(* IEC 61131-3 sources: STAR-PLC-Agent/results/raw/batch_fresh_20261114/PUB016/functional/attempt_0001, 1 file *)

(* ---- test_program.st ---- *)
PROGRAM PLC_PRG
VAR
 BenchStep : UDINT := 0;
 BenchCalls : UDINT := 0;
 BenchDone : BOOL := FALSE;
 BenchUut0 : FB_Task;
 BenchUut1 : FB_Task;
 BenchUut2 : FB_Task;
 BenchUut3 : FB_Task;
 BenchUut4 : FB_Task;
 BenchUut5 : FB_Task;
 BenchUut6 : FB_Task;
 BenchUut7 : FB_Task;
 TraceIn_processLength : ARRAY[0..159] OF USINT;
 TraceIn_sensor1 : ARRAY[0..159] OF BOOL;
 TraceIn_sensor2 : ARRAY[0..159] OF BOOL;
 TraceIn_sensor3 : ARRAY[0..159] OF BOOL;
 TraceIn_sensor4 : ARRAY[0..159] OF BOOL;
 TraceIn_sensor5 : ARRAY[0..159] OF BOOL;
 TraceIn_station1Start : ARRAY[0..159] OF BOOL;
 TraceIn_station2Complete : ARRAY[0..159] OF BOOL;
 TraceIn_station3Complete : ARRAY[0..159] OF BOOL;
 TraceIn_station4Complete : ARRAY[0..159] OF BOOL;
 TraceIn_processSequence_1 : ARRAY[0..159] OF USINT;
 TraceIn_processSequence_2 : ARRAY[0..159] OF USINT;
 TraceIn_processSequence_3 : ARRAY[0..159] OF USINT;
 TraceIn_processSequence_4 : ARRAY[0..159] OF USINT;
 TraceIn_processSequence_5 : ARRAY[0..159] OF USINT;
 TraceIn_processSequence_6 : ARRAY[0..159] OF USINT;
 TraceIn_processSequence_7 : ARRAY[0..159] OF USINT;
 TraceIn_processSequence_8 : ARRAY[0..159] OF USINT;
 TraceOut_conveyorLeft : ARRAY[0..159] OF BOOL;
 TraceOut_conveyorRight : ARRAY[0..159] OF BOOL;
END_VAR

IF NOT BenchDone THEN
 CASE BenchStep OF
 0:
   BenchUut0.processLength := USINT#3;
   BenchUut0.sensor1 := FALSE;
   BenchUut0.sensor2 := FALSE;
   BenchUut0.sensor3 := FALSE;
   BenchUut0.sensor4 := FALSE;
   BenchUut0.sensor5 := FALSE;
   BenchUut0.station1Start := FALSE;
   BenchUut0.station2Complete := FALSE;
   BenchUut0.station3Complete := FALSE;
   BenchUut0.station4Complete := FALSE;
   BenchUut0.processSequence[1] := USINT#4;
   BenchUut0.processSequence[2] := USINT#2;
   BenchUut0.processSequence[3] := USINT#5;
   BenchUut0.processSequence[4] := USINT#0;
   BenchUut0.processSequence[5] := USINT#0;
   BenchUut0.processSequence[6] := USINT#0;
   BenchUut0.processSequence[7] := USINT#0;
   BenchUut0.processSequence[8] := USINT#0;
   TraceIn_processLength[0] := BenchUut0.processLength;
   TraceIn_sensor1[0] := BenchUut0.sensor1;
   TraceIn_sensor2[0] := BenchUut0.sensor2;
   TraceIn_sensor3[0] := BenchUut0.sensor3;
   TraceIn_sensor4[0] := BenchUut0.sensor4;
   TraceIn_sensor5[0] := BenchUut0.sensor5;
   TraceIn_station1Start[0] := BenchUut0.station1Start;
   TraceIn_station2Complete[0] := BenchUut0.station2Complete;
   TraceIn_station3Complete[0] := BenchUut0.station3Complete;
   TraceIn_station4Complete[0] := BenchUut0.station4Complete;
   TraceIn_processSequence_1[0] := BenchUut0.processSequence[1];
   TraceIn_processSequence_2[0] := BenchUut0.processSequence[2];
   TraceIn_processSequence_3[0] := BenchUut0.processSequence[3];
   TraceIn_processSequence_4[0] := BenchUut0.processSequence[4];
   TraceIn_processSequence_5[0] := BenchUut0.processSequence[5];
   TraceIn_processSequence_6[0] := BenchUut0.processSequence[6];
   TraceIn_processSequence_7[0] := BenchUut0.processSequence[7];
   TraceIn_processSequence_8[0] := BenchUut0.processSequence[8];
   BenchUut0();
   TraceOut_conveyorLeft[0] := BenchUut0.conveyorLeft;
   TraceOut_conveyorRight[0] := BenchUut0.conveyorRight;
   BenchCalls := BenchCalls + 1;
 1:
   BenchUut0.processLength := USINT#3;
   BenchUut0.sensor1 := TRUE;
   BenchUut0.sensor2 := FALSE;
   BenchUut0.sensor3 := FALSE;
   BenchUut0.sensor4 := FALSE;
   BenchUut0.sensor5 := FALSE;
   BenchUut0.station1Start := TRUE;
   BenchUut0.station2Complete := FALSE;
   BenchUut0.station3Complete := FALSE;
   BenchUut0.station4Complete := FALSE;
   BenchUut0.processSequence[1] := USINT#4;
   BenchUut0.processSequence[2] := USINT#2;
   BenchUut0.processSequence[3] := USINT#5;
   BenchUut0.processSequence[4] := USINT#0;
   BenchUut0.processSequence[5] := USINT#0;
   BenchUut0.processSequence[6] := USINT#0;
   BenchUut0.processSequence[7] := USINT#0;
   BenchUut0.processSequence[8] := USINT#0;
   TraceIn_processLength[1] := BenchUut0.processLength;
   TraceIn_sensor1[1] := BenchUut0.sensor1;
   TraceIn_sensor2[1] := BenchUut0.sensor2;
   TraceIn_sensor3[1] := BenchUut0.sensor3;
   TraceIn_sensor4[1] := BenchUut0.sensor4;
   TraceIn_sensor5[1] := BenchUut0.sensor5;
   TraceIn_station1Start[1] := BenchUut0.station1Start;
   TraceIn_station2Complete[1] := BenchUut0.station2Complete;
   TraceIn_station3Complete[1] := BenchUut0.station3Complete;
   TraceIn_station4Complete[1] := BenchUut0.station4Complete;
   TraceIn_processSequence_1[1] := BenchUut0.processSequence[1];
   TraceIn_processSequence_2[1] := BenchUut0.processSequence[2];
   TraceIn_processSequence_3[1] := BenchUut0.processSequence[3];
   TraceIn_processSequence_4[1] := BenchUut0.processSequence[4];
   TraceIn_processSequence_5[1] := BenchUut0.processSequence[5];
   TraceIn_processSequence_6[1] := BenchUut0.processSequence[6];
   TraceIn_processSequence_7[1] := BenchUut0.processSequence[7];
   TraceIn_processSequence_8[1] := BenchUut0.processSequence[8];
   BenchUut0();
   TraceOut_conveyorLeft[1] := BenchUut0.conveyorLeft;
   TraceOut_conveyorRight[1] := BenchUut0.conveyorRight;
   BenchCalls := BenchCalls + 1;
 2:
   BenchUut0.processLength := USINT#3;
   BenchUut0.sensor1 := FALSE;
   BenchUut0.sensor2 := FALSE;
   BenchUut0.sensor3 := FALSE;
   BenchUut0.sensor4 := TRUE;
   BenchUut0.sensor5 := FALSE;
   BenchUut0.station1Start := FALSE;
   BenchUut0.station2Complete := FALSE;
   BenchUut0.station3Complete := FALSE;
   BenchUut0.station4Complete := FALSE;
   BenchUut0.processSequence[1] := USINT#4;
   BenchUut0.processSequence[2] := USINT#2;
   BenchUut0.processSequence[3] := USINT#5;
   BenchUut0.processSequence[4] := USINT#0;
   BenchUut0.processSequence[5] := USINT#0;
   BenchUut0.processSequence[6] := USINT#0;
   BenchUut0.processSequence[7] := USINT#0;
   BenchUut0.processSequence[8] := USINT#0;
   TraceIn_processLength[2] := BenchUut0.processLength;
   TraceIn_sensor1[2] := BenchUut0.sensor1;
   TraceIn_sensor2[2] := BenchUut0.sensor2;
   TraceIn_sensor3[2] := BenchUut0.sensor3;
   TraceIn_sensor4[2] := BenchUut0.sensor4;
   TraceIn_sensor5[2] := BenchUut0.sensor5;
   TraceIn_station1Start[2] := BenchUut0.station1Start;
   TraceIn_station2Complete[2] := BenchUut0.station2Complete;
   TraceIn_station3Complete[2] := BenchUut0.station3Complete;
   TraceIn_station4Complete[2] := BenchUut0.station4Complete;
   TraceIn_processSequence_1[2] := BenchUut0.processSequence[1];
   TraceIn_processSequence_2[2] := BenchUut0.processSequence[2];
   TraceIn_processSequence_3[2] := BenchUut0.processSequence[3];
   TraceIn_processSequence_4[2] := BenchUut0.processSequence[4];
   TraceIn_processSequence_5[2] := BenchUut0.processSequence[5];
   TraceIn_processSequence_6[2] := BenchUut0.processSequence[6];
   TraceIn_processSequence_7[2] := BenchUut0.processSequence[7];
   TraceIn_processSequence_8[2] := BenchUut0.processSequence[8];
   BenchUut0();
   TraceOut_conveyorLeft[2] := BenchUut0.conveyorLeft;
   TraceOut_conveyorRight[2] := BenchUut0.conveyorRight;
   BenchCalls := BenchCalls + 1;
 3:
   BenchUut0.processLength := USINT#3;
   BenchUut0.sensor1 := FALSE;
   BenchUut0.sensor2 := FALSE;
   BenchUut0.sensor3 := FALSE;
   BenchUut0.sensor4 := TRUE;
   BenchUut0.sensor5 := FALSE;
   BenchUut0.station1Start := FALSE;
   BenchUut0.station2Complete := FALSE;
   BenchUut0.station3Complete := TRUE;
   BenchUut0.station4Complete := FALSE;
   BenchUut0.processSequence[1] := USINT#4;
   BenchUut0.processSequence[2] := USINT#2;
   BenchUut0.processSequence[3] := USINT#5;
   BenchUut0.processSequence[4] := USINT#0;
   BenchUut0.processSequence[5] := USINT#0;
   BenchUut0.processSequence[6] := USINT#0;
   BenchUut0.processSequence[7] := USINT#0;
   BenchUut0.processSequence[8] := USINT#0;
   TraceIn_processLength[3] := BenchUut0.processLength;
   TraceIn_sensor1[3] := BenchUut0.sensor1;
   TraceIn_sensor2[3] := BenchUut0.sensor2;
   TraceIn_sensor3[3] := BenchUut0.sensor3;
   TraceIn_sensor4[3] := BenchUut0.sensor4;
   TraceIn_sensor5[3] := BenchUut0.sensor5;
   TraceIn_station1Start[3] := BenchUut0.station1Start;
   TraceIn_station2Complete[3] := BenchUut0.station2Complete;
   TraceIn_station3Complete[3] := BenchUut0.station3Complete;
   TraceIn_station4Complete[3] := BenchUut0.station4Complete;
   TraceIn_processSequence_1[3] := BenchUut0.processSequence[1];
   TraceIn_processSequence_2[3] := BenchUut0.processSequence[2];
   TraceIn_processSequence_3[3] := BenchUut0.processSequence[3];
   TraceIn_processSequence_4[3] := BenchUut0.processSequence[4];
   TraceIn_processSequence_5[3] := BenchUut0.processSequence[5];
   TraceIn_processSequence_6[3] := BenchUut0.processSequence[6];
   TraceIn_processSequence_7[3] := BenchUut0.processSequence[7];
   TraceIn_processSequence_8[3] := BenchUut0.processSequence[8];
   BenchUut0();
   TraceOut_conveyorLeft[3] := BenchUut0.conveyorLeft;
   TraceOut_conveyorRight[3] := BenchUut0.conveyorRight;
   BenchCalls := BenchCalls + 1;
 4:
   BenchUut0.processLength := USINT#3;
   BenchUut0.sensor1 := FALSE;
   BenchUut0.sensor2 := FALSE;
   BenchUut0.sensor3 := FALSE;
   BenchUut0.sensor4 := TRUE;
   BenchUut0.sensor5 := FALSE;
   BenchUut0.station1Start := FALSE;
   BenchUut0.station2Complete := FALSE;
   BenchUut0.station3Complete := FALSE;
   BenchUut0.station4Complete := TRUE;
   BenchUut0.processSequence[1] := USINT#4;
   BenchUut0.processSequence[2] := USINT#2;
   BenchUut0.processSequence[3] := USINT#5;
   BenchUut0.processSequence[4] := USINT#0;
   BenchUut0.processSequence[5] := USINT#0;
   BenchUut0.processSequence[6] := USINT#0;
   BenchUut0.processSequence[7] := USINT#0;
   BenchUut0.processSequence[8] := USINT#0;
   TraceIn_processLength[4] := BenchUut0.processLength;
   TraceIn_sensor1[4] := BenchUut0.sensor1;
   TraceIn_sensor2[4] := BenchUut0.sensor2;
   TraceIn_sensor3[4] := BenchUut0.sensor3;
   TraceIn_sensor4[4] := BenchUut0.sensor4;
   TraceIn_sensor5[4] := BenchUut0.sensor5;
   TraceIn_station1Start[4] := BenchUut0.station1Start;
   TraceIn_station2Complete[4] := BenchUut0.station2Complete;
   TraceIn_station3Complete[4] := BenchUut0.station3Complete;
   TraceIn_station4Complete[4] := BenchUut0.station4Complete;
   TraceIn_processSequence_1[4] := BenchUut0.processSequence[1];
   TraceIn_processSequence_2[4] := BenchUut0.processSequence[2];
   TraceIn_processSequence_3[4] := BenchUut0.processSequence[3];
   TraceIn_processSequence_4[4] := BenchUut0.processSequence[4];
   TraceIn_processSequence_5[4] := BenchUut0.processSequence[5];
   TraceIn_processSequence_6[4] := BenchUut0.processSequence[6];
   TraceIn_processSequence_7[4] := BenchUut0.processSequence[7];
   TraceIn_processSequence_8[4] := BenchUut0.processSequence[8];
   BenchUut0();
   TraceOut_conveyorLeft[4] := BenchUut0.conveyorLeft;
   TraceOut_conveyorRight[4] := BenchUut0.conveyorRight;
   BenchCalls := BenchCalls + 1;
 5:
   BenchUut0.processLength := USINT#3;
   BenchUut0.sensor1 := FALSE;
   BenchUut0.sensor2 := TRUE;
   BenchUut0.sensor3 := FALSE;
   BenchUut0.sensor4 := FALSE;
   BenchUut0.sensor5 := FALSE;
   BenchUut0.station1Start := FALSE;
   BenchUut0.station2Complete := FALSE;
   BenchUut0.station3Complete := FALSE;
   BenchUut0.station4Complete := FALSE;
   BenchUut0.processSequence[1] := USINT#4;
   BenchUut0.processSequence[2] := USINT#2;
   BenchUut0.processSequence[3] := USINT#5;
   BenchUut0.processSequence[4] := USINT#0;
   BenchUut0.processSequence[5] := USINT#0;
   BenchUut0.processSequence[6] := USINT#0;
   BenchUut0.processSequence[7] := USINT#0;
   BenchUut0.processSequence[8] := USINT#0;
   TraceIn_processLength[5] := BenchUut0.processLength;
   TraceIn_sensor1[5] := BenchUut0.sensor1;
   TraceIn_sensor2[5] := BenchUut0.sensor2;
   TraceIn_sensor3[5] := BenchUut0.sensor3;
   TraceIn_sensor4[5] := BenchUut0.sensor4;
   TraceIn_sensor5[5] := BenchUut0.sensor5;
   TraceIn_station1Start[5] := BenchUut0.station1Start;
   TraceIn_station2Complete[5] := BenchUut0.station2Complete;
   TraceIn_station3Complete[5] := BenchUut0.station3Complete;
   TraceIn_station4Complete[5] := BenchUut0.station4Complete;
   TraceIn_processSequence_1[5] := BenchUut0.processSequence[1];
   TraceIn_processSequence_2[5] := BenchUut0.processSequence[2];
   TraceIn_processSequence_3[5] := BenchUut0.processSequence[3];
   TraceIn_processSequence_4[5] := BenchUut0.processSequence[4];
   TraceIn_processSequence_5[5] := BenchUut0.processSequence[5];
   TraceIn_processSequence_6[5] := BenchUut0.processSequence[6];
   TraceIn_processSequence_7[5] := BenchUut0.processSequence[7];
   TraceIn_processSequence_8[5] := BenchUut0.processSequence[8];
   BenchUut0();
   TraceOut_conveyorLeft[5] := BenchUut0.conveyorLeft;
   TraceOut_conveyorRight[5] := BenchUut0.conveyorRight;
   BenchCalls := BenchCalls + 1;
 6:
   BenchUut0.processLength := USINT#3;
   BenchUut0.sensor1 := FALSE;
   BenchUut0.sensor2 := TRUE;
   BenchUut0.sensor3 := FALSE;
   BenchUut0.sensor4 := FALSE;
   BenchUut0.sensor5 := FALSE;
   BenchUut0.station1Start := FALSE;
   BenchUut0.station2Complete := TRUE;
   BenchUut0.station3Complete := FALSE;
   BenchUut0.station4Complete := FALSE;
   BenchUut0.processSequence[1] := USINT#4;
   BenchUut0.processSequence[2] := USINT#2;
   BenchUut0.processSequence[3] := USINT#5;
   BenchUut0.processSequence[4] := USINT#0;
   BenchUut0.processSequence[5] := USINT#0;
   BenchUut0.processSequence[6] := USINT#0;
   BenchUut0.processSequence[7] := USINT#0;
   BenchUut0.processSequence[8] := USINT#0;
   TraceIn_processLength[6] := BenchUut0.processLength;
   TraceIn_sensor1[6] := BenchUut0.sensor1;
   TraceIn_sensor2[6] := BenchUut0.sensor2;
   TraceIn_sensor3[6] := BenchUut0.sensor3;
   TraceIn_sensor4[6] := BenchUut0.sensor4;
   TraceIn_sensor5[6] := BenchUut0.sensor5;
   TraceIn_station1Start[6] := BenchUut0.station1Start;
   TraceIn_station2Complete[6] := BenchUut0.station2Complete;
   TraceIn_station3Complete[6] := BenchUut0.station3Complete;
   TraceIn_station4Complete[6] := BenchUut0.station4Complete;
   TraceIn_processSequence_1[6] := BenchUut0.processSequence[1];
   TraceIn_processSequence_2[6] := BenchUut0.processSequence[2];
   TraceIn_processSequence_3[6] := BenchUut0.processSequence[3];
   TraceIn_processSequence_4[6] := BenchUut0.processSequence[4];
   TraceIn_processSequence_5[6] := BenchUut0.processSequence[5];
   TraceIn_processSequence_6[6] := BenchUut0.processSequence[6];
   TraceIn_processSequence_7[6] := BenchUut0.processSequence[7];
   TraceIn_processSequence_8[6] := BenchUut0.processSequence[8];
   BenchUut0();
   TraceOut_conveyorLeft[6] := BenchUut0.conveyorLeft;
   TraceOut_conveyorRight[6] := BenchUut0.conveyorRight;
   BenchCalls := BenchCalls + 1;
 7:
   BenchUut0.processLength := USINT#3;
   BenchUut0.sensor1 := FALSE;
   BenchUut0.sensor2 := FALSE;
   BenchUut0.sensor3 := FALSE;
   BenchUut0.sensor4 := FALSE;
   BenchUut0.sensor5 := TRUE;
   BenchUut0.station1Start := FALSE;
   BenchUut0.station2Complete := FALSE;
   BenchUut0.station3Complete := FALSE;
   BenchUut0.station4Complete := FALSE;
   BenchUut0.processSequence[1] := USINT#4;
   BenchUut0.processSequence[2] := USINT#2;
   BenchUut0.processSequence[3] := USINT#5;
   BenchUut0.processSequence[4] := USINT#0;
   BenchUut0.processSequence[5] := USINT#0;
   BenchUut0.processSequence[6] := USINT#0;
   BenchUut0.processSequence[7] := USINT#0;
   BenchUut0.processSequence[8] := USINT#0;
   TraceIn_processLength[7] := BenchUut0.processLength;
   TraceIn_sensor1[7] := BenchUut0.sensor1;
   TraceIn_sensor2[7] := BenchUut0.sensor2;
   TraceIn_sensor3[7] := BenchUut0.sensor3;
   TraceIn_sensor4[7] := BenchUut0.sensor4;
   TraceIn_sensor5[7] := BenchUut0.sensor5;
   TraceIn_station1Start[7] := BenchUut0.station1Start;
   TraceIn_station2Complete[7] := BenchUut0.station2Complete;
   TraceIn_station3Complete[7] := BenchUut0.station3Complete;
   TraceIn_station4Complete[7] := BenchUut0.station4Complete;
   TraceIn_processSequence_1[7] := BenchUut0.processSequence[1];
   TraceIn_processSequence_2[7] := BenchUut0.processSequence[2];
   TraceIn_processSequence_3[7] := BenchUut0.processSequence[3];
   TraceIn_processSequence_4[7] := BenchUut0.processSequence[4];
   TraceIn_processSequence_5[7] := BenchUut0.processSequence[5];
   TraceIn_processSequence_6[7] := BenchUut0.processSequence[6];
   TraceIn_processSequence_7[7] := BenchUut0.processSequence[7];
   TraceIn_processSequence_8[7] := BenchUut0.processSequence[8];
   BenchUut0();
   TraceOut_conveyorLeft[7] := BenchUut0.conveyorLeft;
   TraceOut_conveyorRight[7] := BenchUut0.conveyorRight;
   BenchCalls := BenchCalls + 1;
 8:
   BenchUut1.processLength := USINT#1;
   BenchUut1.sensor1 := FALSE;
   BenchUut1.sensor2 := FALSE;
   BenchUut1.sensor3 := FALSE;
   BenchUut1.sensor4 := FALSE;
   BenchUut1.sensor5 := FALSE;
   BenchUut1.station1Start := FALSE;
   BenchUut1.station2Complete := FALSE;
   BenchUut1.station3Complete := FALSE;
   BenchUut1.station4Complete := FALSE;
   BenchUut1.processSequence[1] := USINT#5;
   BenchUut1.processSequence[2] := USINT#0;
   BenchUut1.processSequence[3] := USINT#0;
   BenchUut1.processSequence[4] := USINT#0;
   BenchUut1.processSequence[5] := USINT#0;
   BenchUut1.processSequence[6] := USINT#0;
   BenchUut1.processSequence[7] := USINT#0;
   BenchUut1.processSequence[8] := USINT#0;
   TraceIn_processLength[8] := BenchUut1.processLength;
   TraceIn_sensor1[8] := BenchUut1.sensor1;
   TraceIn_sensor2[8] := BenchUut1.sensor2;
   TraceIn_sensor3[8] := BenchUut1.sensor3;
   TraceIn_sensor4[8] := BenchUut1.sensor4;
   TraceIn_sensor5[8] := BenchUut1.sensor5;
   TraceIn_station1Start[8] := BenchUut1.station1Start;
   TraceIn_station2Complete[8] := BenchUut1.station2Complete;
   TraceIn_station3Complete[8] := BenchUut1.station3Complete;
   TraceIn_station4Complete[8] := BenchUut1.station4Complete;
   TraceIn_processSequence_1[8] := BenchUut1.processSequence[1];
   TraceIn_processSequence_2[8] := BenchUut1.processSequence[2];
   TraceIn_processSequence_3[8] := BenchUut1.processSequence[3];
   TraceIn_processSequence_4[8] := BenchUut1.processSequence[4];
   TraceIn_processSequence_5[8] := BenchUut1.processSequence[5];
   TraceIn_processSequence_6[8] := BenchUut1.processSequence[6];
   TraceIn_processSequence_7[8] := BenchUut1.processSequence[7];
   TraceIn_processSequence_8[8] := BenchUut1.processSequence[8];
   BenchUut1();
   TraceOut_conveyorLeft[8] := BenchUut1.conveyorLeft;
   TraceOut_conveyorRight[8] := BenchUut1.conveyorRight;
   BenchCalls := BenchCalls + 1;
 9:
   BenchUut1.processLength := USINT#1;
   BenchUut1.sensor1 := TRUE;
   BenchUut1.sensor2 := FALSE;
   BenchUut1.sensor3 := FALSE;
   BenchUut1.sensor4 := FALSE;
   BenchUut1.sensor5 := FALSE;
   BenchUut1.station1Start := TRUE;
   BenchUut1.station2Complete := FALSE;
   BenchUut1.station3Complete := FALSE;
   BenchUut1.station4Complete := FALSE;
   BenchUut1.processSequence[1] := USINT#5;
   BenchUut1.processSequence[2] := USINT#0;
   BenchUut1.processSequence[3] := USINT#0;
   BenchUut1.processSequence[4] := USINT#0;
   BenchUut1.processSequence[5] := USINT#0;
   BenchUut1.processSequence[6] := USINT#0;
   BenchUut1.processSequence[7] := USINT#0;
   BenchUut1.processSequence[8] := USINT#0;
   TraceIn_processLength[9] := BenchUut1.processLength;
   TraceIn_sensor1[9] := BenchUut1.sensor1;
   TraceIn_sensor2[9] := BenchUut1.sensor2;
   TraceIn_sensor3[9] := BenchUut1.sensor3;
   TraceIn_sensor4[9] := BenchUut1.sensor4;
   TraceIn_sensor5[9] := BenchUut1.sensor5;
   TraceIn_station1Start[9] := BenchUut1.station1Start;
   TraceIn_station2Complete[9] := BenchUut1.station2Complete;
   TraceIn_station3Complete[9] := BenchUut1.station3Complete;
   TraceIn_station4Complete[9] := BenchUut1.station4Complete;
   TraceIn_processSequence_1[9] := BenchUut1.processSequence[1];
   TraceIn_processSequence_2[9] := BenchUut1.processSequence[2];
   TraceIn_processSequence_3[9] := BenchUut1.processSequence[3];
   TraceIn_processSequence_4[9] := BenchUut1.processSequence[4];
   TraceIn_processSequence_5[9] := BenchUut1.processSequence[5];
   TraceIn_processSequence_6[9] := BenchUut1.processSequence[6];
   TraceIn_processSequence_7[9] := BenchUut1.processSequence[7];
   TraceIn_processSequence_8[9] := BenchUut1.processSequence[8];
   BenchUut1();
   TraceOut_conveyorLeft[9] := BenchUut1.conveyorLeft;
   TraceOut_conveyorRight[9] := BenchUut1.conveyorRight;
   BenchCalls := BenchCalls + 1;
 10:
   BenchUut1.processLength := USINT#1;
   BenchUut1.sensor1 := FALSE;
   BenchUut1.sensor2 := FALSE;
   BenchUut1.sensor3 := FALSE;
   BenchUut1.sensor4 := FALSE;
   BenchUut1.sensor5 := TRUE;
   BenchUut1.station1Start := FALSE;
   BenchUut1.station2Complete := FALSE;
   BenchUut1.station3Complete := FALSE;
   BenchUut1.station4Complete := FALSE;
   BenchUut1.processSequence[1] := USINT#5;
   BenchUut1.processSequence[2] := USINT#0;
   BenchUut1.processSequence[3] := USINT#0;
   BenchUut1.processSequence[4] := USINT#0;
   BenchUut1.processSequence[5] := USINT#0;
   BenchUut1.processSequence[6] := USINT#0;
   BenchUut1.processSequence[7] := USINT#0;
   BenchUut1.processSequence[8] := USINT#0;
   TraceIn_processLength[10] := BenchUut1.processLength;
   TraceIn_sensor1[10] := BenchUut1.sensor1;
   TraceIn_sensor2[10] := BenchUut1.sensor2;
   TraceIn_sensor3[10] := BenchUut1.sensor3;
   TraceIn_sensor4[10] := BenchUut1.sensor4;
   TraceIn_sensor5[10] := BenchUut1.sensor5;
   TraceIn_station1Start[10] := BenchUut1.station1Start;
   TraceIn_station2Complete[10] := BenchUut1.station2Complete;
   TraceIn_station3Complete[10] := BenchUut1.station3Complete;
   TraceIn_station4Complete[10] := BenchUut1.station4Complete;
   TraceIn_processSequence_1[10] := BenchUut1.processSequence[1];
   TraceIn_processSequence_2[10] := BenchUut1.processSequence[2];
   TraceIn_processSequence_3[10] := BenchUut1.processSequence[3];
   TraceIn_processSequence_4[10] := BenchUut1.processSequence[4];
   TraceIn_processSequence_5[10] := BenchUut1.processSequence[5];
   TraceIn_processSequence_6[10] := BenchUut1.processSequence[6];
   TraceIn_processSequence_7[10] := BenchUut1.processSequence[7];
   TraceIn_processSequence_8[10] := BenchUut1.processSequence[8];
   BenchUut1();
   TraceOut_conveyorLeft[10] := BenchUut1.conveyorLeft;
   TraceOut_conveyorRight[10] := BenchUut1.conveyorRight;
   BenchCalls := BenchCalls + 1;
 11:
   BenchUut2.processLength := USINT#3;
   BenchUut2.sensor1 := FALSE;
   BenchUut2.sensor2 := FALSE;
   BenchUut2.sensor3 := FALSE;
   BenchUut2.sensor4 := FALSE;
   BenchUut2.sensor5 := FALSE;
   BenchUut2.station1Start := FALSE;
   BenchUut2.station2Complete := FALSE;
   BenchUut2.station3Complete := FALSE;
   BenchUut2.station4Complete := FALSE;
   BenchUut2.processSequence[1] := USINT#2;
   BenchUut2.processSequence[2] := USINT#2;
   BenchUut2.processSequence[3] := USINT#5;
   BenchUut2.processSequence[4] := USINT#0;
   BenchUut2.processSequence[5] := USINT#0;
   BenchUut2.processSequence[6] := USINT#0;
   BenchUut2.processSequence[7] := USINT#0;
   BenchUut2.processSequence[8] := USINT#0;
   TraceIn_processLength[11] := BenchUut2.processLength;
   TraceIn_sensor1[11] := BenchUut2.sensor1;
   TraceIn_sensor2[11] := BenchUut2.sensor2;
   TraceIn_sensor3[11] := BenchUut2.sensor3;
   TraceIn_sensor4[11] := BenchUut2.sensor4;
   TraceIn_sensor5[11] := BenchUut2.sensor5;
   TraceIn_station1Start[11] := BenchUut2.station1Start;
   TraceIn_station2Complete[11] := BenchUut2.station2Complete;
   TraceIn_station3Complete[11] := BenchUut2.station3Complete;
   TraceIn_station4Complete[11] := BenchUut2.station4Complete;
   TraceIn_processSequence_1[11] := BenchUut2.processSequence[1];
   TraceIn_processSequence_2[11] := BenchUut2.processSequence[2];
   TraceIn_processSequence_3[11] := BenchUut2.processSequence[3];
   TraceIn_processSequence_4[11] := BenchUut2.processSequence[4];
   TraceIn_processSequence_5[11] := BenchUut2.processSequence[5];
   TraceIn_processSequence_6[11] := BenchUut2.processSequence[6];
   TraceIn_processSequence_7[11] := BenchUut2.processSequence[7];
   TraceIn_processSequence_8[11] := BenchUut2.processSequence[8];
   BenchUut2();
   TraceOut_conveyorLeft[11] := BenchUut2.conveyorLeft;
   TraceOut_conveyorRight[11] := BenchUut2.conveyorRight;
   BenchCalls := BenchCalls + 1;
 12:
   BenchUut2.processLength := USINT#3;
   BenchUut2.sensor1 := TRUE;
   BenchUut2.sensor2 := FALSE;
   BenchUut2.sensor3 := FALSE;
   BenchUut2.sensor4 := FALSE;
   BenchUut2.sensor5 := FALSE;
   BenchUut2.station1Start := TRUE;
   BenchUut2.station2Complete := FALSE;
   BenchUut2.station3Complete := FALSE;
   BenchUut2.station4Complete := FALSE;
   BenchUut2.processSequence[1] := USINT#2;
   BenchUut2.processSequence[2] := USINT#2;
   BenchUut2.processSequence[3] := USINT#5;
   BenchUut2.processSequence[4] := USINT#0;
   BenchUut2.processSequence[5] := USINT#0;
   BenchUut2.processSequence[6] := USINT#0;
   BenchUut2.processSequence[7] := USINT#0;
   BenchUut2.processSequence[8] := USINT#0;
   TraceIn_processLength[12] := BenchUut2.processLength;
   TraceIn_sensor1[12] := BenchUut2.sensor1;
   TraceIn_sensor2[12] := BenchUut2.sensor2;
   TraceIn_sensor3[12] := BenchUut2.sensor3;
   TraceIn_sensor4[12] := BenchUut2.sensor4;
   TraceIn_sensor5[12] := BenchUut2.sensor5;
   TraceIn_station1Start[12] := BenchUut2.station1Start;
   TraceIn_station2Complete[12] := BenchUut2.station2Complete;
   TraceIn_station3Complete[12] := BenchUut2.station3Complete;
   TraceIn_station4Complete[12] := BenchUut2.station4Complete;
   TraceIn_processSequence_1[12] := BenchUut2.processSequence[1];
   TraceIn_processSequence_2[12] := BenchUut2.processSequence[2];
   TraceIn_processSequence_3[12] := BenchUut2.processSequence[3];
   TraceIn_processSequence_4[12] := BenchUut2.processSequence[4];
   TraceIn_processSequence_5[12] := BenchUut2.processSequence[5];
   TraceIn_processSequence_6[12] := BenchUut2.processSequence[6];
   TraceIn_processSequence_7[12] := BenchUut2.processSequence[7];
   TraceIn_processSequence_8[12] := BenchUut2.processSequence[8];
   BenchUut2();
   TraceOut_conveyorLeft[12] := BenchUut2.conveyorLeft;
   TraceOut_conveyorRight[12] := BenchUut2.conveyorRight;
   BenchCalls := BenchCalls + 1;
 13:
   BenchUut2.processLength := USINT#3;
   BenchUut2.sensor1 := FALSE;
   BenchUut2.sensor2 := TRUE;
   BenchUut2.sensor3 := FALSE;
   BenchUut2.sensor4 := FALSE;
   BenchUut2.sensor5 := FALSE;
   BenchUut2.station1Start := FALSE;
   BenchUut2.station2Complete := FALSE;
   BenchUut2.station3Complete := FALSE;
   BenchUut2.station4Complete := FALSE;
   BenchUut2.processSequence[1] := USINT#2;
   BenchUut2.processSequence[2] := USINT#2;
   BenchUut2.processSequence[3] := USINT#5;
   BenchUut2.processSequence[4] := USINT#0;
   BenchUut2.processSequence[5] := USINT#0;
   BenchUut2.processSequence[6] := USINT#0;
   BenchUut2.processSequence[7] := USINT#0;
   BenchUut2.processSequence[8] := USINT#0;
   TraceIn_processLength[13] := BenchUut2.processLength;
   TraceIn_sensor1[13] := BenchUut2.sensor1;
   TraceIn_sensor2[13] := BenchUut2.sensor2;
   TraceIn_sensor3[13] := BenchUut2.sensor3;
   TraceIn_sensor4[13] := BenchUut2.sensor4;
   TraceIn_sensor5[13] := BenchUut2.sensor5;
   TraceIn_station1Start[13] := BenchUut2.station1Start;
   TraceIn_station2Complete[13] := BenchUut2.station2Complete;
   TraceIn_station3Complete[13] := BenchUut2.station3Complete;
   TraceIn_station4Complete[13] := BenchUut2.station4Complete;
   TraceIn_processSequence_1[13] := BenchUut2.processSequence[1];
   TraceIn_processSequence_2[13] := BenchUut2.processSequence[2];
   TraceIn_processSequence_3[13] := BenchUut2.processSequence[3];
   TraceIn_processSequence_4[13] := BenchUut2.processSequence[4];
   TraceIn_processSequence_5[13] := BenchUut2.processSequence[5];
   TraceIn_processSequence_6[13] := BenchUut2.processSequence[6];
   TraceIn_processSequence_7[13] := BenchUut2.processSequence[7];
   TraceIn_processSequence_8[13] := BenchUut2.processSequence[8];
   BenchUut2();
   TraceOut_conveyorLeft[13] := BenchUut2.conveyorLeft;
   TraceOut_conveyorRight[13] := BenchUut2.conveyorRight;
   BenchCalls := BenchCalls + 1;
 14:
   BenchUut2.processLength := USINT#3;
   BenchUut2.sensor1 := FALSE;
   BenchUut2.sensor2 := TRUE;
   BenchUut2.sensor3 := FALSE;
   BenchUut2.sensor4 := FALSE;
   BenchUut2.sensor5 := FALSE;
   BenchUut2.station1Start := FALSE;
   BenchUut2.station2Complete := TRUE;
   BenchUut2.station3Complete := FALSE;
   BenchUut2.station4Complete := FALSE;
   BenchUut2.processSequence[1] := USINT#2;
   BenchUut2.processSequence[2] := USINT#2;
   BenchUut2.processSequence[3] := USINT#5;
   BenchUut2.processSequence[4] := USINT#0;
   BenchUut2.processSequence[5] := USINT#0;
   BenchUut2.processSequence[6] := USINT#0;
   BenchUut2.processSequence[7] := USINT#0;
   BenchUut2.processSequence[8] := USINT#0;
   TraceIn_processLength[14] := BenchUut2.processLength;
   TraceIn_sensor1[14] := BenchUut2.sensor1;
   TraceIn_sensor2[14] := BenchUut2.sensor2;
   TraceIn_sensor3[14] := BenchUut2.sensor3;
   TraceIn_sensor4[14] := BenchUut2.sensor4;
   TraceIn_sensor5[14] := BenchUut2.sensor5;
   TraceIn_station1Start[14] := BenchUut2.station1Start;
   TraceIn_station2Complete[14] := BenchUut2.station2Complete;
   TraceIn_station3Complete[14] := BenchUut2.station3Complete;
   TraceIn_station4Complete[14] := BenchUut2.station4Complete;
   TraceIn_processSequence_1[14] := BenchUut2.processSequence[1];
   TraceIn_processSequence_2[14] := BenchUut2.processSequence[2];
   TraceIn_processSequence_3[14] := BenchUut2.processSequence[3];
   TraceIn_processSequence_4[14] := BenchUut2.processSequence[4];
   TraceIn_processSequence_5[14] := BenchUut2.processSequence[5];
   TraceIn_processSequence_6[14] := BenchUut2.processSequence[6];
   TraceIn_processSequence_7[14] := BenchUut2.processSequence[7];
   TraceIn_processSequence_8[14] := BenchUut2.processSequence[8];
   BenchUut2();
   TraceOut_conveyorLeft[14] := BenchUut2.conveyorLeft;
   TraceOut_conveyorRight[14] := BenchUut2.conveyorRight;
   BenchCalls := BenchCalls + 1;
 15:
   BenchUut2.processLength := USINT#3;
   BenchUut2.sensor1 := FALSE;
   BenchUut2.sensor2 := TRUE;
   BenchUut2.sensor3 := FALSE;
   BenchUut2.sensor4 := FALSE;
   BenchUut2.sensor5 := FALSE;
   BenchUut2.station1Start := FALSE;
   BenchUut2.station2Complete := TRUE;
   BenchUut2.station3Complete := FALSE;
   BenchUut2.station4Complete := FALSE;
   BenchUut2.processSequence[1] := USINT#2;
   BenchUut2.processSequence[2] := USINT#2;
   BenchUut2.processSequence[3] := USINT#5;
   BenchUut2.processSequence[4] := USINT#0;
   BenchUut2.processSequence[5] := USINT#0;
   BenchUut2.processSequence[6] := USINT#0;
   BenchUut2.processSequence[7] := USINT#0;
   BenchUut2.processSequence[8] := USINT#0;
   TraceIn_processLength[15] := BenchUut2.processLength;
   TraceIn_sensor1[15] := BenchUut2.sensor1;
   TraceIn_sensor2[15] := BenchUut2.sensor2;
   TraceIn_sensor3[15] := BenchUut2.sensor3;
   TraceIn_sensor4[15] := BenchUut2.sensor4;
   TraceIn_sensor5[15] := BenchUut2.sensor5;
   TraceIn_station1Start[15] := BenchUut2.station1Start;
   TraceIn_station2Complete[15] := BenchUut2.station2Complete;
   TraceIn_station3Complete[15] := BenchUut2.station3Complete;
   TraceIn_station4Complete[15] := BenchUut2.station4Complete;
   TraceIn_processSequence_1[15] := BenchUut2.processSequence[1];
   TraceIn_processSequence_2[15] := BenchUut2.processSequence[2];
   TraceIn_processSequence_3[15] := BenchUut2.processSequence[3];
   TraceIn_processSequence_4[15] := BenchUut2.processSequence[4];
   TraceIn_processSequence_5[15] := BenchUut2.processSequence[5];
   TraceIn_processSequence_6[15] := BenchUut2.processSequence[6];
   TraceIn_processSequence_7[15] := BenchUut2.processSequence[7];
   TraceIn_processSequence_8[15] := BenchUut2.processSequence[8];
   BenchUut2();
   TraceOut_conveyorLeft[15] := BenchUut2.conveyorLeft;
   TraceOut_conveyorRight[15] := BenchUut2.conveyorRight;
   BenchCalls := BenchCalls + 1;
 16:
   BenchUut2.processLength := USINT#3;
   BenchUut2.sensor1 := FALSE;
   BenchUut2.sensor2 := TRUE;
   BenchUut2.sensor3 := FALSE;
   BenchUut2.sensor4 := FALSE;
   BenchUut2.sensor5 := FALSE;
   BenchUut2.station1Start := FALSE;
   BenchUut2.station2Complete := FALSE;
   BenchUut2.station3Complete := FALSE;
   BenchUut2.station4Complete := FALSE;
   BenchUut2.processSequence[1] := USINT#2;
   BenchUut2.processSequence[2] := USINT#2;
   BenchUut2.processSequence[3] := USINT#5;
   BenchUut2.processSequence[4] := USINT#0;
   BenchUut2.processSequence[5] := USINT#0;
   BenchUut2.processSequence[6] := USINT#0;
   BenchUut2.processSequence[7] := USINT#0;
   BenchUut2.processSequence[8] := USINT#0;
   TraceIn_processLength[16] := BenchUut2.processLength;
   TraceIn_sensor1[16] := BenchUut2.sensor1;
   TraceIn_sensor2[16] := BenchUut2.sensor2;
   TraceIn_sensor3[16] := BenchUut2.sensor3;
   TraceIn_sensor4[16] := BenchUut2.sensor4;
   TraceIn_sensor5[16] := BenchUut2.sensor5;
   TraceIn_station1Start[16] := BenchUut2.station1Start;
   TraceIn_station2Complete[16] := BenchUut2.station2Complete;
   TraceIn_station3Complete[16] := BenchUut2.station3Complete;
   TraceIn_station4Complete[16] := BenchUut2.station4Complete;
   TraceIn_processSequence_1[16] := BenchUut2.processSequence[1];
   TraceIn_processSequence_2[16] := BenchUut2.processSequence[2];
   TraceIn_processSequence_3[16] := BenchUut2.processSequence[3];
   TraceIn_processSequence_4[16] := BenchUut2.processSequence[4];
   TraceIn_processSequence_5[16] := BenchUut2.processSequence[5];
   TraceIn_processSequence_6[16] := BenchUut2.processSequence[6];
   TraceIn_processSequence_7[16] := BenchUut2.processSequence[7];
   TraceIn_processSequence_8[16] := BenchUut2.processSequence[8];
   BenchUut2();
   TraceOut_conveyorLeft[16] := BenchUut2.conveyorLeft;
   TraceOut_conveyorRight[16] := BenchUut2.conveyorRight;
   BenchCalls := BenchCalls + 1;
 17:
   BenchUut2.processLength := USINT#3;
   BenchUut2.sensor1 := FALSE;
   BenchUut2.sensor2 := TRUE;
   BenchUut2.sensor3 := FALSE;
   BenchUut2.sensor4 := FALSE;
   BenchUut2.sensor5 := FALSE;
   BenchUut2.station1Start := FALSE;
   BenchUut2.station2Complete := TRUE;
   BenchUut2.station3Complete := FALSE;
   BenchUut2.station4Complete := FALSE;
   BenchUut2.processSequence[1] := USINT#2;
   BenchUut2.processSequence[2] := USINT#2;
   BenchUut2.processSequence[3] := USINT#5;
   BenchUut2.processSequence[4] := USINT#0;
   BenchUut2.processSequence[5] := USINT#0;
   BenchUut2.processSequence[6] := USINT#0;
   BenchUut2.processSequence[7] := USINT#0;
   BenchUut2.processSequence[8] := USINT#0;
   TraceIn_processLength[17] := BenchUut2.processLength;
   TraceIn_sensor1[17] := BenchUut2.sensor1;
   TraceIn_sensor2[17] := BenchUut2.sensor2;
   TraceIn_sensor3[17] := BenchUut2.sensor3;
   TraceIn_sensor4[17] := BenchUut2.sensor4;
   TraceIn_sensor5[17] := BenchUut2.sensor5;
   TraceIn_station1Start[17] := BenchUut2.station1Start;
   TraceIn_station2Complete[17] := BenchUut2.station2Complete;
   TraceIn_station3Complete[17] := BenchUut2.station3Complete;
   TraceIn_station4Complete[17] := BenchUut2.station4Complete;
   TraceIn_processSequence_1[17] := BenchUut2.processSequence[1];
   TraceIn_processSequence_2[17] := BenchUut2.processSequence[2];
   TraceIn_processSequence_3[17] := BenchUut2.processSequence[3];
   TraceIn_processSequence_4[17] := BenchUut2.processSequence[4];
   TraceIn_processSequence_5[17] := BenchUut2.processSequence[5];
   TraceIn_processSequence_6[17] := BenchUut2.processSequence[6];
   TraceIn_processSequence_7[17] := BenchUut2.processSequence[7];
   TraceIn_processSequence_8[17] := BenchUut2.processSequence[8];
   BenchUut2();
   TraceOut_conveyorLeft[17] := BenchUut2.conveyorLeft;
   TraceOut_conveyorRight[17] := BenchUut2.conveyorRight;
   BenchCalls := BenchCalls + 1;
 18:
   BenchUut3.processLength := USINT#3;
   BenchUut3.sensor1 := TRUE;
   BenchUut3.sensor2 := FALSE;
   BenchUut3.sensor3 := FALSE;
   BenchUut3.sensor4 := FALSE;
   BenchUut3.sensor5 := FALSE;
   BenchUut3.station1Start := TRUE;
   BenchUut3.station2Complete := FALSE;
   BenchUut3.station3Complete := FALSE;
   BenchUut3.station4Complete := FALSE;
   BenchUut3.processSequence[1] := USINT#2;
   BenchUut3.processSequence[2] := USINT#2;
   BenchUut3.processSequence[3] := USINT#5;
   BenchUut3.processSequence[4] := USINT#0;
   BenchUut3.processSequence[5] := USINT#0;
   BenchUut3.processSequence[6] := USINT#0;
   BenchUut3.processSequence[7] := USINT#0;
   BenchUut3.processSequence[8] := USINT#0;
   TraceIn_processLength[18] := BenchUut3.processLength;
   TraceIn_sensor1[18] := BenchUut3.sensor1;
   TraceIn_sensor2[18] := BenchUut3.sensor2;
   TraceIn_sensor3[18] := BenchUut3.sensor3;
   TraceIn_sensor4[18] := BenchUut3.sensor4;
   TraceIn_sensor5[18] := BenchUut3.sensor5;
   TraceIn_station1Start[18] := BenchUut3.station1Start;
   TraceIn_station2Complete[18] := BenchUut3.station2Complete;
   TraceIn_station3Complete[18] := BenchUut3.station3Complete;
   TraceIn_station4Complete[18] := BenchUut3.station4Complete;
   TraceIn_processSequence_1[18] := BenchUut3.processSequence[1];
   TraceIn_processSequence_2[18] := BenchUut3.processSequence[2];
   TraceIn_processSequence_3[18] := BenchUut3.processSequence[3];
   TraceIn_processSequence_4[18] := BenchUut3.processSequence[4];
   TraceIn_processSequence_5[18] := BenchUut3.processSequence[5];
   TraceIn_processSequence_6[18] := BenchUut3.processSequence[6];
   TraceIn_processSequence_7[18] := BenchUut3.processSequence[7];
   TraceIn_processSequence_8[18] := BenchUut3.processSequence[8];
   BenchUut3();
   TraceOut_conveyorLeft[18] := BenchUut3.conveyorLeft;
   TraceOut_conveyorRight[18] := BenchUut3.conveyorRight;
   BenchCalls := BenchCalls + 1;
 19:
   BenchUut3.processLength := USINT#3;
   BenchUut3.sensor1 := FALSE;
   BenchUut3.sensor2 := TRUE;
   BenchUut3.sensor3 := FALSE;
   BenchUut3.sensor4 := FALSE;
   BenchUut3.sensor5 := FALSE;
   BenchUut3.station1Start := FALSE;
   BenchUut3.station2Complete := TRUE;
   BenchUut3.station3Complete := FALSE;
   BenchUut3.station4Complete := FALSE;
   BenchUut3.processSequence[1] := USINT#2;
   BenchUut3.processSequence[2] := USINT#2;
   BenchUut3.processSequence[3] := USINT#5;
   BenchUut3.processSequence[4] := USINT#0;
   BenchUut3.processSequence[5] := USINT#0;
   BenchUut3.processSequence[6] := USINT#0;
   BenchUut3.processSequence[7] := USINT#0;
   BenchUut3.processSequence[8] := USINT#0;
   TraceIn_processLength[19] := BenchUut3.processLength;
   TraceIn_sensor1[19] := BenchUut3.sensor1;
   TraceIn_sensor2[19] := BenchUut3.sensor2;
   TraceIn_sensor3[19] := BenchUut3.sensor3;
   TraceIn_sensor4[19] := BenchUut3.sensor4;
   TraceIn_sensor5[19] := BenchUut3.sensor5;
   TraceIn_station1Start[19] := BenchUut3.station1Start;
   TraceIn_station2Complete[19] := BenchUut3.station2Complete;
   TraceIn_station3Complete[19] := BenchUut3.station3Complete;
   TraceIn_station4Complete[19] := BenchUut3.station4Complete;
   TraceIn_processSequence_1[19] := BenchUut3.processSequence[1];
   TraceIn_processSequence_2[19] := BenchUut3.processSequence[2];
   TraceIn_processSequence_3[19] := BenchUut3.processSequence[3];
   TraceIn_processSequence_4[19] := BenchUut3.processSequence[4];
   TraceIn_processSequence_5[19] := BenchUut3.processSequence[5];
   TraceIn_processSequence_6[19] := BenchUut3.processSequence[6];
   TraceIn_processSequence_7[19] := BenchUut3.processSequence[7];
   TraceIn_processSequence_8[19] := BenchUut3.processSequence[8];
   BenchUut3();
   TraceOut_conveyorLeft[19] := BenchUut3.conveyorLeft;
   TraceOut_conveyorRight[19] := BenchUut3.conveyorRight;
   BenchCalls := BenchCalls + 1;
 20:
   BenchUut3.processLength := USINT#3;
   BenchUut3.sensor1 := FALSE;
   BenchUut3.sensor2 := TRUE;
   BenchUut3.sensor3 := FALSE;
   BenchUut3.sensor4 := FALSE;
   BenchUut3.sensor5 := FALSE;
   BenchUut3.station1Start := FALSE;
   BenchUut3.station2Complete := TRUE;
   BenchUut3.station3Complete := FALSE;
   BenchUut3.station4Complete := FALSE;
   BenchUut3.processSequence[1] := USINT#2;
   BenchUut3.processSequence[2] := USINT#2;
   BenchUut3.processSequence[3] := USINT#5;
   BenchUut3.processSequence[4] := USINT#0;
   BenchUut3.processSequence[5] := USINT#0;
   BenchUut3.processSequence[6] := USINT#0;
   BenchUut3.processSequence[7] := USINT#0;
   BenchUut3.processSequence[8] := USINT#0;
   TraceIn_processLength[20] := BenchUut3.processLength;
   TraceIn_sensor1[20] := BenchUut3.sensor1;
   TraceIn_sensor2[20] := BenchUut3.sensor2;
   TraceIn_sensor3[20] := BenchUut3.sensor3;
   TraceIn_sensor4[20] := BenchUut3.sensor4;
   TraceIn_sensor5[20] := BenchUut3.sensor5;
   TraceIn_station1Start[20] := BenchUut3.station1Start;
   TraceIn_station2Complete[20] := BenchUut3.station2Complete;
   TraceIn_station3Complete[20] := BenchUut3.station3Complete;
   TraceIn_station4Complete[20] := BenchUut3.station4Complete;
   TraceIn_processSequence_1[20] := BenchUut3.processSequence[1];
   TraceIn_processSequence_2[20] := BenchUut3.processSequence[2];
   TraceIn_processSequence_3[20] := BenchUut3.processSequence[3];
   TraceIn_processSequence_4[20] := BenchUut3.processSequence[4];
   TraceIn_processSequence_5[20] := BenchUut3.processSequence[5];
   TraceIn_processSequence_6[20] := BenchUut3.processSequence[6];
   TraceIn_processSequence_7[20] := BenchUut3.processSequence[7];
   TraceIn_processSequence_8[20] := BenchUut3.processSequence[8];
   BenchUut3();
   TraceOut_conveyorLeft[20] := BenchUut3.conveyorLeft;
   TraceOut_conveyorRight[20] := BenchUut3.conveyorRight;
   BenchCalls := BenchCalls + 1;
 21:
   BenchUut3.processLength := USINT#3;
   BenchUut3.sensor1 := FALSE;
   BenchUut3.sensor2 := TRUE;
   BenchUut3.sensor3 := FALSE;
   BenchUut3.sensor4 := FALSE;
   BenchUut3.sensor5 := FALSE;
   BenchUut3.station1Start := FALSE;
   BenchUut3.station2Complete := FALSE;
   BenchUut3.station3Complete := FALSE;
   BenchUut3.station4Complete := FALSE;
   BenchUut3.processSequence[1] := USINT#2;
   BenchUut3.processSequence[2] := USINT#2;
   BenchUut3.processSequence[3] := USINT#5;
   BenchUut3.processSequence[4] := USINT#0;
   BenchUut3.processSequence[5] := USINT#0;
   BenchUut3.processSequence[6] := USINT#0;
   BenchUut3.processSequence[7] := USINT#0;
   BenchUut3.processSequence[8] := USINT#0;
   TraceIn_processLength[21] := BenchUut3.processLength;
   TraceIn_sensor1[21] := BenchUut3.sensor1;
   TraceIn_sensor2[21] := BenchUut3.sensor2;
   TraceIn_sensor3[21] := BenchUut3.sensor3;
   TraceIn_sensor4[21] := BenchUut3.sensor4;
   TraceIn_sensor5[21] := BenchUut3.sensor5;
   TraceIn_station1Start[21] := BenchUut3.station1Start;
   TraceIn_station2Complete[21] := BenchUut3.station2Complete;
   TraceIn_station3Complete[21] := BenchUut3.station3Complete;
   TraceIn_station4Complete[21] := BenchUut3.station4Complete;
   TraceIn_processSequence_1[21] := BenchUut3.processSequence[1];
   TraceIn_processSequence_2[21] := BenchUut3.processSequence[2];
   TraceIn_processSequence_3[21] := BenchUut3.processSequence[3];
   TraceIn_processSequence_4[21] := BenchUut3.processSequence[4];
   TraceIn_processSequence_5[21] := BenchUut3.processSequence[5];
   TraceIn_processSequence_6[21] := BenchUut3.processSequence[6];
   TraceIn_processSequence_7[21] := BenchUut3.processSequence[7];
   TraceIn_processSequence_8[21] := BenchUut3.processSequence[8];
   BenchUut3();
   TraceOut_conveyorLeft[21] := BenchUut3.conveyorLeft;
   TraceOut_conveyorRight[21] := BenchUut3.conveyorRight;
   BenchCalls := BenchCalls + 1;
 22:
   BenchUut3.processLength := USINT#3;
   BenchUut3.sensor1 := FALSE;
   BenchUut3.sensor2 := TRUE;
   BenchUut3.sensor3 := FALSE;
   BenchUut3.sensor4 := FALSE;
   BenchUut3.sensor5 := FALSE;
   BenchUut3.station1Start := FALSE;
   BenchUut3.station2Complete := TRUE;
   BenchUut3.station3Complete := FALSE;
   BenchUut3.station4Complete := FALSE;
   BenchUut3.processSequence[1] := USINT#2;
   BenchUut3.processSequence[2] := USINT#2;
   BenchUut3.processSequence[3] := USINT#5;
   BenchUut3.processSequence[4] := USINT#0;
   BenchUut3.processSequence[5] := USINT#0;
   BenchUut3.processSequence[6] := USINT#0;
   BenchUut3.processSequence[7] := USINT#0;
   BenchUut3.processSequence[8] := USINT#0;
   TraceIn_processLength[22] := BenchUut3.processLength;
   TraceIn_sensor1[22] := BenchUut3.sensor1;
   TraceIn_sensor2[22] := BenchUut3.sensor2;
   TraceIn_sensor3[22] := BenchUut3.sensor3;
   TraceIn_sensor4[22] := BenchUut3.sensor4;
   TraceIn_sensor5[22] := BenchUut3.sensor5;
   TraceIn_station1Start[22] := BenchUut3.station1Start;
   TraceIn_station2Complete[22] := BenchUut3.station2Complete;
   TraceIn_station3Complete[22] := BenchUut3.station3Complete;
   TraceIn_station4Complete[22] := BenchUut3.station4Complete;
   TraceIn_processSequence_1[22] := BenchUut3.processSequence[1];
   TraceIn_processSequence_2[22] := BenchUut3.processSequence[2];
   TraceIn_processSequence_3[22] := BenchUut3.processSequence[3];
   TraceIn_processSequence_4[22] := BenchUut3.processSequence[4];
   TraceIn_processSequence_5[22] := BenchUut3.processSequence[5];
   TraceIn_processSequence_6[22] := BenchUut3.processSequence[6];
   TraceIn_processSequence_7[22] := BenchUut3.processSequence[7];
   TraceIn_processSequence_8[22] := BenchUut3.processSequence[8];
   BenchUut3();
   TraceOut_conveyorLeft[22] := BenchUut3.conveyorLeft;
   TraceOut_conveyorRight[22] := BenchUut3.conveyorRight;
   BenchCalls := BenchCalls + 1;
 23:
   BenchUut3.processLength := USINT#3;
   BenchUut3.sensor1 := FALSE;
   BenchUut3.sensor2 := TRUE;
   BenchUut3.sensor3 := FALSE;
   BenchUut3.sensor4 := FALSE;
   BenchUut3.sensor5 := FALSE;
   BenchUut3.station1Start := FALSE;
   BenchUut3.station2Complete := TRUE;
   BenchUut3.station3Complete := FALSE;
   BenchUut3.station4Complete := FALSE;
   BenchUut3.processSequence[1] := USINT#2;
   BenchUut3.processSequence[2] := USINT#2;
   BenchUut3.processSequence[3] := USINT#5;
   BenchUut3.processSequence[4] := USINT#0;
   BenchUut3.processSequence[5] := USINT#0;
   BenchUut3.processSequence[6] := USINT#0;
   BenchUut3.processSequence[7] := USINT#0;
   BenchUut3.processSequence[8] := USINT#0;
   TraceIn_processLength[23] := BenchUut3.processLength;
   TraceIn_sensor1[23] := BenchUut3.sensor1;
   TraceIn_sensor2[23] := BenchUut3.sensor2;
   TraceIn_sensor3[23] := BenchUut3.sensor3;
   TraceIn_sensor4[23] := BenchUut3.sensor4;
   TraceIn_sensor5[23] := BenchUut3.sensor5;
   TraceIn_station1Start[23] := BenchUut3.station1Start;
   TraceIn_station2Complete[23] := BenchUut3.station2Complete;
   TraceIn_station3Complete[23] := BenchUut3.station3Complete;
   TraceIn_station4Complete[23] := BenchUut3.station4Complete;
   TraceIn_processSequence_1[23] := BenchUut3.processSequence[1];
   TraceIn_processSequence_2[23] := BenchUut3.processSequence[2];
   TraceIn_processSequence_3[23] := BenchUut3.processSequence[3];
   TraceIn_processSequence_4[23] := BenchUut3.processSequence[4];
   TraceIn_processSequence_5[23] := BenchUut3.processSequence[5];
   TraceIn_processSequence_6[23] := BenchUut3.processSequence[6];
   TraceIn_processSequence_7[23] := BenchUut3.processSequence[7];
   TraceIn_processSequence_8[23] := BenchUut3.processSequence[8];
   BenchUut3();
   TraceOut_conveyorLeft[23] := BenchUut3.conveyorLeft;
   TraceOut_conveyorRight[23] := BenchUut3.conveyorRight;
   BenchCalls := BenchCalls + 1;
 24:
   BenchUut3.processLength := USINT#3;
   BenchUut3.sensor1 := FALSE;
   BenchUut3.sensor2 := TRUE;
   BenchUut3.sensor3 := FALSE;
   BenchUut3.sensor4 := FALSE;
   BenchUut3.sensor5 := FALSE;
   BenchUut3.station1Start := FALSE;
   BenchUut3.station2Complete := FALSE;
   BenchUut3.station3Complete := FALSE;
   BenchUut3.station4Complete := FALSE;
   BenchUut3.processSequence[1] := USINT#2;
   BenchUut3.processSequence[2] := USINT#2;
   BenchUut3.processSequence[3] := USINT#5;
   BenchUut3.processSequence[4] := USINT#0;
   BenchUut3.processSequence[5] := USINT#0;
   BenchUut3.processSequence[6] := USINT#0;
   BenchUut3.processSequence[7] := USINT#0;
   BenchUut3.processSequence[8] := USINT#0;
   TraceIn_processLength[24] := BenchUut3.processLength;
   TraceIn_sensor1[24] := BenchUut3.sensor1;
   TraceIn_sensor2[24] := BenchUut3.sensor2;
   TraceIn_sensor3[24] := BenchUut3.sensor3;
   TraceIn_sensor4[24] := BenchUut3.sensor4;
   TraceIn_sensor5[24] := BenchUut3.sensor5;
   TraceIn_station1Start[24] := BenchUut3.station1Start;
   TraceIn_station2Complete[24] := BenchUut3.station2Complete;
   TraceIn_station3Complete[24] := BenchUut3.station3Complete;
   TraceIn_station4Complete[24] := BenchUut3.station4Complete;
   TraceIn_processSequence_1[24] := BenchUut3.processSequence[1];
   TraceIn_processSequence_2[24] := BenchUut3.processSequence[2];
   TraceIn_processSequence_3[24] := BenchUut3.processSequence[3];
   TraceIn_processSequence_4[24] := BenchUut3.processSequence[4];
   TraceIn_processSequence_5[24] := BenchUut3.processSequence[5];
   TraceIn_processSequence_6[24] := BenchUut3.processSequence[6];
   TraceIn_processSequence_7[24] := BenchUut3.processSequence[7];
   TraceIn_processSequence_8[24] := BenchUut3.processSequence[8];
   BenchUut3();
   TraceOut_conveyorLeft[24] := BenchUut3.conveyorLeft;
   TraceOut_conveyorRight[24] := BenchUut3.conveyorRight;
   BenchCalls := BenchCalls + 1;
 25:
   BenchUut3.processLength := USINT#3;
   BenchUut3.sensor1 := FALSE;
   BenchUut3.sensor2 := TRUE;
   BenchUut3.sensor3 := FALSE;
   BenchUut3.sensor4 := FALSE;
   BenchUut3.sensor5 := FALSE;
   BenchUut3.station1Start := FALSE;
   BenchUut3.station2Complete := TRUE;
   BenchUut3.station3Complete := FALSE;
   BenchUut3.station4Complete := FALSE;
   BenchUut3.processSequence[1] := USINT#2;
   BenchUut3.processSequence[2] := USINT#2;
   BenchUut3.processSequence[3] := USINT#5;
   BenchUut3.processSequence[4] := USINT#0;
   BenchUut3.processSequence[5] := USINT#0;
   BenchUut3.processSequence[6] := USINT#0;
   BenchUut3.processSequence[7] := USINT#0;
   BenchUut3.processSequence[8] := USINT#0;
   TraceIn_processLength[25] := BenchUut3.processLength;
   TraceIn_sensor1[25] := BenchUut3.sensor1;
   TraceIn_sensor2[25] := BenchUut3.sensor2;
   TraceIn_sensor3[25] := BenchUut3.sensor3;
   TraceIn_sensor4[25] := BenchUut3.sensor4;
   TraceIn_sensor5[25] := BenchUut3.sensor5;
   TraceIn_station1Start[25] := BenchUut3.station1Start;
   TraceIn_station2Complete[25] := BenchUut3.station2Complete;
   TraceIn_station3Complete[25] := BenchUut3.station3Complete;
   TraceIn_station4Complete[25] := BenchUut3.station4Complete;
   TraceIn_processSequence_1[25] := BenchUut3.processSequence[1];
   TraceIn_processSequence_2[25] := BenchUut3.processSequence[2];
   TraceIn_processSequence_3[25] := BenchUut3.processSequence[3];
   TraceIn_processSequence_4[25] := BenchUut3.processSequence[4];
   TraceIn_processSequence_5[25] := BenchUut3.processSequence[5];
   TraceIn_processSequence_6[25] := BenchUut3.processSequence[6];
   TraceIn_processSequence_7[25] := BenchUut3.processSequence[7];
   TraceIn_processSequence_8[25] := BenchUut3.processSequence[8];
   BenchUut3();
   TraceOut_conveyorLeft[25] := BenchUut3.conveyorLeft;
   TraceOut_conveyorRight[25] := BenchUut3.conveyorRight;
   BenchCalls := BenchCalls + 1;
 26:
   BenchUut3.processLength := USINT#3;
   BenchUut3.sensor1 := FALSE;
   BenchUut3.sensor2 := FALSE;
   BenchUut3.sensor3 := FALSE;
   BenchUut3.sensor4 := FALSE;
   BenchUut3.sensor5 := TRUE;
   BenchUut3.station1Start := FALSE;
   BenchUut3.station2Complete := FALSE;
   BenchUut3.station3Complete := FALSE;
   BenchUut3.station4Complete := FALSE;
   BenchUut3.processSequence[1] := USINT#2;
   BenchUut3.processSequence[2] := USINT#2;
   BenchUut3.processSequence[3] := USINT#5;
   BenchUut3.processSequence[4] := USINT#0;
   BenchUut3.processSequence[5] := USINT#0;
   BenchUut3.processSequence[6] := USINT#0;
   BenchUut3.processSequence[7] := USINT#0;
   BenchUut3.processSequence[8] := USINT#0;
   TraceIn_processLength[26] := BenchUut3.processLength;
   TraceIn_sensor1[26] := BenchUut3.sensor1;
   TraceIn_sensor2[26] := BenchUut3.sensor2;
   TraceIn_sensor3[26] := BenchUut3.sensor3;
   TraceIn_sensor4[26] := BenchUut3.sensor4;
   TraceIn_sensor5[26] := BenchUut3.sensor5;
   TraceIn_station1Start[26] := BenchUut3.station1Start;
   TraceIn_station2Complete[26] := BenchUut3.station2Complete;
   TraceIn_station3Complete[26] := BenchUut3.station3Complete;
   TraceIn_station4Complete[26] := BenchUut3.station4Complete;
   TraceIn_processSequence_1[26] := BenchUut3.processSequence[1];
   TraceIn_processSequence_2[26] := BenchUut3.processSequence[2];
   TraceIn_processSequence_3[26] := BenchUut3.processSequence[3];
   TraceIn_processSequence_4[26] := BenchUut3.processSequence[4];
   TraceIn_processSequence_5[26] := BenchUut3.processSequence[5];
   TraceIn_processSequence_6[26] := BenchUut3.processSequence[6];
   TraceIn_processSequence_7[26] := BenchUut3.processSequence[7];
   TraceIn_processSequence_8[26] := BenchUut3.processSequence[8];
   BenchUut3();
   TraceOut_conveyorLeft[26] := BenchUut3.conveyorLeft;
   TraceOut_conveyorRight[26] := BenchUut3.conveyorRight;
   BenchCalls := BenchCalls + 1;
 27:
   BenchUut4.processLength := USINT#8;
   BenchUut4.sensor1 := FALSE;
   BenchUut4.sensor2 := FALSE;
   BenchUut4.sensor3 := FALSE;
   BenchUut4.sensor4 := FALSE;
   BenchUut4.sensor5 := FALSE;
   BenchUut4.station1Start := TRUE;
   BenchUut4.station2Complete := FALSE;
   BenchUut4.station3Complete := FALSE;
   BenchUut4.station4Complete := FALSE;
   BenchUut4.processSequence[1] := USINT#4;
   BenchUut4.processSequence[2] := USINT#3;
   BenchUut4.processSequence[3] := USINT#2;
   BenchUut4.processSequence[4] := USINT#4;
   BenchUut4.processSequence[5] := USINT#2;
   BenchUut4.processSequence[6] := USINT#3;
   BenchUut4.processSequence[7] := USINT#4;
   BenchUut4.processSequence[8] := USINT#5;
   TraceIn_processLength[27] := BenchUut4.processLength;
   TraceIn_sensor1[27] := BenchUut4.sensor1;
   TraceIn_sensor2[27] := BenchUut4.sensor2;
   TraceIn_sensor3[27] := BenchUut4.sensor3;
   TraceIn_sensor4[27] := BenchUut4.sensor4;
   TraceIn_sensor5[27] := BenchUut4.sensor5;
   TraceIn_station1Start[27] := BenchUut4.station1Start;
   TraceIn_station2Complete[27] := BenchUut4.station2Complete;
   TraceIn_station3Complete[27] := BenchUut4.station3Complete;
   TraceIn_station4Complete[27] := BenchUut4.station4Complete;
   TraceIn_processSequence_1[27] := BenchUut4.processSequence[1];
   TraceIn_processSequence_2[27] := BenchUut4.processSequence[2];
   TraceIn_processSequence_3[27] := BenchUut4.processSequence[3];
   TraceIn_processSequence_4[27] := BenchUut4.processSequence[4];
   TraceIn_processSequence_5[27] := BenchUut4.processSequence[5];
   TraceIn_processSequence_6[27] := BenchUut4.processSequence[6];
   TraceIn_processSequence_7[27] := BenchUut4.processSequence[7];
   TraceIn_processSequence_8[27] := BenchUut4.processSequence[8];
   BenchUut4();
   TraceOut_conveyorLeft[27] := BenchUut4.conveyorLeft;
   TraceOut_conveyorRight[27] := BenchUut4.conveyorRight;
   BenchCalls := BenchCalls + 1;
 28:
   BenchUut4.processLength := USINT#8;
   BenchUut4.sensor1 := TRUE;
   BenchUut4.sensor2 := FALSE;
   BenchUut4.sensor3 := FALSE;
   BenchUut4.sensor4 := FALSE;
   BenchUut4.sensor5 := FALSE;
   BenchUut4.station1Start := TRUE;
   BenchUut4.station2Complete := FALSE;
   BenchUut4.station3Complete := FALSE;
   BenchUut4.station4Complete := FALSE;
   BenchUut4.processSequence[1] := USINT#4;
   BenchUut4.processSequence[2] := USINT#3;
   BenchUut4.processSequence[3] := USINT#2;
   BenchUut4.processSequence[4] := USINT#4;
   BenchUut4.processSequence[5] := USINT#2;
   BenchUut4.processSequence[6] := USINT#3;
   BenchUut4.processSequence[7] := USINT#4;
   BenchUut4.processSequence[8] := USINT#5;
   TraceIn_processLength[28] := BenchUut4.processLength;
   TraceIn_sensor1[28] := BenchUut4.sensor1;
   TraceIn_sensor2[28] := BenchUut4.sensor2;
   TraceIn_sensor3[28] := BenchUut4.sensor3;
   TraceIn_sensor4[28] := BenchUut4.sensor4;
   TraceIn_sensor5[28] := BenchUut4.sensor5;
   TraceIn_station1Start[28] := BenchUut4.station1Start;
   TraceIn_station2Complete[28] := BenchUut4.station2Complete;
   TraceIn_station3Complete[28] := BenchUut4.station3Complete;
   TraceIn_station4Complete[28] := BenchUut4.station4Complete;
   TraceIn_processSequence_1[28] := BenchUut4.processSequence[1];
   TraceIn_processSequence_2[28] := BenchUut4.processSequence[2];
   TraceIn_processSequence_3[28] := BenchUut4.processSequence[3];
   TraceIn_processSequence_4[28] := BenchUut4.processSequence[4];
   TraceIn_processSequence_5[28] := BenchUut4.processSequence[5];
   TraceIn_processSequence_6[28] := BenchUut4.processSequence[6];
   TraceIn_processSequence_7[28] := BenchUut4.processSequence[7];
   TraceIn_processSequence_8[28] := BenchUut4.processSequence[8];
   BenchUut4();
   TraceOut_conveyorLeft[28] := BenchUut4.conveyorLeft;
   TraceOut_conveyorRight[28] := BenchUut4.conveyorRight;
   BenchCalls := BenchCalls + 1;
 29:
   BenchUut4.processLength := USINT#8;
   BenchUut4.sensor1 := FALSE;
   BenchUut4.sensor2 := TRUE;
   BenchUut4.sensor3 := FALSE;
   BenchUut4.sensor4 := FALSE;
   BenchUut4.sensor5 := FALSE;
   BenchUut4.station1Start := FALSE;
   BenchUut4.station2Complete := FALSE;
   BenchUut4.station3Complete := FALSE;
   BenchUut4.station4Complete := FALSE;
   BenchUut4.processSequence[1] := USINT#4;
   BenchUut4.processSequence[2] := USINT#3;
   BenchUut4.processSequence[3] := USINT#2;
   BenchUut4.processSequence[4] := USINT#4;
   BenchUut4.processSequence[5] := USINT#2;
   BenchUut4.processSequence[6] := USINT#3;
   BenchUut4.processSequence[7] := USINT#4;
   BenchUut4.processSequence[8] := USINT#5;
   TraceIn_processLength[29] := BenchUut4.processLength;
   TraceIn_sensor1[29] := BenchUut4.sensor1;
   TraceIn_sensor2[29] := BenchUut4.sensor2;
   TraceIn_sensor3[29] := BenchUut4.sensor3;
   TraceIn_sensor4[29] := BenchUut4.sensor4;
   TraceIn_sensor5[29] := BenchUut4.sensor5;
   TraceIn_station1Start[29] := BenchUut4.station1Start;
   TraceIn_station2Complete[29] := BenchUut4.station2Complete;
   TraceIn_station3Complete[29] := BenchUut4.station3Complete;
   TraceIn_station4Complete[29] := BenchUut4.station4Complete;
   TraceIn_processSequence_1[29] := BenchUut4.processSequence[1];
   TraceIn_processSequence_2[29] := BenchUut4.processSequence[2];
   TraceIn_processSequence_3[29] := BenchUut4.processSequence[3];
   TraceIn_processSequence_4[29] := BenchUut4.processSequence[4];
   TraceIn_processSequence_5[29] := BenchUut4.processSequence[5];
   TraceIn_processSequence_6[29] := BenchUut4.processSequence[6];
   TraceIn_processSequence_7[29] := BenchUut4.processSequence[7];
   TraceIn_processSequence_8[29] := BenchUut4.processSequence[8];
   BenchUut4();
   TraceOut_conveyorLeft[29] := BenchUut4.conveyorLeft;
   TraceOut_conveyorRight[29] := BenchUut4.conveyorRight;
   BenchCalls := BenchCalls + 1;
 30:
   BenchUut4.processLength := USINT#8;
   BenchUut4.sensor1 := FALSE;
   BenchUut4.sensor2 := FALSE;
   BenchUut4.sensor3 := FALSE;
   BenchUut4.sensor4 := FALSE;
   BenchUut4.sensor5 := FALSE;
   BenchUut4.station1Start := FALSE;
   BenchUut4.station2Complete := FALSE;
   BenchUut4.station3Complete := FALSE;
   BenchUut4.station4Complete := FALSE;
   BenchUut4.processSequence[1] := USINT#4;
   BenchUut4.processSequence[2] := USINT#3;
   BenchUut4.processSequence[3] := USINT#2;
   BenchUut4.processSequence[4] := USINT#4;
   BenchUut4.processSequence[5] := USINT#2;
   BenchUut4.processSequence[6] := USINT#3;
   BenchUut4.processSequence[7] := USINT#4;
   BenchUut4.processSequence[8] := USINT#5;
   TraceIn_processLength[30] := BenchUut4.processLength;
   TraceIn_sensor1[30] := BenchUut4.sensor1;
   TraceIn_sensor2[30] := BenchUut4.sensor2;
   TraceIn_sensor3[30] := BenchUut4.sensor3;
   TraceIn_sensor4[30] := BenchUut4.sensor4;
   TraceIn_sensor5[30] := BenchUut4.sensor5;
   TraceIn_station1Start[30] := BenchUut4.station1Start;
   TraceIn_station2Complete[30] := BenchUut4.station2Complete;
   TraceIn_station3Complete[30] := BenchUut4.station3Complete;
   TraceIn_station4Complete[30] := BenchUut4.station4Complete;
   TraceIn_processSequence_1[30] := BenchUut4.processSequence[1];
   TraceIn_processSequence_2[30] := BenchUut4.processSequence[2];
   TraceIn_processSequence_3[30] := BenchUut4.processSequence[3];
   TraceIn_processSequence_4[30] := BenchUut4.processSequence[4];
   TraceIn_processSequence_5[30] := BenchUut4.processSequence[5];
   TraceIn_processSequence_6[30] := BenchUut4.processSequence[6];
   TraceIn_processSequence_7[30] := BenchUut4.processSequence[7];
   TraceIn_processSequence_8[30] := BenchUut4.processSequence[8];
   BenchUut4();
   TraceOut_conveyorLeft[30] := BenchUut4.conveyorLeft;
   TraceOut_conveyorRight[30] := BenchUut4.conveyorRight;
   BenchCalls := BenchCalls + 1;
 31:
   BenchUut4.processLength := USINT#8;
   BenchUut4.sensor1 := FALSE;
   BenchUut4.sensor2 := FALSE;
   BenchUut4.sensor3 := FALSE;
   BenchUut4.sensor4 := TRUE;
   BenchUut4.sensor5 := FALSE;
   BenchUut4.station1Start := FALSE;
   BenchUut4.station2Complete := FALSE;
   BenchUut4.station3Complete := FALSE;
   BenchUut4.station4Complete := FALSE;
   BenchUut4.processSequence[1] := USINT#4;
   BenchUut4.processSequence[2] := USINT#3;
   BenchUut4.processSequence[3] := USINT#2;
   BenchUut4.processSequence[4] := USINT#4;
   BenchUut4.processSequence[5] := USINT#2;
   BenchUut4.processSequence[6] := USINT#3;
   BenchUut4.processSequence[7] := USINT#4;
   BenchUut4.processSequence[8] := USINT#5;
   TraceIn_processLength[31] := BenchUut4.processLength;
   TraceIn_sensor1[31] := BenchUut4.sensor1;
   TraceIn_sensor2[31] := BenchUut4.sensor2;
   TraceIn_sensor3[31] := BenchUut4.sensor3;
   TraceIn_sensor4[31] := BenchUut4.sensor4;
   TraceIn_sensor5[31] := BenchUut4.sensor5;
   TraceIn_station1Start[31] := BenchUut4.station1Start;
   TraceIn_station2Complete[31] := BenchUut4.station2Complete;
   TraceIn_station3Complete[31] := BenchUut4.station3Complete;
   TraceIn_station4Complete[31] := BenchUut4.station4Complete;
   TraceIn_processSequence_1[31] := BenchUut4.processSequence[1];
   TraceIn_processSequence_2[31] := BenchUut4.processSequence[2];
   TraceIn_processSequence_3[31] := BenchUut4.processSequence[3];
   TraceIn_processSequence_4[31] := BenchUut4.processSequence[4];
   TraceIn_processSequence_5[31] := BenchUut4.processSequence[5];
   TraceIn_processSequence_6[31] := BenchUut4.processSequence[6];
   TraceIn_processSequence_7[31] := BenchUut4.processSequence[7];
   TraceIn_processSequence_8[31] := BenchUut4.processSequence[8];
   BenchUut4();
   TraceOut_conveyorLeft[31] := BenchUut4.conveyorLeft;
   TraceOut_conveyorRight[31] := BenchUut4.conveyorRight;
   BenchCalls := BenchCalls + 1;
 32:
   BenchUut4.processLength := USINT#8;
   BenchUut4.sensor1 := FALSE;
   BenchUut4.sensor2 := FALSE;
   BenchUut4.sensor3 := FALSE;
   BenchUut4.sensor4 := TRUE;
   BenchUut4.sensor5 := FALSE;
   BenchUut4.station1Start := FALSE;
   BenchUut4.station2Complete := FALSE;
   BenchUut4.station3Complete := FALSE;
   BenchUut4.station4Complete := TRUE;
   BenchUut4.processSequence[1] := USINT#4;
   BenchUut4.processSequence[2] := USINT#3;
   BenchUut4.processSequence[3] := USINT#2;
   BenchUut4.processSequence[4] := USINT#4;
   BenchUut4.processSequence[5] := USINT#2;
   BenchUut4.processSequence[6] := USINT#3;
   BenchUut4.processSequence[7] := USINT#4;
   BenchUut4.processSequence[8] := USINT#5;
   TraceIn_processLength[32] := BenchUut4.processLength;
   TraceIn_sensor1[32] := BenchUut4.sensor1;
   TraceIn_sensor2[32] := BenchUut4.sensor2;
   TraceIn_sensor3[32] := BenchUut4.sensor3;
   TraceIn_sensor4[32] := BenchUut4.sensor4;
   TraceIn_sensor5[32] := BenchUut4.sensor5;
   TraceIn_station1Start[32] := BenchUut4.station1Start;
   TraceIn_station2Complete[32] := BenchUut4.station2Complete;
   TraceIn_station3Complete[32] := BenchUut4.station3Complete;
   TraceIn_station4Complete[32] := BenchUut4.station4Complete;
   TraceIn_processSequence_1[32] := BenchUut4.processSequence[1];
   TraceIn_processSequence_2[32] := BenchUut4.processSequence[2];
   TraceIn_processSequence_3[32] := BenchUut4.processSequence[3];
   TraceIn_processSequence_4[32] := BenchUut4.processSequence[4];
   TraceIn_processSequence_5[32] := BenchUut4.processSequence[5];
   TraceIn_processSequence_6[32] := BenchUut4.processSequence[6];
   TraceIn_processSequence_7[32] := BenchUut4.processSequence[7];
   TraceIn_processSequence_8[32] := BenchUut4.processSequence[8];
   BenchUut4();
   TraceOut_conveyorLeft[32] := BenchUut4.conveyorLeft;
   TraceOut_conveyorRight[32] := BenchUut4.conveyorRight;
   BenchCalls := BenchCalls + 1;
 33:
   BenchUut4.processLength := USINT#8;
   BenchUut4.sensor1 := FALSE;
   BenchUut4.sensor2 := FALSE;
   BenchUut4.sensor3 := FALSE;
   BenchUut4.sensor4 := FALSE;
   BenchUut4.sensor5 := FALSE;
   BenchUut4.station1Start := FALSE;
   BenchUut4.station2Complete := FALSE;
   BenchUut4.station3Complete := FALSE;
   BenchUut4.station4Complete := FALSE;
   BenchUut4.processSequence[1] := USINT#4;
   BenchUut4.processSequence[2] := USINT#3;
   BenchUut4.processSequence[3] := USINT#2;
   BenchUut4.processSequence[4] := USINT#4;
   BenchUut4.processSequence[5] := USINT#2;
   BenchUut4.processSequence[6] := USINT#3;
   BenchUut4.processSequence[7] := USINT#4;
   BenchUut4.processSequence[8] := USINT#5;
   TraceIn_processLength[33] := BenchUut4.processLength;
   TraceIn_sensor1[33] := BenchUut4.sensor1;
   TraceIn_sensor2[33] := BenchUut4.sensor2;
   TraceIn_sensor3[33] := BenchUut4.sensor3;
   TraceIn_sensor4[33] := BenchUut4.sensor4;
   TraceIn_sensor5[33] := BenchUut4.sensor5;
   TraceIn_station1Start[33] := BenchUut4.station1Start;
   TraceIn_station2Complete[33] := BenchUut4.station2Complete;
   TraceIn_station3Complete[33] := BenchUut4.station3Complete;
   TraceIn_station4Complete[33] := BenchUut4.station4Complete;
   TraceIn_processSequence_1[33] := BenchUut4.processSequence[1];
   TraceIn_processSequence_2[33] := BenchUut4.processSequence[2];
   TraceIn_processSequence_3[33] := BenchUut4.processSequence[3];
   TraceIn_processSequence_4[33] := BenchUut4.processSequence[4];
   TraceIn_processSequence_5[33] := BenchUut4.processSequence[5];
   TraceIn_processSequence_6[33] := BenchUut4.processSequence[6];
   TraceIn_processSequence_7[33] := BenchUut4.processSequence[7];
   TraceIn_processSequence_8[33] := BenchUut4.processSequence[8];
   BenchUut4();
   TraceOut_conveyorLeft[33] := BenchUut4.conveyorLeft;
   TraceOut_conveyorRight[33] := BenchUut4.conveyorRight;
   BenchCalls := BenchCalls + 1;
 34:
   BenchUut4.processLength := USINT#8;
   BenchUut4.sensor1 := FALSE;
   BenchUut4.sensor2 := FALSE;
   BenchUut4.sensor3 := TRUE;
   BenchUut4.sensor4 := FALSE;
   BenchUut4.sensor5 := FALSE;
   BenchUut4.station1Start := FALSE;
   BenchUut4.station2Complete := FALSE;
   BenchUut4.station3Complete := FALSE;
   BenchUut4.station4Complete := FALSE;
   BenchUut4.processSequence[1] := USINT#4;
   BenchUut4.processSequence[2] := USINT#3;
   BenchUut4.processSequence[3] := USINT#2;
   BenchUut4.processSequence[4] := USINT#4;
   BenchUut4.processSequence[5] := USINT#2;
   BenchUut4.processSequence[6] := USINT#3;
   BenchUut4.processSequence[7] := USINT#4;
   BenchUut4.processSequence[8] := USINT#5;
   TraceIn_processLength[34] := BenchUut4.processLength;
   TraceIn_sensor1[34] := BenchUut4.sensor1;
   TraceIn_sensor2[34] := BenchUut4.sensor2;
   TraceIn_sensor3[34] := BenchUut4.sensor3;
   TraceIn_sensor4[34] := BenchUut4.sensor4;
   TraceIn_sensor5[34] := BenchUut4.sensor5;
   TraceIn_station1Start[34] := BenchUut4.station1Start;
   TraceIn_station2Complete[34] := BenchUut4.station2Complete;
   TraceIn_station3Complete[34] := BenchUut4.station3Complete;
   TraceIn_station4Complete[34] := BenchUut4.station4Complete;
   TraceIn_processSequence_1[34] := BenchUut4.processSequence[1];
   TraceIn_processSequence_2[34] := BenchUut4.processSequence[2];
   TraceIn_processSequence_3[34] := BenchUut4.processSequence[3];
   TraceIn_processSequence_4[34] := BenchUut4.processSequence[4];
   TraceIn_processSequence_5[34] := BenchUut4.processSequence[5];
   TraceIn_processSequence_6[34] := BenchUut4.processSequence[6];
   TraceIn_processSequence_7[34] := BenchUut4.processSequence[7];
   TraceIn_processSequence_8[34] := BenchUut4.processSequence[8];
   BenchUut4();
   TraceOut_conveyorLeft[34] := BenchUut4.conveyorLeft;
   TraceOut_conveyorRight[34] := BenchUut4.conveyorRight;
   BenchCalls := BenchCalls + 1;
 35:
   BenchUut4.processLength := USINT#8;
   BenchUut4.sensor1 := FALSE;
   BenchUut4.sensor2 := FALSE;
   BenchUut4.sensor3 := TRUE;
   BenchUut4.sensor4 := FALSE;
   BenchUut4.sensor5 := FALSE;
   BenchUut4.station1Start := FALSE;
   BenchUut4.station2Complete := FALSE;
   BenchUut4.station3Complete := TRUE;
   BenchUut4.station4Complete := FALSE;
   BenchUut4.processSequence[1] := USINT#4;
   BenchUut4.processSequence[2] := USINT#3;
   BenchUut4.processSequence[3] := USINT#2;
   BenchUut4.processSequence[4] := USINT#4;
   BenchUut4.processSequence[5] := USINT#2;
   BenchUut4.processSequence[6] := USINT#3;
   BenchUut4.processSequence[7] := USINT#4;
   BenchUut4.processSequence[8] := USINT#5;
   TraceIn_processLength[35] := BenchUut4.processLength;
   TraceIn_sensor1[35] := BenchUut4.sensor1;
   TraceIn_sensor2[35] := BenchUut4.sensor2;
   TraceIn_sensor3[35] := BenchUut4.sensor3;
   TraceIn_sensor4[35] := BenchUut4.sensor4;
   TraceIn_sensor5[35] := BenchUut4.sensor5;
   TraceIn_station1Start[35] := BenchUut4.station1Start;
   TraceIn_station2Complete[35] := BenchUut4.station2Complete;
   TraceIn_station3Complete[35] := BenchUut4.station3Complete;
   TraceIn_station4Complete[35] := BenchUut4.station4Complete;
   TraceIn_processSequence_1[35] := BenchUut4.processSequence[1];
   TraceIn_processSequence_2[35] := BenchUut4.processSequence[2];
   TraceIn_processSequence_3[35] := BenchUut4.processSequence[3];
   TraceIn_processSequence_4[35] := BenchUut4.processSequence[4];
   TraceIn_processSequence_5[35] := BenchUut4.processSequence[5];
   TraceIn_processSequence_6[35] := BenchUut4.processSequence[6];
   TraceIn_processSequence_7[35] := BenchUut4.processSequence[7];
   TraceIn_processSequence_8[35] := BenchUut4.processSequence[8];
   BenchUut4();
   TraceOut_conveyorLeft[35] := BenchUut4.conveyorLeft;
   TraceOut_conveyorRight[35] := BenchUut4.conveyorRight;
   BenchCalls := BenchCalls + 1;
 36:
   BenchUut4.processLength := USINT#8;
   BenchUut4.sensor1 := FALSE;
   BenchUut4.sensor2 := TRUE;
   BenchUut4.sensor3 := FALSE;
   BenchUut4.sensor4 := FALSE;
   BenchUut4.sensor5 := FALSE;
   BenchUut4.station1Start := FALSE;
   BenchUut4.station2Complete := FALSE;
   BenchUut4.station3Complete := FALSE;
   BenchUut4.station4Complete := FALSE;
   BenchUut4.processSequence[1] := USINT#4;
   BenchUut4.processSequence[2] := USINT#3;
   BenchUut4.processSequence[3] := USINT#2;
   BenchUut4.processSequence[4] := USINT#4;
   BenchUut4.processSequence[5] := USINT#2;
   BenchUut4.processSequence[6] := USINT#3;
   BenchUut4.processSequence[7] := USINT#4;
   BenchUut4.processSequence[8] := USINT#5;
   TraceIn_processLength[36] := BenchUut4.processLength;
   TraceIn_sensor1[36] := BenchUut4.sensor1;
   TraceIn_sensor2[36] := BenchUut4.sensor2;
   TraceIn_sensor3[36] := BenchUut4.sensor3;
   TraceIn_sensor4[36] := BenchUut4.sensor4;
   TraceIn_sensor5[36] := BenchUut4.sensor5;
   TraceIn_station1Start[36] := BenchUut4.station1Start;
   TraceIn_station2Complete[36] := BenchUut4.station2Complete;
   TraceIn_station3Complete[36] := BenchUut4.station3Complete;
   TraceIn_station4Complete[36] := BenchUut4.station4Complete;
   TraceIn_processSequence_1[36] := BenchUut4.processSequence[1];
   TraceIn_processSequence_2[36] := BenchUut4.processSequence[2];
   TraceIn_processSequence_3[36] := BenchUut4.processSequence[3];
   TraceIn_processSequence_4[36] := BenchUut4.processSequence[4];
   TraceIn_processSequence_5[36] := BenchUut4.processSequence[5];
   TraceIn_processSequence_6[36] := BenchUut4.processSequence[6];
   TraceIn_processSequence_7[36] := BenchUut4.processSequence[7];
   TraceIn_processSequence_8[36] := BenchUut4.processSequence[8];
   BenchUut4();
   TraceOut_conveyorLeft[36] := BenchUut4.conveyorLeft;
   TraceOut_conveyorRight[36] := BenchUut4.conveyorRight;
   BenchCalls := BenchCalls + 1;
 37:
   BenchUut4.processLength := USINT#8;
   BenchUut4.sensor1 := FALSE;
   BenchUut4.sensor2 := TRUE;
   BenchUut4.sensor3 := FALSE;
   BenchUut4.sensor4 := FALSE;
   BenchUut4.sensor5 := FALSE;
   BenchUut4.station1Start := FALSE;
   BenchUut4.station2Complete := TRUE;
   BenchUut4.station3Complete := FALSE;
   BenchUut4.station4Complete := FALSE;
   BenchUut4.processSequence[1] := USINT#4;
   BenchUut4.processSequence[2] := USINT#3;
   BenchUut4.processSequence[3] := USINT#2;
   BenchUut4.processSequence[4] := USINT#4;
   BenchUut4.processSequence[5] := USINT#2;
   BenchUut4.processSequence[6] := USINT#3;
   BenchUut4.processSequence[7] := USINT#4;
   BenchUut4.processSequence[8] := USINT#5;
   TraceIn_processLength[37] := BenchUut4.processLength;
   TraceIn_sensor1[37] := BenchUut4.sensor1;
   TraceIn_sensor2[37] := BenchUut4.sensor2;
   TraceIn_sensor3[37] := BenchUut4.sensor3;
   TraceIn_sensor4[37] := BenchUut4.sensor4;
   TraceIn_sensor5[37] := BenchUut4.sensor5;
   TraceIn_station1Start[37] := BenchUut4.station1Start;
   TraceIn_station2Complete[37] := BenchUut4.station2Complete;
   TraceIn_station3Complete[37] := BenchUut4.station3Complete;
   TraceIn_station4Complete[37] := BenchUut4.station4Complete;
   TraceIn_processSequence_1[37] := BenchUut4.processSequence[1];
   TraceIn_processSequence_2[37] := BenchUut4.processSequence[2];
   TraceIn_processSequence_3[37] := BenchUut4.processSequence[3];
   TraceIn_processSequence_4[37] := BenchUut4.processSequence[4];
   TraceIn_processSequence_5[37] := BenchUut4.processSequence[5];
   TraceIn_processSequence_6[37] := BenchUut4.processSequence[6];
   TraceIn_processSequence_7[37] := BenchUut4.processSequence[7];
   TraceIn_processSequence_8[37] := BenchUut4.processSequence[8];
   BenchUut4();
   TraceOut_conveyorLeft[37] := BenchUut4.conveyorLeft;
   TraceOut_conveyorRight[37] := BenchUut4.conveyorRight;
   BenchCalls := BenchCalls + 1;
 38:
   BenchUut4.processLength := USINT#8;
   BenchUut4.sensor1 := FALSE;
   BenchUut4.sensor2 := FALSE;
   BenchUut4.sensor3 := FALSE;
   BenchUut4.sensor4 := TRUE;
   BenchUut4.sensor5 := FALSE;
   BenchUut4.station1Start := FALSE;
   BenchUut4.station2Complete := FALSE;
   BenchUut4.station3Complete := FALSE;
   BenchUut4.station4Complete := FALSE;
   BenchUut4.processSequence[1] := USINT#4;
   BenchUut4.processSequence[2] := USINT#3;
   BenchUut4.processSequence[3] := USINT#2;
   BenchUut4.processSequence[4] := USINT#4;
   BenchUut4.processSequence[5] := USINT#2;
   BenchUut4.processSequence[6] := USINT#3;
   BenchUut4.processSequence[7] := USINT#4;
   BenchUut4.processSequence[8] := USINT#5;
   TraceIn_processLength[38] := BenchUut4.processLength;
   TraceIn_sensor1[38] := BenchUut4.sensor1;
   TraceIn_sensor2[38] := BenchUut4.sensor2;
   TraceIn_sensor3[38] := BenchUut4.sensor3;
   TraceIn_sensor4[38] := BenchUut4.sensor4;
   TraceIn_sensor5[38] := BenchUut4.sensor5;
   TraceIn_station1Start[38] := BenchUut4.station1Start;
   TraceIn_station2Complete[38] := BenchUut4.station2Complete;
   TraceIn_station3Complete[38] := BenchUut4.station3Complete;
   TraceIn_station4Complete[38] := BenchUut4.station4Complete;
   TraceIn_processSequence_1[38] := BenchUut4.processSequence[1];
   TraceIn_processSequence_2[38] := BenchUut4.processSequence[2];
   TraceIn_processSequence_3[38] := BenchUut4.processSequence[3];
   TraceIn_processSequence_4[38] := BenchUut4.processSequence[4];
   TraceIn_processSequence_5[38] := BenchUut4.processSequence[5];
   TraceIn_processSequence_6[38] := BenchUut4.processSequence[6];
   TraceIn_processSequence_7[38] := BenchUut4.processSequence[7];
   TraceIn_processSequence_8[38] := BenchUut4.processSequence[8];
   BenchUut4();
   TraceOut_conveyorLeft[38] := BenchUut4.conveyorLeft;
   TraceOut_conveyorRight[38] := BenchUut4.conveyorRight;
   BenchCalls := BenchCalls + 1;
 39:
   BenchUut4.processLength := USINT#8;
   BenchUut4.sensor1 := FALSE;
   BenchUut4.sensor2 := FALSE;
   BenchUut4.sensor3 := FALSE;
   BenchUut4.sensor4 := TRUE;
   BenchUut4.sensor5 := FALSE;
   BenchUut4.station1Start := FALSE;
   BenchUut4.station2Complete := FALSE;
   BenchUut4.station3Complete := FALSE;
   BenchUut4.station4Complete := TRUE;
   BenchUut4.processSequence[1] := USINT#4;
   BenchUut4.processSequence[2] := USINT#3;
   BenchUut4.processSequence[3] := USINT#2;
   BenchUut4.processSequence[4] := USINT#4;
   BenchUut4.processSequence[5] := USINT#2;
   BenchUut4.processSequence[6] := USINT#3;
   BenchUut4.processSequence[7] := USINT#4;
   BenchUut4.processSequence[8] := USINT#5;
   TraceIn_processLength[39] := BenchUut4.processLength;
   TraceIn_sensor1[39] := BenchUut4.sensor1;
   TraceIn_sensor2[39] := BenchUut4.sensor2;
   TraceIn_sensor3[39] := BenchUut4.sensor3;
   TraceIn_sensor4[39] := BenchUut4.sensor4;
   TraceIn_sensor5[39] := BenchUut4.sensor5;
   TraceIn_station1Start[39] := BenchUut4.station1Start;
   TraceIn_station2Complete[39] := BenchUut4.station2Complete;
   TraceIn_station3Complete[39] := BenchUut4.station3Complete;
   TraceIn_station4Complete[39] := BenchUut4.station4Complete;
   TraceIn_processSequence_1[39] := BenchUut4.processSequence[1];
   TraceIn_processSequence_2[39] := BenchUut4.processSequence[2];
   TraceIn_processSequence_3[39] := BenchUut4.processSequence[3];
   TraceIn_processSequence_4[39] := BenchUut4.processSequence[4];
   TraceIn_processSequence_5[39] := BenchUut4.processSequence[5];
   TraceIn_processSequence_6[39] := BenchUut4.processSequence[6];
   TraceIn_processSequence_7[39] := BenchUut4.processSequence[7];
   TraceIn_processSequence_8[39] := BenchUut4.processSequence[8];
   BenchUut4();
   TraceOut_conveyorLeft[39] := BenchUut4.conveyorLeft;
   TraceOut_conveyorRight[39] := BenchUut4.conveyorRight;
   BenchCalls := BenchCalls + 1;
 40:
   BenchUut4.processLength := USINT#8;
   BenchUut4.sensor1 := FALSE;
   BenchUut4.sensor2 := TRUE;
   BenchUut4.sensor3 := FALSE;
   BenchUut4.sensor4 := FALSE;
   BenchUut4.sensor5 := FALSE;
   BenchUut4.station1Start := FALSE;
   BenchUut4.station2Complete := FALSE;
   BenchUut4.station3Complete := FALSE;
   BenchUut4.station4Complete := FALSE;
   BenchUut4.processSequence[1] := USINT#4;
   BenchUut4.processSequence[2] := USINT#3;
   BenchUut4.processSequence[3] := USINT#2;
   BenchUut4.processSequence[4] := USINT#4;
   BenchUut4.processSequence[5] := USINT#2;
   BenchUut4.processSequence[6] := USINT#3;
   BenchUut4.processSequence[7] := USINT#4;
   BenchUut4.processSequence[8] := USINT#5;
   TraceIn_processLength[40] := BenchUut4.processLength;
   TraceIn_sensor1[40] := BenchUut4.sensor1;
   TraceIn_sensor2[40] := BenchUut4.sensor2;
   TraceIn_sensor3[40] := BenchUut4.sensor3;
   TraceIn_sensor4[40] := BenchUut4.sensor4;
   TraceIn_sensor5[40] := BenchUut4.sensor5;
   TraceIn_station1Start[40] := BenchUut4.station1Start;
   TraceIn_station2Complete[40] := BenchUut4.station2Complete;
   TraceIn_station3Complete[40] := BenchUut4.station3Complete;
   TraceIn_station4Complete[40] := BenchUut4.station4Complete;
   TraceIn_processSequence_1[40] := BenchUut4.processSequence[1];
   TraceIn_processSequence_2[40] := BenchUut4.processSequence[2];
   TraceIn_processSequence_3[40] := BenchUut4.processSequence[3];
   TraceIn_processSequence_4[40] := BenchUut4.processSequence[4];
   TraceIn_processSequence_5[40] := BenchUut4.processSequence[5];
   TraceIn_processSequence_6[40] := BenchUut4.processSequence[6];
   TraceIn_processSequence_7[40] := BenchUut4.processSequence[7];
   TraceIn_processSequence_8[40] := BenchUut4.processSequence[8];
   BenchUut4();
   TraceOut_conveyorLeft[40] := BenchUut4.conveyorLeft;
   TraceOut_conveyorRight[40] := BenchUut4.conveyorRight;
   BenchCalls := BenchCalls + 1;
 41:
   BenchUut4.processLength := USINT#8;
   BenchUut4.sensor1 := FALSE;
   BenchUut4.sensor2 := TRUE;
   BenchUut4.sensor3 := FALSE;
   BenchUut4.sensor4 := FALSE;
   BenchUut4.sensor5 := FALSE;
   BenchUut4.station1Start := FALSE;
   BenchUut4.station2Complete := TRUE;
   BenchUut4.station3Complete := FALSE;
   BenchUut4.station4Complete := FALSE;
   BenchUut4.processSequence[1] := USINT#4;
   BenchUut4.processSequence[2] := USINT#3;
   BenchUut4.processSequence[3] := USINT#2;
   BenchUut4.processSequence[4] := USINT#4;
   BenchUut4.processSequence[5] := USINT#2;
   BenchUut4.processSequence[6] := USINT#3;
   BenchUut4.processSequence[7] := USINT#4;
   BenchUut4.processSequence[8] := USINT#5;
   TraceIn_processLength[41] := BenchUut4.processLength;
   TraceIn_sensor1[41] := BenchUut4.sensor1;
   TraceIn_sensor2[41] := BenchUut4.sensor2;
   TraceIn_sensor3[41] := BenchUut4.sensor3;
   TraceIn_sensor4[41] := BenchUut4.sensor4;
   TraceIn_sensor5[41] := BenchUut4.sensor5;
   TraceIn_station1Start[41] := BenchUut4.station1Start;
   TraceIn_station2Complete[41] := BenchUut4.station2Complete;
   TraceIn_station3Complete[41] := BenchUut4.station3Complete;
   TraceIn_station4Complete[41] := BenchUut4.station4Complete;
   TraceIn_processSequence_1[41] := BenchUut4.processSequence[1];
   TraceIn_processSequence_2[41] := BenchUut4.processSequence[2];
   TraceIn_processSequence_3[41] := BenchUut4.processSequence[3];
   TraceIn_processSequence_4[41] := BenchUut4.processSequence[4];
   TraceIn_processSequence_5[41] := BenchUut4.processSequence[5];
   TraceIn_processSequence_6[41] := BenchUut4.processSequence[6];
   TraceIn_processSequence_7[41] := BenchUut4.processSequence[7];
   TraceIn_processSequence_8[41] := BenchUut4.processSequence[8];
   BenchUut4();
   TraceOut_conveyorLeft[41] := BenchUut4.conveyorLeft;
   TraceOut_conveyorRight[41] := BenchUut4.conveyorRight;
   BenchCalls := BenchCalls + 1;
 42:
   BenchUut4.processLength := USINT#8;
   BenchUut4.sensor1 := FALSE;
   BenchUut4.sensor2 := FALSE;
   BenchUut4.sensor3 := TRUE;
   BenchUut4.sensor4 := FALSE;
   BenchUut4.sensor5 := FALSE;
   BenchUut4.station1Start := FALSE;
   BenchUut4.station2Complete := FALSE;
   BenchUut4.station3Complete := FALSE;
   BenchUut4.station4Complete := FALSE;
   BenchUut4.processSequence[1] := USINT#4;
   BenchUut4.processSequence[2] := USINT#3;
   BenchUut4.processSequence[3] := USINT#2;
   BenchUut4.processSequence[4] := USINT#4;
   BenchUut4.processSequence[5] := USINT#2;
   BenchUut4.processSequence[6] := USINT#3;
   BenchUut4.processSequence[7] := USINT#4;
   BenchUut4.processSequence[8] := USINT#5;
   TraceIn_processLength[42] := BenchUut4.processLength;
   TraceIn_sensor1[42] := BenchUut4.sensor1;
   TraceIn_sensor2[42] := BenchUut4.sensor2;
   TraceIn_sensor3[42] := BenchUut4.sensor3;
   TraceIn_sensor4[42] := BenchUut4.sensor4;
   TraceIn_sensor5[42] := BenchUut4.sensor5;
   TraceIn_station1Start[42] := BenchUut4.station1Start;
   TraceIn_station2Complete[42] := BenchUut4.station2Complete;
   TraceIn_station3Complete[42] := BenchUut4.station3Complete;
   TraceIn_station4Complete[42] := BenchUut4.station4Complete;
   TraceIn_processSequence_1[42] := BenchUut4.processSequence[1];
   TraceIn_processSequence_2[42] := BenchUut4.processSequence[2];
   TraceIn_processSequence_3[42] := BenchUut4.processSequence[3];
   TraceIn_processSequence_4[42] := BenchUut4.processSequence[4];
   TraceIn_processSequence_5[42] := BenchUut4.processSequence[5];
   TraceIn_processSequence_6[42] := BenchUut4.processSequence[6];
   TraceIn_processSequence_7[42] := BenchUut4.processSequence[7];
   TraceIn_processSequence_8[42] := BenchUut4.processSequence[8];
   BenchUut4();
   TraceOut_conveyorLeft[42] := BenchUut4.conveyorLeft;
   TraceOut_conveyorRight[42] := BenchUut4.conveyorRight;
   BenchCalls := BenchCalls + 1;
 43:
   BenchUut4.processLength := USINT#8;
   BenchUut4.sensor1 := FALSE;
   BenchUut4.sensor2 := FALSE;
   BenchUut4.sensor3 := TRUE;
   BenchUut4.sensor4 := FALSE;
   BenchUut4.sensor5 := FALSE;
   BenchUut4.station1Start := FALSE;
   BenchUut4.station2Complete := FALSE;
   BenchUut4.station3Complete := TRUE;
   BenchUut4.station4Complete := FALSE;
   BenchUut4.processSequence[1] := USINT#4;
   BenchUut4.processSequence[2] := USINT#3;
   BenchUut4.processSequence[3] := USINT#2;
   BenchUut4.processSequence[4] := USINT#4;
   BenchUut4.processSequence[5] := USINT#2;
   BenchUut4.processSequence[6] := USINT#3;
   BenchUut4.processSequence[7] := USINT#4;
   BenchUut4.processSequence[8] := USINT#5;
   TraceIn_processLength[43] := BenchUut4.processLength;
   TraceIn_sensor1[43] := BenchUut4.sensor1;
   TraceIn_sensor2[43] := BenchUut4.sensor2;
   TraceIn_sensor3[43] := BenchUut4.sensor3;
   TraceIn_sensor4[43] := BenchUut4.sensor4;
   TraceIn_sensor5[43] := BenchUut4.sensor5;
   TraceIn_station1Start[43] := BenchUut4.station1Start;
   TraceIn_station2Complete[43] := BenchUut4.station2Complete;
   TraceIn_station3Complete[43] := BenchUut4.station3Complete;
   TraceIn_station4Complete[43] := BenchUut4.station4Complete;
   TraceIn_processSequence_1[43] := BenchUut4.processSequence[1];
   TraceIn_processSequence_2[43] := BenchUut4.processSequence[2];
   TraceIn_processSequence_3[43] := BenchUut4.processSequence[3];
   TraceIn_processSequence_4[43] := BenchUut4.processSequence[4];
   TraceIn_processSequence_5[43] := BenchUut4.processSequence[5];
   TraceIn_processSequence_6[43] := BenchUut4.processSequence[6];
   TraceIn_processSequence_7[43] := BenchUut4.processSequence[7];
   TraceIn_processSequence_8[43] := BenchUut4.processSequence[8];
   BenchUut4();
   TraceOut_conveyorLeft[43] := BenchUut4.conveyorLeft;
   TraceOut_conveyorRight[43] := BenchUut4.conveyorRight;
   BenchCalls := BenchCalls + 1;
 44:
   BenchUut4.processLength := USINT#8;
   BenchUut4.sensor1 := FALSE;
   BenchUut4.sensor2 := FALSE;
   BenchUut4.sensor3 := FALSE;
   BenchUut4.sensor4 := TRUE;
   BenchUut4.sensor5 := FALSE;
   BenchUut4.station1Start := FALSE;
   BenchUut4.station2Complete := FALSE;
   BenchUut4.station3Complete := FALSE;
   BenchUut4.station4Complete := FALSE;
   BenchUut4.processSequence[1] := USINT#4;
   BenchUut4.processSequence[2] := USINT#3;
   BenchUut4.processSequence[3] := USINT#2;
   BenchUut4.processSequence[4] := USINT#4;
   BenchUut4.processSequence[5] := USINT#2;
   BenchUut4.processSequence[6] := USINT#3;
   BenchUut4.processSequence[7] := USINT#4;
   BenchUut4.processSequence[8] := USINT#5;
   TraceIn_processLength[44] := BenchUut4.processLength;
   TraceIn_sensor1[44] := BenchUut4.sensor1;
   TraceIn_sensor2[44] := BenchUut4.sensor2;
   TraceIn_sensor3[44] := BenchUut4.sensor3;
   TraceIn_sensor4[44] := BenchUut4.sensor4;
   TraceIn_sensor5[44] := BenchUut4.sensor5;
   TraceIn_station1Start[44] := BenchUut4.station1Start;
   TraceIn_station2Complete[44] := BenchUut4.station2Complete;
   TraceIn_station3Complete[44] := BenchUut4.station3Complete;
   TraceIn_station4Complete[44] := BenchUut4.station4Complete;
   TraceIn_processSequence_1[44] := BenchUut4.processSequence[1];
   TraceIn_processSequence_2[44] := BenchUut4.processSequence[2];
   TraceIn_processSequence_3[44] := BenchUut4.processSequence[3];
   TraceIn_processSequence_4[44] := BenchUut4.processSequence[4];
   TraceIn_processSequence_5[44] := BenchUut4.processSequence[5];
   TraceIn_processSequence_6[44] := BenchUut4.processSequence[6];
   TraceIn_processSequence_7[44] := BenchUut4.processSequence[7];
   TraceIn_processSequence_8[44] := BenchUut4.processSequence[8];
   BenchUut4();
   TraceOut_conveyorLeft[44] := BenchUut4.conveyorLeft;
   TraceOut_conveyorRight[44] := BenchUut4.conveyorRight;
   BenchCalls := BenchCalls + 1;
 45:
   BenchUut4.processLength := USINT#8;
   BenchUut4.sensor1 := FALSE;
   BenchUut4.sensor2 := FALSE;
   BenchUut4.sensor3 := FALSE;
   BenchUut4.sensor4 := TRUE;
   BenchUut4.sensor5 := FALSE;
   BenchUut4.station1Start := FALSE;
   BenchUut4.station2Complete := FALSE;
   BenchUut4.station3Complete := FALSE;
   BenchUut4.station4Complete := TRUE;
   BenchUut4.processSequence[1] := USINT#4;
   BenchUut4.processSequence[2] := USINT#3;
   BenchUut4.processSequence[3] := USINT#2;
   BenchUut4.processSequence[4] := USINT#4;
   BenchUut4.processSequence[5] := USINT#2;
   BenchUut4.processSequence[6] := USINT#3;
   BenchUut4.processSequence[7] := USINT#4;
   BenchUut4.processSequence[8] := USINT#5;
   TraceIn_processLength[45] := BenchUut4.processLength;
   TraceIn_sensor1[45] := BenchUut4.sensor1;
   TraceIn_sensor2[45] := BenchUut4.sensor2;
   TraceIn_sensor3[45] := BenchUut4.sensor3;
   TraceIn_sensor4[45] := BenchUut4.sensor4;
   TraceIn_sensor5[45] := BenchUut4.sensor5;
   TraceIn_station1Start[45] := BenchUut4.station1Start;
   TraceIn_station2Complete[45] := BenchUut4.station2Complete;
   TraceIn_station3Complete[45] := BenchUut4.station3Complete;
   TraceIn_station4Complete[45] := BenchUut4.station4Complete;
   TraceIn_processSequence_1[45] := BenchUut4.processSequence[1];
   TraceIn_processSequence_2[45] := BenchUut4.processSequence[2];
   TraceIn_processSequence_3[45] := BenchUut4.processSequence[3];
   TraceIn_processSequence_4[45] := BenchUut4.processSequence[4];
   TraceIn_processSequence_5[45] := BenchUut4.processSequence[5];
   TraceIn_processSequence_6[45] := BenchUut4.processSequence[6];
   TraceIn_processSequence_7[45] := BenchUut4.processSequence[7];
   TraceIn_processSequence_8[45] := BenchUut4.processSequence[8];
   BenchUut4();
   TraceOut_conveyorLeft[45] := BenchUut4.conveyorLeft;
   TraceOut_conveyorRight[45] := BenchUut4.conveyorRight;
   BenchCalls := BenchCalls + 1;
 46:
   BenchUut4.processLength := USINT#8;
   BenchUut4.sensor1 := FALSE;
   BenchUut4.sensor2 := FALSE;
   BenchUut4.sensor3 := FALSE;
   BenchUut4.sensor4 := FALSE;
   BenchUut4.sensor5 := TRUE;
   BenchUut4.station1Start := FALSE;
   BenchUut4.station2Complete := FALSE;
   BenchUut4.station3Complete := FALSE;
   BenchUut4.station4Complete := FALSE;
   BenchUut4.processSequence[1] := USINT#4;
   BenchUut4.processSequence[2] := USINT#3;
   BenchUut4.processSequence[3] := USINT#2;
   BenchUut4.processSequence[4] := USINT#4;
   BenchUut4.processSequence[5] := USINT#2;
   BenchUut4.processSequence[6] := USINT#3;
   BenchUut4.processSequence[7] := USINT#4;
   BenchUut4.processSequence[8] := USINT#5;
   TraceIn_processLength[46] := BenchUut4.processLength;
   TraceIn_sensor1[46] := BenchUut4.sensor1;
   TraceIn_sensor2[46] := BenchUut4.sensor2;
   TraceIn_sensor3[46] := BenchUut4.sensor3;
   TraceIn_sensor4[46] := BenchUut4.sensor4;
   TraceIn_sensor5[46] := BenchUut4.sensor5;
   TraceIn_station1Start[46] := BenchUut4.station1Start;
   TraceIn_station2Complete[46] := BenchUut4.station2Complete;
   TraceIn_station3Complete[46] := BenchUut4.station3Complete;
   TraceIn_station4Complete[46] := BenchUut4.station4Complete;
   TraceIn_processSequence_1[46] := BenchUut4.processSequence[1];
   TraceIn_processSequence_2[46] := BenchUut4.processSequence[2];
   TraceIn_processSequence_3[46] := BenchUut4.processSequence[3];
   TraceIn_processSequence_4[46] := BenchUut4.processSequence[4];
   TraceIn_processSequence_5[46] := BenchUut4.processSequence[5];
   TraceIn_processSequence_6[46] := BenchUut4.processSequence[6];
   TraceIn_processSequence_7[46] := BenchUut4.processSequence[7];
   TraceIn_processSequence_8[46] := BenchUut4.processSequence[8];
   BenchUut4();
   TraceOut_conveyorLeft[46] := BenchUut4.conveyorLeft;
   TraceOut_conveyorRight[46] := BenchUut4.conveyorRight;
   BenchCalls := BenchCalls + 1;
 47:
   BenchUut5.processLength := USINT#8;
   BenchUut5.sensor1 := TRUE;
   BenchUut5.sensor2 := FALSE;
   BenchUut5.sensor3 := FALSE;
   BenchUut5.sensor4 := FALSE;
   BenchUut5.sensor5 := FALSE;
   BenchUut5.station1Start := TRUE;
   BenchUut5.station2Complete := FALSE;
   BenchUut5.station3Complete := FALSE;
   BenchUut5.station4Complete := FALSE;
   BenchUut5.processSequence[1] := USINT#2;
   BenchUut5.processSequence[2] := USINT#3;
   BenchUut5.processSequence[3] := USINT#4;
   BenchUut5.processSequence[4] := USINT#3;
   BenchUut5.processSequence[5] := USINT#2;
   BenchUut5.processSequence[6] := USINT#4;
   BenchUut5.processSequence[7] := USINT#3;
   BenchUut5.processSequence[8] := USINT#5;
   TraceIn_processLength[47] := BenchUut5.processLength;
   TraceIn_sensor1[47] := BenchUut5.sensor1;
   TraceIn_sensor2[47] := BenchUut5.sensor2;
   TraceIn_sensor3[47] := BenchUut5.sensor3;
   TraceIn_sensor4[47] := BenchUut5.sensor4;
   TraceIn_sensor5[47] := BenchUut5.sensor5;
   TraceIn_station1Start[47] := BenchUut5.station1Start;
   TraceIn_station2Complete[47] := BenchUut5.station2Complete;
   TraceIn_station3Complete[47] := BenchUut5.station3Complete;
   TraceIn_station4Complete[47] := BenchUut5.station4Complete;
   TraceIn_processSequence_1[47] := BenchUut5.processSequence[1];
   TraceIn_processSequence_2[47] := BenchUut5.processSequence[2];
   TraceIn_processSequence_3[47] := BenchUut5.processSequence[3];
   TraceIn_processSequence_4[47] := BenchUut5.processSequence[4];
   TraceIn_processSequence_5[47] := BenchUut5.processSequence[5];
   TraceIn_processSequence_6[47] := BenchUut5.processSequence[6];
   TraceIn_processSequence_7[47] := BenchUut5.processSequence[7];
   TraceIn_processSequence_8[47] := BenchUut5.processSequence[8];
   BenchUut5();
   TraceOut_conveyorLeft[47] := BenchUut5.conveyorLeft;
   TraceOut_conveyorRight[47] := BenchUut5.conveyorRight;
   BenchCalls := BenchCalls + 1;
 48:
   BenchUut5.processLength := USINT#8;
   BenchUut5.sensor1 := FALSE;
   BenchUut5.sensor2 := FALSE;
   BenchUut5.sensor3 := FALSE;
   BenchUut5.sensor4 := FALSE;
   BenchUut5.sensor5 := FALSE;
   BenchUut5.station1Start := FALSE;
   BenchUut5.station2Complete := FALSE;
   BenchUut5.station3Complete := FALSE;
   BenchUut5.station4Complete := FALSE;
   BenchUut5.processSequence[1] := USINT#2;
   BenchUut5.processSequence[2] := USINT#3;
   BenchUut5.processSequence[3] := USINT#4;
   BenchUut5.processSequence[4] := USINT#3;
   BenchUut5.processSequence[5] := USINT#2;
   BenchUut5.processSequence[6] := USINT#4;
   BenchUut5.processSequence[7] := USINT#3;
   BenchUut5.processSequence[8] := USINT#5;
   TraceIn_processLength[48] := BenchUut5.processLength;
   TraceIn_sensor1[48] := BenchUut5.sensor1;
   TraceIn_sensor2[48] := BenchUut5.sensor2;
   TraceIn_sensor3[48] := BenchUut5.sensor3;
   TraceIn_sensor4[48] := BenchUut5.sensor4;
   TraceIn_sensor5[48] := BenchUut5.sensor5;
   TraceIn_station1Start[48] := BenchUut5.station1Start;
   TraceIn_station2Complete[48] := BenchUut5.station2Complete;
   TraceIn_station3Complete[48] := BenchUut5.station3Complete;
   TraceIn_station4Complete[48] := BenchUut5.station4Complete;
   TraceIn_processSequence_1[48] := BenchUut5.processSequence[1];
   TraceIn_processSequence_2[48] := BenchUut5.processSequence[2];
   TraceIn_processSequence_3[48] := BenchUut5.processSequence[3];
   TraceIn_processSequence_4[48] := BenchUut5.processSequence[4];
   TraceIn_processSequence_5[48] := BenchUut5.processSequence[5];
   TraceIn_processSequence_6[48] := BenchUut5.processSequence[6];
   TraceIn_processSequence_7[48] := BenchUut5.processSequence[7];
   TraceIn_processSequence_8[48] := BenchUut5.processSequence[8];
   BenchUut5();
   TraceOut_conveyorLeft[48] := BenchUut5.conveyorLeft;
   TraceOut_conveyorRight[48] := BenchUut5.conveyorRight;
   BenchCalls := BenchCalls + 1;
 49:
   BenchUut5.processLength := USINT#8;
   BenchUut5.sensor1 := FALSE;
   BenchUut5.sensor2 := FALSE;
   BenchUut5.sensor3 := FALSE;
   BenchUut5.sensor4 := FALSE;
   BenchUut5.sensor5 := FALSE;
   BenchUut5.station1Start := FALSE;
   BenchUut5.station2Complete := FALSE;
   BenchUut5.station3Complete := FALSE;
   BenchUut5.station4Complete := FALSE;
   BenchUut5.processSequence[1] := USINT#2;
   BenchUut5.processSequence[2] := USINT#3;
   BenchUut5.processSequence[3] := USINT#4;
   BenchUut5.processSequence[4] := USINT#3;
   BenchUut5.processSequence[5] := USINT#2;
   BenchUut5.processSequence[6] := USINT#4;
   BenchUut5.processSequence[7] := USINT#3;
   BenchUut5.processSequence[8] := USINT#5;
   TraceIn_processLength[49] := BenchUut5.processLength;
   TraceIn_sensor1[49] := BenchUut5.sensor1;
   TraceIn_sensor2[49] := BenchUut5.sensor2;
   TraceIn_sensor3[49] := BenchUut5.sensor3;
   TraceIn_sensor4[49] := BenchUut5.sensor4;
   TraceIn_sensor5[49] := BenchUut5.sensor5;
   TraceIn_station1Start[49] := BenchUut5.station1Start;
   TraceIn_station2Complete[49] := BenchUut5.station2Complete;
   TraceIn_station3Complete[49] := BenchUut5.station3Complete;
   TraceIn_station4Complete[49] := BenchUut5.station4Complete;
   TraceIn_processSequence_1[49] := BenchUut5.processSequence[1];
   TraceIn_processSequence_2[49] := BenchUut5.processSequence[2];
   TraceIn_processSequence_3[49] := BenchUut5.processSequence[3];
   TraceIn_processSequence_4[49] := BenchUut5.processSequence[4];
   TraceIn_processSequence_5[49] := BenchUut5.processSequence[5];
   TraceIn_processSequence_6[49] := BenchUut5.processSequence[6];
   TraceIn_processSequence_7[49] := BenchUut5.processSequence[7];
   TraceIn_processSequence_8[49] := BenchUut5.processSequence[8];
   BenchUut5();
   TraceOut_conveyorLeft[49] := BenchUut5.conveyorLeft;
   TraceOut_conveyorRight[49] := BenchUut5.conveyorRight;
   BenchCalls := BenchCalls + 1;
 50:
   BenchUut5.processLength := USINT#8;
   BenchUut5.sensor1 := FALSE;
   BenchUut5.sensor2 := TRUE;
   BenchUut5.sensor3 := FALSE;
   BenchUut5.sensor4 := FALSE;
   BenchUut5.sensor5 := FALSE;
   BenchUut5.station1Start := FALSE;
   BenchUut5.station2Complete := FALSE;
   BenchUut5.station3Complete := FALSE;
   BenchUut5.station4Complete := FALSE;
   BenchUut5.processSequence[1] := USINT#2;
   BenchUut5.processSequence[2] := USINT#3;
   BenchUut5.processSequence[3] := USINT#4;
   BenchUut5.processSequence[4] := USINT#3;
   BenchUut5.processSequence[5] := USINT#2;
   BenchUut5.processSequence[6] := USINT#4;
   BenchUut5.processSequence[7] := USINT#3;
   BenchUut5.processSequence[8] := USINT#5;
   TraceIn_processLength[50] := BenchUut5.processLength;
   TraceIn_sensor1[50] := BenchUut5.sensor1;
   TraceIn_sensor2[50] := BenchUut5.sensor2;
   TraceIn_sensor3[50] := BenchUut5.sensor3;
   TraceIn_sensor4[50] := BenchUut5.sensor4;
   TraceIn_sensor5[50] := BenchUut5.sensor5;
   TraceIn_station1Start[50] := BenchUut5.station1Start;
   TraceIn_station2Complete[50] := BenchUut5.station2Complete;
   TraceIn_station3Complete[50] := BenchUut5.station3Complete;
   TraceIn_station4Complete[50] := BenchUut5.station4Complete;
   TraceIn_processSequence_1[50] := BenchUut5.processSequence[1];
   TraceIn_processSequence_2[50] := BenchUut5.processSequence[2];
   TraceIn_processSequence_3[50] := BenchUut5.processSequence[3];
   TraceIn_processSequence_4[50] := BenchUut5.processSequence[4];
   TraceIn_processSequence_5[50] := BenchUut5.processSequence[5];
   TraceIn_processSequence_6[50] := BenchUut5.processSequence[6];
   TraceIn_processSequence_7[50] := BenchUut5.processSequence[7];
   TraceIn_processSequence_8[50] := BenchUut5.processSequence[8];
   BenchUut5();
   TraceOut_conveyorLeft[50] := BenchUut5.conveyorLeft;
   TraceOut_conveyorRight[50] := BenchUut5.conveyorRight;
   BenchCalls := BenchCalls + 1;
 51:
   BenchUut5.processLength := USINT#8;
   BenchUut5.sensor1 := FALSE;
   BenchUut5.sensor2 := TRUE;
   BenchUut5.sensor3 := FALSE;
   BenchUut5.sensor4 := FALSE;
   BenchUut5.sensor5 := FALSE;
   BenchUut5.station1Start := FALSE;
   BenchUut5.station2Complete := FALSE;
   BenchUut5.station3Complete := FALSE;
   BenchUut5.station4Complete := FALSE;
   BenchUut5.processSequence[1] := USINT#2;
   BenchUut5.processSequence[2] := USINT#3;
   BenchUut5.processSequence[3] := USINT#4;
   BenchUut5.processSequence[4] := USINT#3;
   BenchUut5.processSequence[5] := USINT#2;
   BenchUut5.processSequence[6] := USINT#4;
   BenchUut5.processSequence[7] := USINT#3;
   BenchUut5.processSequence[8] := USINT#5;
   TraceIn_processLength[51] := BenchUut5.processLength;
   TraceIn_sensor1[51] := BenchUut5.sensor1;
   TraceIn_sensor2[51] := BenchUut5.sensor2;
   TraceIn_sensor3[51] := BenchUut5.sensor3;
   TraceIn_sensor4[51] := BenchUut5.sensor4;
   TraceIn_sensor5[51] := BenchUut5.sensor5;
   TraceIn_station1Start[51] := BenchUut5.station1Start;
   TraceIn_station2Complete[51] := BenchUut5.station2Complete;
   TraceIn_station3Complete[51] := BenchUut5.station3Complete;
   TraceIn_station4Complete[51] := BenchUut5.station4Complete;
   TraceIn_processSequence_1[51] := BenchUut5.processSequence[1];
   TraceIn_processSequence_2[51] := BenchUut5.processSequence[2];
   TraceIn_processSequence_3[51] := BenchUut5.processSequence[3];
   TraceIn_processSequence_4[51] := BenchUut5.processSequence[4];
   TraceIn_processSequence_5[51] := BenchUut5.processSequence[5];
   TraceIn_processSequence_6[51] := BenchUut5.processSequence[6];
   TraceIn_processSequence_7[51] := BenchUut5.processSequence[7];
   TraceIn_processSequence_8[51] := BenchUut5.processSequence[8];
   BenchUut5();
   TraceOut_conveyorLeft[51] := BenchUut5.conveyorLeft;
   TraceOut_conveyorRight[51] := BenchUut5.conveyorRight;
   BenchCalls := BenchCalls + 1;
 52:
   BenchUut5.processLength := USINT#8;
   BenchUut5.sensor1 := FALSE;
   BenchUut5.sensor2 := TRUE;
   BenchUut5.sensor3 := FALSE;
   BenchUut5.sensor4 := FALSE;
   BenchUut5.sensor5 := FALSE;
   BenchUut5.station1Start := FALSE;
   BenchUut5.station2Complete := FALSE;
   BenchUut5.station3Complete := FALSE;
   BenchUut5.station4Complete := FALSE;
   BenchUut5.processSequence[1] := USINT#2;
   BenchUut5.processSequence[2] := USINT#3;
   BenchUut5.processSequence[3] := USINT#4;
   BenchUut5.processSequence[4] := USINT#3;
   BenchUut5.processSequence[5] := USINT#2;
   BenchUut5.processSequence[6] := USINT#4;
   BenchUut5.processSequence[7] := USINT#3;
   BenchUut5.processSequence[8] := USINT#5;
   TraceIn_processLength[52] := BenchUut5.processLength;
   TraceIn_sensor1[52] := BenchUut5.sensor1;
   TraceIn_sensor2[52] := BenchUut5.sensor2;
   TraceIn_sensor3[52] := BenchUut5.sensor3;
   TraceIn_sensor4[52] := BenchUut5.sensor4;
   TraceIn_sensor5[52] := BenchUut5.sensor5;
   TraceIn_station1Start[52] := BenchUut5.station1Start;
   TraceIn_station2Complete[52] := BenchUut5.station2Complete;
   TraceIn_station3Complete[52] := BenchUut5.station3Complete;
   TraceIn_station4Complete[52] := BenchUut5.station4Complete;
   TraceIn_processSequence_1[52] := BenchUut5.processSequence[1];
   TraceIn_processSequence_2[52] := BenchUut5.processSequence[2];
   TraceIn_processSequence_3[52] := BenchUut5.processSequence[3];
   TraceIn_processSequence_4[52] := BenchUut5.processSequence[4];
   TraceIn_processSequence_5[52] := BenchUut5.processSequence[5];
   TraceIn_processSequence_6[52] := BenchUut5.processSequence[6];
   TraceIn_processSequence_7[52] := BenchUut5.processSequence[7];
   TraceIn_processSequence_8[52] := BenchUut5.processSequence[8];
   BenchUut5();
   TraceOut_conveyorLeft[52] := BenchUut5.conveyorLeft;
   TraceOut_conveyorRight[52] := BenchUut5.conveyorRight;
   BenchCalls := BenchCalls + 1;
 53:
   BenchUut5.processLength := USINT#8;
   BenchUut5.sensor1 := FALSE;
   BenchUut5.sensor2 := TRUE;
   BenchUut5.sensor3 := FALSE;
   BenchUut5.sensor4 := FALSE;
   BenchUut5.sensor5 := FALSE;
   BenchUut5.station1Start := FALSE;
   BenchUut5.station2Complete := TRUE;
   BenchUut5.station3Complete := FALSE;
   BenchUut5.station4Complete := FALSE;
   BenchUut5.processSequence[1] := USINT#2;
   BenchUut5.processSequence[2] := USINT#3;
   BenchUut5.processSequence[3] := USINT#4;
   BenchUut5.processSequence[4] := USINT#3;
   BenchUut5.processSequence[5] := USINT#2;
   BenchUut5.processSequence[6] := USINT#4;
   BenchUut5.processSequence[7] := USINT#3;
   BenchUut5.processSequence[8] := USINT#5;
   TraceIn_processLength[53] := BenchUut5.processLength;
   TraceIn_sensor1[53] := BenchUut5.sensor1;
   TraceIn_sensor2[53] := BenchUut5.sensor2;
   TraceIn_sensor3[53] := BenchUut5.sensor3;
   TraceIn_sensor4[53] := BenchUut5.sensor4;
   TraceIn_sensor5[53] := BenchUut5.sensor5;
   TraceIn_station1Start[53] := BenchUut5.station1Start;
   TraceIn_station2Complete[53] := BenchUut5.station2Complete;
   TraceIn_station3Complete[53] := BenchUut5.station3Complete;
   TraceIn_station4Complete[53] := BenchUut5.station4Complete;
   TraceIn_processSequence_1[53] := BenchUut5.processSequence[1];
   TraceIn_processSequence_2[53] := BenchUut5.processSequence[2];
   TraceIn_processSequence_3[53] := BenchUut5.processSequence[3];
   TraceIn_processSequence_4[53] := BenchUut5.processSequence[4];
   TraceIn_processSequence_5[53] := BenchUut5.processSequence[5];
   TraceIn_processSequence_6[53] := BenchUut5.processSequence[6];
   TraceIn_processSequence_7[53] := BenchUut5.processSequence[7];
   TraceIn_processSequence_8[53] := BenchUut5.processSequence[8];
   BenchUut5();
   TraceOut_conveyorLeft[53] := BenchUut5.conveyorLeft;
   TraceOut_conveyorRight[53] := BenchUut5.conveyorRight;
   BenchCalls := BenchCalls + 1;
 54:
   BenchUut5.processLength := USINT#8;
   BenchUut5.sensor1 := FALSE;
   BenchUut5.sensor2 := FALSE;
   BenchUut5.sensor3 := FALSE;
   BenchUut5.sensor4 := FALSE;
   BenchUut5.sensor5 := FALSE;
   BenchUut5.station1Start := FALSE;
   BenchUut5.station2Complete := FALSE;
   BenchUut5.station3Complete := FALSE;
   BenchUut5.station4Complete := FALSE;
   BenchUut5.processSequence[1] := USINT#2;
   BenchUut5.processSequence[2] := USINT#3;
   BenchUut5.processSequence[3] := USINT#4;
   BenchUut5.processSequence[4] := USINT#3;
   BenchUut5.processSequence[5] := USINT#2;
   BenchUut5.processSequence[6] := USINT#4;
   BenchUut5.processSequence[7] := USINT#3;
   BenchUut5.processSequence[8] := USINT#5;
   TraceIn_processLength[54] := BenchUut5.processLength;
   TraceIn_sensor1[54] := BenchUut5.sensor1;
   TraceIn_sensor2[54] := BenchUut5.sensor2;
   TraceIn_sensor3[54] := BenchUut5.sensor3;
   TraceIn_sensor4[54] := BenchUut5.sensor4;
   TraceIn_sensor5[54] := BenchUut5.sensor5;
   TraceIn_station1Start[54] := BenchUut5.station1Start;
   TraceIn_station2Complete[54] := BenchUut5.station2Complete;
   TraceIn_station3Complete[54] := BenchUut5.station3Complete;
   TraceIn_station4Complete[54] := BenchUut5.station4Complete;
   TraceIn_processSequence_1[54] := BenchUut5.processSequence[1];
   TraceIn_processSequence_2[54] := BenchUut5.processSequence[2];
   TraceIn_processSequence_3[54] := BenchUut5.processSequence[3];
   TraceIn_processSequence_4[54] := BenchUut5.processSequence[4];
   TraceIn_processSequence_5[54] := BenchUut5.processSequence[5];
   TraceIn_processSequence_6[54] := BenchUut5.processSequence[6];
   TraceIn_processSequence_7[54] := BenchUut5.processSequence[7];
   TraceIn_processSequence_8[54] := BenchUut5.processSequence[8];
   BenchUut5();
   TraceOut_conveyorLeft[54] := BenchUut5.conveyorLeft;
   TraceOut_conveyorRight[54] := BenchUut5.conveyorRight;
   BenchCalls := BenchCalls + 1;
 55:
   BenchUut5.processLength := USINT#8;
   BenchUut5.sensor1 := FALSE;
   BenchUut5.sensor2 := FALSE;
   BenchUut5.sensor3 := FALSE;
   BenchUut5.sensor4 := FALSE;
   BenchUut5.sensor5 := FALSE;
   BenchUut5.station1Start := FALSE;
   BenchUut5.station2Complete := FALSE;
   BenchUut5.station3Complete := FALSE;
   BenchUut5.station4Complete := FALSE;
   BenchUut5.processSequence[1] := USINT#2;
   BenchUut5.processSequence[2] := USINT#3;
   BenchUut5.processSequence[3] := USINT#4;
   BenchUut5.processSequence[4] := USINT#3;
   BenchUut5.processSequence[5] := USINT#2;
   BenchUut5.processSequence[6] := USINT#4;
   BenchUut5.processSequence[7] := USINT#3;
   BenchUut5.processSequence[8] := USINT#5;
   TraceIn_processLength[55] := BenchUut5.processLength;
   TraceIn_sensor1[55] := BenchUut5.sensor1;
   TraceIn_sensor2[55] := BenchUut5.sensor2;
   TraceIn_sensor3[55] := BenchUut5.sensor3;
   TraceIn_sensor4[55] := BenchUut5.sensor4;
   TraceIn_sensor5[55] := BenchUut5.sensor5;
   TraceIn_station1Start[55] := BenchUut5.station1Start;
   TraceIn_station2Complete[55] := BenchUut5.station2Complete;
   TraceIn_station3Complete[55] := BenchUut5.station3Complete;
   TraceIn_station4Complete[55] := BenchUut5.station4Complete;
   TraceIn_processSequence_1[55] := BenchUut5.processSequence[1];
   TraceIn_processSequence_2[55] := BenchUut5.processSequence[2];
   TraceIn_processSequence_3[55] := BenchUut5.processSequence[3];
   TraceIn_processSequence_4[55] := BenchUut5.processSequence[4];
   TraceIn_processSequence_5[55] := BenchUut5.processSequence[5];
   TraceIn_processSequence_6[55] := BenchUut5.processSequence[6];
   TraceIn_processSequence_7[55] := BenchUut5.processSequence[7];
   TraceIn_processSequence_8[55] := BenchUut5.processSequence[8];
   BenchUut5();
   TraceOut_conveyorLeft[55] := BenchUut5.conveyorLeft;
   TraceOut_conveyorRight[55] := BenchUut5.conveyorRight;
   BenchCalls := BenchCalls + 1;
 56:
   BenchUut5.processLength := USINT#8;
   BenchUut5.sensor1 := FALSE;
   BenchUut5.sensor2 := FALSE;
   BenchUut5.sensor3 := TRUE;
   BenchUut5.sensor4 := FALSE;
   BenchUut5.sensor5 := FALSE;
   BenchUut5.station1Start := FALSE;
   BenchUut5.station2Complete := FALSE;
   BenchUut5.station3Complete := FALSE;
   BenchUut5.station4Complete := FALSE;
   BenchUut5.processSequence[1] := USINT#2;
   BenchUut5.processSequence[2] := USINT#3;
   BenchUut5.processSequence[3] := USINT#4;
   BenchUut5.processSequence[4] := USINT#3;
   BenchUut5.processSequence[5] := USINT#2;
   BenchUut5.processSequence[6] := USINT#4;
   BenchUut5.processSequence[7] := USINT#3;
   BenchUut5.processSequence[8] := USINT#5;
   TraceIn_processLength[56] := BenchUut5.processLength;
   TraceIn_sensor1[56] := BenchUut5.sensor1;
   TraceIn_sensor2[56] := BenchUut5.sensor2;
   TraceIn_sensor3[56] := BenchUut5.sensor3;
   TraceIn_sensor4[56] := BenchUut5.sensor4;
   TraceIn_sensor5[56] := BenchUut5.sensor5;
   TraceIn_station1Start[56] := BenchUut5.station1Start;
   TraceIn_station2Complete[56] := BenchUut5.station2Complete;
   TraceIn_station3Complete[56] := BenchUut5.station3Complete;
   TraceIn_station4Complete[56] := BenchUut5.station4Complete;
   TraceIn_processSequence_1[56] := BenchUut5.processSequence[1];
   TraceIn_processSequence_2[56] := BenchUut5.processSequence[2];
   TraceIn_processSequence_3[56] := BenchUut5.processSequence[3];
   TraceIn_processSequence_4[56] := BenchUut5.processSequence[4];
   TraceIn_processSequence_5[56] := BenchUut5.processSequence[5];
   TraceIn_processSequence_6[56] := BenchUut5.processSequence[6];
   TraceIn_processSequence_7[56] := BenchUut5.processSequence[7];
   TraceIn_processSequence_8[56] := BenchUut5.processSequence[8];
   BenchUut5();
   TraceOut_conveyorLeft[56] := BenchUut5.conveyorLeft;
   TraceOut_conveyorRight[56] := BenchUut5.conveyorRight;
   BenchCalls := BenchCalls + 1;
 57:
   BenchUut5.processLength := USINT#8;
   BenchUut5.sensor1 := FALSE;
   BenchUut5.sensor2 := FALSE;
   BenchUut5.sensor3 := TRUE;
   BenchUut5.sensor4 := FALSE;
   BenchUut5.sensor5 := FALSE;
   BenchUut5.station1Start := FALSE;
   BenchUut5.station2Complete := FALSE;
   BenchUut5.station3Complete := FALSE;
   BenchUut5.station4Complete := FALSE;
   BenchUut5.processSequence[1] := USINT#2;
   BenchUut5.processSequence[2] := USINT#3;
   BenchUut5.processSequence[3] := USINT#4;
   BenchUut5.processSequence[4] := USINT#3;
   BenchUut5.processSequence[5] := USINT#2;
   BenchUut5.processSequence[6] := USINT#4;
   BenchUut5.processSequence[7] := USINT#3;
   BenchUut5.processSequence[8] := USINT#5;
   TraceIn_processLength[57] := BenchUut5.processLength;
   TraceIn_sensor1[57] := BenchUut5.sensor1;
   TraceIn_sensor2[57] := BenchUut5.sensor2;
   TraceIn_sensor3[57] := BenchUut5.sensor3;
   TraceIn_sensor4[57] := BenchUut5.sensor4;
   TraceIn_sensor5[57] := BenchUut5.sensor5;
   TraceIn_station1Start[57] := BenchUut5.station1Start;
   TraceIn_station2Complete[57] := BenchUut5.station2Complete;
   TraceIn_station3Complete[57] := BenchUut5.station3Complete;
   TraceIn_station4Complete[57] := BenchUut5.station4Complete;
   TraceIn_processSequence_1[57] := BenchUut5.processSequence[1];
   TraceIn_processSequence_2[57] := BenchUut5.processSequence[2];
   TraceIn_processSequence_3[57] := BenchUut5.processSequence[3];
   TraceIn_processSequence_4[57] := BenchUut5.processSequence[4];
   TraceIn_processSequence_5[57] := BenchUut5.processSequence[5];
   TraceIn_processSequence_6[57] := BenchUut5.processSequence[6];
   TraceIn_processSequence_7[57] := BenchUut5.processSequence[7];
   TraceIn_processSequence_8[57] := BenchUut5.processSequence[8];
   BenchUut5();
   TraceOut_conveyorLeft[57] := BenchUut5.conveyorLeft;
   TraceOut_conveyorRight[57] := BenchUut5.conveyorRight;
   BenchCalls := BenchCalls + 1;
 58:
   BenchUut5.processLength := USINT#8;
   BenchUut5.sensor1 := FALSE;
   BenchUut5.sensor2 := FALSE;
   BenchUut5.sensor3 := TRUE;
   BenchUut5.sensor4 := FALSE;
   BenchUut5.sensor5 := FALSE;
   BenchUut5.station1Start := FALSE;
   BenchUut5.station2Complete := FALSE;
   BenchUut5.station3Complete := FALSE;
   BenchUut5.station4Complete := FALSE;
   BenchUut5.processSequence[1] := USINT#2;
   BenchUut5.processSequence[2] := USINT#3;
   BenchUut5.processSequence[3] := USINT#4;
   BenchUut5.processSequence[4] := USINT#3;
   BenchUut5.processSequence[5] := USINT#2;
   BenchUut5.processSequence[6] := USINT#4;
   BenchUut5.processSequence[7] := USINT#3;
   BenchUut5.processSequence[8] := USINT#5;
   TraceIn_processLength[58] := BenchUut5.processLength;
   TraceIn_sensor1[58] := BenchUut5.sensor1;
   TraceIn_sensor2[58] := BenchUut5.sensor2;
   TraceIn_sensor3[58] := BenchUut5.sensor3;
   TraceIn_sensor4[58] := BenchUut5.sensor4;
   TraceIn_sensor5[58] := BenchUut5.sensor5;
   TraceIn_station1Start[58] := BenchUut5.station1Start;
   TraceIn_station2Complete[58] := BenchUut5.station2Complete;
   TraceIn_station3Complete[58] := BenchUut5.station3Complete;
   TraceIn_station4Complete[58] := BenchUut5.station4Complete;
   TraceIn_processSequence_1[58] := BenchUut5.processSequence[1];
   TraceIn_processSequence_2[58] := BenchUut5.processSequence[2];
   TraceIn_processSequence_3[58] := BenchUut5.processSequence[3];
   TraceIn_processSequence_4[58] := BenchUut5.processSequence[4];
   TraceIn_processSequence_5[58] := BenchUut5.processSequence[5];
   TraceIn_processSequence_6[58] := BenchUut5.processSequence[6];
   TraceIn_processSequence_7[58] := BenchUut5.processSequence[7];
   TraceIn_processSequence_8[58] := BenchUut5.processSequence[8];
   BenchUut5();
   TraceOut_conveyorLeft[58] := BenchUut5.conveyorLeft;
   TraceOut_conveyorRight[58] := BenchUut5.conveyorRight;
   BenchCalls := BenchCalls + 1;
 59:
   BenchUut5.processLength := USINT#8;
   BenchUut5.sensor1 := FALSE;
   BenchUut5.sensor2 := FALSE;
   BenchUut5.sensor3 := TRUE;
   BenchUut5.sensor4 := FALSE;
   BenchUut5.sensor5 := FALSE;
   BenchUut5.station1Start := FALSE;
   BenchUut5.station2Complete := FALSE;
   BenchUut5.station3Complete := TRUE;
   BenchUut5.station4Complete := FALSE;
   BenchUut5.processSequence[1] := USINT#2;
   BenchUut5.processSequence[2] := USINT#3;
   BenchUut5.processSequence[3] := USINT#4;
   BenchUut5.processSequence[4] := USINT#3;
   BenchUut5.processSequence[5] := USINT#2;
   BenchUut5.processSequence[6] := USINT#4;
   BenchUut5.processSequence[7] := USINT#3;
   BenchUut5.processSequence[8] := USINT#5;
   TraceIn_processLength[59] := BenchUut5.processLength;
   TraceIn_sensor1[59] := BenchUut5.sensor1;
   TraceIn_sensor2[59] := BenchUut5.sensor2;
   TraceIn_sensor3[59] := BenchUut5.sensor3;
   TraceIn_sensor4[59] := BenchUut5.sensor4;
   TraceIn_sensor5[59] := BenchUut5.sensor5;
   TraceIn_station1Start[59] := BenchUut5.station1Start;
   TraceIn_station2Complete[59] := BenchUut5.station2Complete;
   TraceIn_station3Complete[59] := BenchUut5.station3Complete;
   TraceIn_station4Complete[59] := BenchUut5.station4Complete;
   TraceIn_processSequence_1[59] := BenchUut5.processSequence[1];
   TraceIn_processSequence_2[59] := BenchUut5.processSequence[2];
   TraceIn_processSequence_3[59] := BenchUut5.processSequence[3];
   TraceIn_processSequence_4[59] := BenchUut5.processSequence[4];
   TraceIn_processSequence_5[59] := BenchUut5.processSequence[5];
   TraceIn_processSequence_6[59] := BenchUut5.processSequence[6];
   TraceIn_processSequence_7[59] := BenchUut5.processSequence[7];
   TraceIn_processSequence_8[59] := BenchUut5.processSequence[8];
   BenchUut5();
   TraceOut_conveyorLeft[59] := BenchUut5.conveyorLeft;
   TraceOut_conveyorRight[59] := BenchUut5.conveyorRight;
   BenchCalls := BenchCalls + 1;
 60:
   BenchUut5.processLength := USINT#8;
   BenchUut5.sensor1 := FALSE;
   BenchUut5.sensor2 := FALSE;
   BenchUut5.sensor3 := FALSE;
   BenchUut5.sensor4 := FALSE;
   BenchUut5.sensor5 := FALSE;
   BenchUut5.station1Start := FALSE;
   BenchUut5.station2Complete := FALSE;
   BenchUut5.station3Complete := FALSE;
   BenchUut5.station4Complete := FALSE;
   BenchUut5.processSequence[1] := USINT#2;
   BenchUut5.processSequence[2] := USINT#3;
   BenchUut5.processSequence[3] := USINT#4;
   BenchUut5.processSequence[4] := USINT#3;
   BenchUut5.processSequence[5] := USINT#2;
   BenchUut5.processSequence[6] := USINT#4;
   BenchUut5.processSequence[7] := USINT#3;
   BenchUut5.processSequence[8] := USINT#5;
   TraceIn_processLength[60] := BenchUut5.processLength;
   TraceIn_sensor1[60] := BenchUut5.sensor1;
   TraceIn_sensor2[60] := BenchUut5.sensor2;
   TraceIn_sensor3[60] := BenchUut5.sensor3;
   TraceIn_sensor4[60] := BenchUut5.sensor4;
   TraceIn_sensor5[60] := BenchUut5.sensor5;
   TraceIn_station1Start[60] := BenchUut5.station1Start;
   TraceIn_station2Complete[60] := BenchUut5.station2Complete;
   TraceIn_station3Complete[60] := BenchUut5.station3Complete;
   TraceIn_station4Complete[60] := BenchUut5.station4Complete;
   TraceIn_processSequence_1[60] := BenchUut5.processSequence[1];
   TraceIn_processSequence_2[60] := BenchUut5.processSequence[2];
   TraceIn_processSequence_3[60] := BenchUut5.processSequence[3];
   TraceIn_processSequence_4[60] := BenchUut5.processSequence[4];
   TraceIn_processSequence_5[60] := BenchUut5.processSequence[5];
   TraceIn_processSequence_6[60] := BenchUut5.processSequence[6];
   TraceIn_processSequence_7[60] := BenchUut5.processSequence[7];
   TraceIn_processSequence_8[60] := BenchUut5.processSequence[8];
   BenchUut5();
   TraceOut_conveyorLeft[60] := BenchUut5.conveyorLeft;
   TraceOut_conveyorRight[60] := BenchUut5.conveyorRight;
   BenchCalls := BenchCalls + 1;
 61:
   BenchUut5.processLength := USINT#8;
   BenchUut5.sensor1 := FALSE;
   BenchUut5.sensor2 := FALSE;
   BenchUut5.sensor3 := FALSE;
   BenchUut5.sensor4 := FALSE;
   BenchUut5.sensor5 := FALSE;
   BenchUut5.station1Start := FALSE;
   BenchUut5.station2Complete := FALSE;
   BenchUut5.station3Complete := FALSE;
   BenchUut5.station4Complete := FALSE;
   BenchUut5.processSequence[1] := USINT#2;
   BenchUut5.processSequence[2] := USINT#3;
   BenchUut5.processSequence[3] := USINT#4;
   BenchUut5.processSequence[4] := USINT#3;
   BenchUut5.processSequence[5] := USINT#2;
   BenchUut5.processSequence[6] := USINT#4;
   BenchUut5.processSequence[7] := USINT#3;
   BenchUut5.processSequence[8] := USINT#5;
   TraceIn_processLength[61] := BenchUut5.processLength;
   TraceIn_sensor1[61] := BenchUut5.sensor1;
   TraceIn_sensor2[61] := BenchUut5.sensor2;
   TraceIn_sensor3[61] := BenchUut5.sensor3;
   TraceIn_sensor4[61] := BenchUut5.sensor4;
   TraceIn_sensor5[61] := BenchUut5.sensor5;
   TraceIn_station1Start[61] := BenchUut5.station1Start;
   TraceIn_station2Complete[61] := BenchUut5.station2Complete;
   TraceIn_station3Complete[61] := BenchUut5.station3Complete;
   TraceIn_station4Complete[61] := BenchUut5.station4Complete;
   TraceIn_processSequence_1[61] := BenchUut5.processSequence[1];
   TraceIn_processSequence_2[61] := BenchUut5.processSequence[2];
   TraceIn_processSequence_3[61] := BenchUut5.processSequence[3];
   TraceIn_processSequence_4[61] := BenchUut5.processSequence[4];
   TraceIn_processSequence_5[61] := BenchUut5.processSequence[5];
   TraceIn_processSequence_6[61] := BenchUut5.processSequence[6];
   TraceIn_processSequence_7[61] := BenchUut5.processSequence[7];
   TraceIn_processSequence_8[61] := BenchUut5.processSequence[8];
   BenchUut5();
   TraceOut_conveyorLeft[61] := BenchUut5.conveyorLeft;
   TraceOut_conveyorRight[61] := BenchUut5.conveyorRight;
   BenchCalls := BenchCalls + 1;
 62:
   BenchUut5.processLength := USINT#8;
   BenchUut5.sensor1 := FALSE;
   BenchUut5.sensor2 := FALSE;
   BenchUut5.sensor3 := FALSE;
   BenchUut5.sensor4 := TRUE;
   BenchUut5.sensor5 := FALSE;
   BenchUut5.station1Start := FALSE;
   BenchUut5.station2Complete := FALSE;
   BenchUut5.station3Complete := FALSE;
   BenchUut5.station4Complete := FALSE;
   BenchUut5.processSequence[1] := USINT#2;
   BenchUut5.processSequence[2] := USINT#3;
   BenchUut5.processSequence[3] := USINT#4;
   BenchUut5.processSequence[4] := USINT#3;
   BenchUut5.processSequence[5] := USINT#2;
   BenchUut5.processSequence[6] := USINT#4;
   BenchUut5.processSequence[7] := USINT#3;
   BenchUut5.processSequence[8] := USINT#5;
   TraceIn_processLength[62] := BenchUut5.processLength;
   TraceIn_sensor1[62] := BenchUut5.sensor1;
   TraceIn_sensor2[62] := BenchUut5.sensor2;
   TraceIn_sensor3[62] := BenchUut5.sensor3;
   TraceIn_sensor4[62] := BenchUut5.sensor4;
   TraceIn_sensor5[62] := BenchUut5.sensor5;
   TraceIn_station1Start[62] := BenchUut5.station1Start;
   TraceIn_station2Complete[62] := BenchUut5.station2Complete;
   TraceIn_station3Complete[62] := BenchUut5.station3Complete;
   TraceIn_station4Complete[62] := BenchUut5.station4Complete;
   TraceIn_processSequence_1[62] := BenchUut5.processSequence[1];
   TraceIn_processSequence_2[62] := BenchUut5.processSequence[2];
   TraceIn_processSequence_3[62] := BenchUut5.processSequence[3];
   TraceIn_processSequence_4[62] := BenchUut5.processSequence[4];
   TraceIn_processSequence_5[62] := BenchUut5.processSequence[5];
   TraceIn_processSequence_6[62] := BenchUut5.processSequence[6];
   TraceIn_processSequence_7[62] := BenchUut5.processSequence[7];
   TraceIn_processSequence_8[62] := BenchUut5.processSequence[8];
   BenchUut5();
   TraceOut_conveyorLeft[62] := BenchUut5.conveyorLeft;
   TraceOut_conveyorRight[62] := BenchUut5.conveyorRight;
   BenchCalls := BenchCalls + 1;
 63:
   BenchUut5.processLength := USINT#8;
   BenchUut5.sensor1 := FALSE;
   BenchUut5.sensor2 := FALSE;
   BenchUut5.sensor3 := FALSE;
   BenchUut5.sensor4 := TRUE;
   BenchUut5.sensor5 := FALSE;
   BenchUut5.station1Start := FALSE;
   BenchUut5.station2Complete := FALSE;
   BenchUut5.station3Complete := FALSE;
   BenchUut5.station4Complete := FALSE;
   BenchUut5.processSequence[1] := USINT#2;
   BenchUut5.processSequence[2] := USINT#3;
   BenchUut5.processSequence[3] := USINT#4;
   BenchUut5.processSequence[4] := USINT#3;
   BenchUut5.processSequence[5] := USINT#2;
   BenchUut5.processSequence[6] := USINT#4;
   BenchUut5.processSequence[7] := USINT#3;
   BenchUut5.processSequence[8] := USINT#5;
   TraceIn_processLength[63] := BenchUut5.processLength;
   TraceIn_sensor1[63] := BenchUut5.sensor1;
   TraceIn_sensor2[63] := BenchUut5.sensor2;
   TraceIn_sensor3[63] := BenchUut5.sensor3;
   TraceIn_sensor4[63] := BenchUut5.sensor4;
   TraceIn_sensor5[63] := BenchUut5.sensor5;
   TraceIn_station1Start[63] := BenchUut5.station1Start;
   TraceIn_station2Complete[63] := BenchUut5.station2Complete;
   TraceIn_station3Complete[63] := BenchUut5.station3Complete;
   TraceIn_station4Complete[63] := BenchUut5.station4Complete;
   TraceIn_processSequence_1[63] := BenchUut5.processSequence[1];
   TraceIn_processSequence_2[63] := BenchUut5.processSequence[2];
   TraceIn_processSequence_3[63] := BenchUut5.processSequence[3];
   TraceIn_processSequence_4[63] := BenchUut5.processSequence[4];
   TraceIn_processSequence_5[63] := BenchUut5.processSequence[5];
   TraceIn_processSequence_6[63] := BenchUut5.processSequence[6];
   TraceIn_processSequence_7[63] := BenchUut5.processSequence[7];
   TraceIn_processSequence_8[63] := BenchUut5.processSequence[8];
   BenchUut5();
   TraceOut_conveyorLeft[63] := BenchUut5.conveyorLeft;
   TraceOut_conveyorRight[63] := BenchUut5.conveyorRight;
   BenchCalls := BenchCalls + 1;
 64:
   BenchUut5.processLength := USINT#8;
   BenchUut5.sensor1 := FALSE;
   BenchUut5.sensor2 := FALSE;
   BenchUut5.sensor3 := FALSE;
   BenchUut5.sensor4 := TRUE;
   BenchUut5.sensor5 := FALSE;
   BenchUut5.station1Start := FALSE;
   BenchUut5.station2Complete := FALSE;
   BenchUut5.station3Complete := FALSE;
   BenchUut5.station4Complete := FALSE;
   BenchUut5.processSequence[1] := USINT#2;
   BenchUut5.processSequence[2] := USINT#3;
   BenchUut5.processSequence[3] := USINT#4;
   BenchUut5.processSequence[4] := USINT#3;
   BenchUut5.processSequence[5] := USINT#2;
   BenchUut5.processSequence[6] := USINT#4;
   BenchUut5.processSequence[7] := USINT#3;
   BenchUut5.processSequence[8] := USINT#5;
   TraceIn_processLength[64] := BenchUut5.processLength;
   TraceIn_sensor1[64] := BenchUut5.sensor1;
   TraceIn_sensor2[64] := BenchUut5.sensor2;
   TraceIn_sensor3[64] := BenchUut5.sensor3;
   TraceIn_sensor4[64] := BenchUut5.sensor4;
   TraceIn_sensor5[64] := BenchUut5.sensor5;
   TraceIn_station1Start[64] := BenchUut5.station1Start;
   TraceIn_station2Complete[64] := BenchUut5.station2Complete;
   TraceIn_station3Complete[64] := BenchUut5.station3Complete;
   TraceIn_station4Complete[64] := BenchUut5.station4Complete;
   TraceIn_processSequence_1[64] := BenchUut5.processSequence[1];
   TraceIn_processSequence_2[64] := BenchUut5.processSequence[2];
   TraceIn_processSequence_3[64] := BenchUut5.processSequence[3];
   TraceIn_processSequence_4[64] := BenchUut5.processSequence[4];
   TraceIn_processSequence_5[64] := BenchUut5.processSequence[5];
   TraceIn_processSequence_6[64] := BenchUut5.processSequence[6];
   TraceIn_processSequence_7[64] := BenchUut5.processSequence[7];
   TraceIn_processSequence_8[64] := BenchUut5.processSequence[8];
   BenchUut5();
   TraceOut_conveyorLeft[64] := BenchUut5.conveyorLeft;
   TraceOut_conveyorRight[64] := BenchUut5.conveyorRight;
   BenchCalls := BenchCalls + 1;
 65:
   BenchUut5.processLength := USINT#8;
   BenchUut5.sensor1 := FALSE;
   BenchUut5.sensor2 := FALSE;
   BenchUut5.sensor3 := FALSE;
   BenchUut5.sensor4 := TRUE;
   BenchUut5.sensor5 := FALSE;
   BenchUut5.station1Start := FALSE;
   BenchUut5.station2Complete := FALSE;
   BenchUut5.station3Complete := FALSE;
   BenchUut5.station4Complete := TRUE;
   BenchUut5.processSequence[1] := USINT#2;
   BenchUut5.processSequence[2] := USINT#3;
   BenchUut5.processSequence[3] := USINT#4;
   BenchUut5.processSequence[4] := USINT#3;
   BenchUut5.processSequence[5] := USINT#2;
   BenchUut5.processSequence[6] := USINT#4;
   BenchUut5.processSequence[7] := USINT#3;
   BenchUut5.processSequence[8] := USINT#5;
   TraceIn_processLength[65] := BenchUut5.processLength;
   TraceIn_sensor1[65] := BenchUut5.sensor1;
   TraceIn_sensor2[65] := BenchUut5.sensor2;
   TraceIn_sensor3[65] := BenchUut5.sensor3;
   TraceIn_sensor4[65] := BenchUut5.sensor4;
   TraceIn_sensor5[65] := BenchUut5.sensor5;
   TraceIn_station1Start[65] := BenchUut5.station1Start;
   TraceIn_station2Complete[65] := BenchUut5.station2Complete;
   TraceIn_station3Complete[65] := BenchUut5.station3Complete;
   TraceIn_station4Complete[65] := BenchUut5.station4Complete;
   TraceIn_processSequence_1[65] := BenchUut5.processSequence[1];
   TraceIn_processSequence_2[65] := BenchUut5.processSequence[2];
   TraceIn_processSequence_3[65] := BenchUut5.processSequence[3];
   TraceIn_processSequence_4[65] := BenchUut5.processSequence[4];
   TraceIn_processSequence_5[65] := BenchUut5.processSequence[5];
   TraceIn_processSequence_6[65] := BenchUut5.processSequence[6];
   TraceIn_processSequence_7[65] := BenchUut5.processSequence[7];
   TraceIn_processSequence_8[65] := BenchUut5.processSequence[8];
   BenchUut5();
   TraceOut_conveyorLeft[65] := BenchUut5.conveyorLeft;
   TraceOut_conveyorRight[65] := BenchUut5.conveyorRight;
   BenchCalls := BenchCalls + 1;
 66:
   BenchUut5.processLength := USINT#8;
   BenchUut5.sensor1 := FALSE;
   BenchUut5.sensor2 := FALSE;
   BenchUut5.sensor3 := FALSE;
   BenchUut5.sensor4 := FALSE;
   BenchUut5.sensor5 := FALSE;
   BenchUut5.station1Start := FALSE;
   BenchUut5.station2Complete := FALSE;
   BenchUut5.station3Complete := FALSE;
   BenchUut5.station4Complete := FALSE;
   BenchUut5.processSequence[1] := USINT#2;
   BenchUut5.processSequence[2] := USINT#3;
   BenchUut5.processSequence[3] := USINT#4;
   BenchUut5.processSequence[4] := USINT#3;
   BenchUut5.processSequence[5] := USINT#2;
   BenchUut5.processSequence[6] := USINT#4;
   BenchUut5.processSequence[7] := USINT#3;
   BenchUut5.processSequence[8] := USINT#5;
   TraceIn_processLength[66] := BenchUut5.processLength;
   TraceIn_sensor1[66] := BenchUut5.sensor1;
   TraceIn_sensor2[66] := BenchUut5.sensor2;
   TraceIn_sensor3[66] := BenchUut5.sensor3;
   TraceIn_sensor4[66] := BenchUut5.sensor4;
   TraceIn_sensor5[66] := BenchUut5.sensor5;
   TraceIn_station1Start[66] := BenchUut5.station1Start;
   TraceIn_station2Complete[66] := BenchUut5.station2Complete;
   TraceIn_station3Complete[66] := BenchUut5.station3Complete;
   TraceIn_station4Complete[66] := BenchUut5.station4Complete;
   TraceIn_processSequence_1[66] := BenchUut5.processSequence[1];
   TraceIn_processSequence_2[66] := BenchUut5.processSequence[2];
   TraceIn_processSequence_3[66] := BenchUut5.processSequence[3];
   TraceIn_processSequence_4[66] := BenchUut5.processSequence[4];
   TraceIn_processSequence_5[66] := BenchUut5.processSequence[5];
   TraceIn_processSequence_6[66] := BenchUut5.processSequence[6];
   TraceIn_processSequence_7[66] := BenchUut5.processSequence[7];
   TraceIn_processSequence_8[66] := BenchUut5.processSequence[8];
   BenchUut5();
   TraceOut_conveyorLeft[66] := BenchUut5.conveyorLeft;
   TraceOut_conveyorRight[66] := BenchUut5.conveyorRight;
   BenchCalls := BenchCalls + 1;
 67:
   BenchUut5.processLength := USINT#8;
   BenchUut5.sensor1 := FALSE;
   BenchUut5.sensor2 := FALSE;
   BenchUut5.sensor3 := FALSE;
   BenchUut5.sensor4 := FALSE;
   BenchUut5.sensor5 := FALSE;
   BenchUut5.station1Start := FALSE;
   BenchUut5.station2Complete := FALSE;
   BenchUut5.station3Complete := FALSE;
   BenchUut5.station4Complete := FALSE;
   BenchUut5.processSequence[1] := USINT#2;
   BenchUut5.processSequence[2] := USINT#3;
   BenchUut5.processSequence[3] := USINT#4;
   BenchUut5.processSequence[4] := USINT#3;
   BenchUut5.processSequence[5] := USINT#2;
   BenchUut5.processSequence[6] := USINT#4;
   BenchUut5.processSequence[7] := USINT#3;
   BenchUut5.processSequence[8] := USINT#5;
   TraceIn_processLength[67] := BenchUut5.processLength;
   TraceIn_sensor1[67] := BenchUut5.sensor1;
   TraceIn_sensor2[67] := BenchUut5.sensor2;
   TraceIn_sensor3[67] := BenchUut5.sensor3;
   TraceIn_sensor4[67] := BenchUut5.sensor4;
   TraceIn_sensor5[67] := BenchUut5.sensor5;
   TraceIn_station1Start[67] := BenchUut5.station1Start;
   TraceIn_station2Complete[67] := BenchUut5.station2Complete;
   TraceIn_station3Complete[67] := BenchUut5.station3Complete;
   TraceIn_station4Complete[67] := BenchUut5.station4Complete;
   TraceIn_processSequence_1[67] := BenchUut5.processSequence[1];
   TraceIn_processSequence_2[67] := BenchUut5.processSequence[2];
   TraceIn_processSequence_3[67] := BenchUut5.processSequence[3];
   TraceIn_processSequence_4[67] := BenchUut5.processSequence[4];
   TraceIn_processSequence_5[67] := BenchUut5.processSequence[5];
   TraceIn_processSequence_6[67] := BenchUut5.processSequence[6];
   TraceIn_processSequence_7[67] := BenchUut5.processSequence[7];
   TraceIn_processSequence_8[67] := BenchUut5.processSequence[8];
   BenchUut5();
   TraceOut_conveyorLeft[67] := BenchUut5.conveyorLeft;
   TraceOut_conveyorRight[67] := BenchUut5.conveyorRight;
   BenchCalls := BenchCalls + 1;
 68:
   BenchUut5.processLength := USINT#8;
   BenchUut5.sensor1 := FALSE;
   BenchUut5.sensor2 := FALSE;
   BenchUut5.sensor3 := TRUE;
   BenchUut5.sensor4 := FALSE;
   BenchUut5.sensor5 := FALSE;
   BenchUut5.station1Start := FALSE;
   BenchUut5.station2Complete := FALSE;
   BenchUut5.station3Complete := FALSE;
   BenchUut5.station4Complete := FALSE;
   BenchUut5.processSequence[1] := USINT#2;
   BenchUut5.processSequence[2] := USINT#3;
   BenchUut5.processSequence[3] := USINT#4;
   BenchUut5.processSequence[4] := USINT#3;
   BenchUut5.processSequence[5] := USINT#2;
   BenchUut5.processSequence[6] := USINT#4;
   BenchUut5.processSequence[7] := USINT#3;
   BenchUut5.processSequence[8] := USINT#5;
   TraceIn_processLength[68] := BenchUut5.processLength;
   TraceIn_sensor1[68] := BenchUut5.sensor1;
   TraceIn_sensor2[68] := BenchUut5.sensor2;
   TraceIn_sensor3[68] := BenchUut5.sensor3;
   TraceIn_sensor4[68] := BenchUut5.sensor4;
   TraceIn_sensor5[68] := BenchUut5.sensor5;
   TraceIn_station1Start[68] := BenchUut5.station1Start;
   TraceIn_station2Complete[68] := BenchUut5.station2Complete;
   TraceIn_station3Complete[68] := BenchUut5.station3Complete;
   TraceIn_station4Complete[68] := BenchUut5.station4Complete;
   TraceIn_processSequence_1[68] := BenchUut5.processSequence[1];
   TraceIn_processSequence_2[68] := BenchUut5.processSequence[2];
   TraceIn_processSequence_3[68] := BenchUut5.processSequence[3];
   TraceIn_processSequence_4[68] := BenchUut5.processSequence[4];
   TraceIn_processSequence_5[68] := BenchUut5.processSequence[5];
   TraceIn_processSequence_6[68] := BenchUut5.processSequence[6];
   TraceIn_processSequence_7[68] := BenchUut5.processSequence[7];
   TraceIn_processSequence_8[68] := BenchUut5.processSequence[8];
   BenchUut5();
   TraceOut_conveyorLeft[68] := BenchUut5.conveyorLeft;
   TraceOut_conveyorRight[68] := BenchUut5.conveyorRight;
   BenchCalls := BenchCalls + 1;
 69:
   BenchUut5.processLength := USINT#8;
   BenchUut5.sensor1 := FALSE;
   BenchUut5.sensor2 := FALSE;
   BenchUut5.sensor3 := TRUE;
   BenchUut5.sensor4 := FALSE;
   BenchUut5.sensor5 := FALSE;
   BenchUut5.station1Start := FALSE;
   BenchUut5.station2Complete := FALSE;
   BenchUut5.station3Complete := FALSE;
   BenchUut5.station4Complete := FALSE;
   BenchUut5.processSequence[1] := USINT#2;
   BenchUut5.processSequence[2] := USINT#3;
   BenchUut5.processSequence[3] := USINT#4;
   BenchUut5.processSequence[4] := USINT#3;
   BenchUut5.processSequence[5] := USINT#2;
   BenchUut5.processSequence[6] := USINT#4;
   BenchUut5.processSequence[7] := USINT#3;
   BenchUut5.processSequence[8] := USINT#5;
   TraceIn_processLength[69] := BenchUut5.processLength;
   TraceIn_sensor1[69] := BenchUut5.sensor1;
   TraceIn_sensor2[69] := BenchUut5.sensor2;
   TraceIn_sensor3[69] := BenchUut5.sensor3;
   TraceIn_sensor4[69] := BenchUut5.sensor4;
   TraceIn_sensor5[69] := BenchUut5.sensor5;
   TraceIn_station1Start[69] := BenchUut5.station1Start;
   TraceIn_station2Complete[69] := BenchUut5.station2Complete;
   TraceIn_station3Complete[69] := BenchUut5.station3Complete;
   TraceIn_station4Complete[69] := BenchUut5.station4Complete;
   TraceIn_processSequence_1[69] := BenchUut5.processSequence[1];
   TraceIn_processSequence_2[69] := BenchUut5.processSequence[2];
   TraceIn_processSequence_3[69] := BenchUut5.processSequence[3];
   TraceIn_processSequence_4[69] := BenchUut5.processSequence[4];
   TraceIn_processSequence_5[69] := BenchUut5.processSequence[5];
   TraceIn_processSequence_6[69] := BenchUut5.processSequence[6];
   TraceIn_processSequence_7[69] := BenchUut5.processSequence[7];
   TraceIn_processSequence_8[69] := BenchUut5.processSequence[8];
   BenchUut5();
   TraceOut_conveyorLeft[69] := BenchUut5.conveyorLeft;
   TraceOut_conveyorRight[69] := BenchUut5.conveyorRight;
   BenchCalls := BenchCalls + 1;
 70:
   BenchUut5.processLength := USINT#8;
   BenchUut5.sensor1 := FALSE;
   BenchUut5.sensor2 := FALSE;
   BenchUut5.sensor3 := TRUE;
   BenchUut5.sensor4 := FALSE;
   BenchUut5.sensor5 := FALSE;
   BenchUut5.station1Start := FALSE;
   BenchUut5.station2Complete := FALSE;
   BenchUut5.station3Complete := FALSE;
   BenchUut5.station4Complete := FALSE;
   BenchUut5.processSequence[1] := USINT#2;
   BenchUut5.processSequence[2] := USINT#3;
   BenchUut5.processSequence[3] := USINT#4;
   BenchUut5.processSequence[4] := USINT#3;
   BenchUut5.processSequence[5] := USINT#2;
   BenchUut5.processSequence[6] := USINT#4;
   BenchUut5.processSequence[7] := USINT#3;
   BenchUut5.processSequence[8] := USINT#5;
   TraceIn_processLength[70] := BenchUut5.processLength;
   TraceIn_sensor1[70] := BenchUut5.sensor1;
   TraceIn_sensor2[70] := BenchUut5.sensor2;
   TraceIn_sensor3[70] := BenchUut5.sensor3;
   TraceIn_sensor4[70] := BenchUut5.sensor4;
   TraceIn_sensor5[70] := BenchUut5.sensor5;
   TraceIn_station1Start[70] := BenchUut5.station1Start;
   TraceIn_station2Complete[70] := BenchUut5.station2Complete;
   TraceIn_station3Complete[70] := BenchUut5.station3Complete;
   TraceIn_station4Complete[70] := BenchUut5.station4Complete;
   TraceIn_processSequence_1[70] := BenchUut5.processSequence[1];
   TraceIn_processSequence_2[70] := BenchUut5.processSequence[2];
   TraceIn_processSequence_3[70] := BenchUut5.processSequence[3];
   TraceIn_processSequence_4[70] := BenchUut5.processSequence[4];
   TraceIn_processSequence_5[70] := BenchUut5.processSequence[5];
   TraceIn_processSequence_6[70] := BenchUut5.processSequence[6];
   TraceIn_processSequence_7[70] := BenchUut5.processSequence[7];
   TraceIn_processSequence_8[70] := BenchUut5.processSequence[8];
   BenchUut5();
   TraceOut_conveyorLeft[70] := BenchUut5.conveyorLeft;
   TraceOut_conveyorRight[70] := BenchUut5.conveyorRight;
   BenchCalls := BenchCalls + 1;
 71:
   BenchUut5.processLength := USINT#8;
   BenchUut5.sensor1 := FALSE;
   BenchUut5.sensor2 := FALSE;
   BenchUut5.sensor3 := TRUE;
   BenchUut5.sensor4 := FALSE;
   BenchUut5.sensor5 := FALSE;
   BenchUut5.station1Start := FALSE;
   BenchUut5.station2Complete := FALSE;
   BenchUut5.station3Complete := TRUE;
   BenchUut5.station4Complete := FALSE;
   BenchUut5.processSequence[1] := USINT#2;
   BenchUut5.processSequence[2] := USINT#3;
   BenchUut5.processSequence[3] := USINT#4;
   BenchUut5.processSequence[4] := USINT#3;
   BenchUut5.processSequence[5] := USINT#2;
   BenchUut5.processSequence[6] := USINT#4;
   BenchUut5.processSequence[7] := USINT#3;
   BenchUut5.processSequence[8] := USINT#5;
   TraceIn_processLength[71] := BenchUut5.processLength;
   TraceIn_sensor1[71] := BenchUut5.sensor1;
   TraceIn_sensor2[71] := BenchUut5.sensor2;
   TraceIn_sensor3[71] := BenchUut5.sensor3;
   TraceIn_sensor4[71] := BenchUut5.sensor4;
   TraceIn_sensor5[71] := BenchUut5.sensor5;
   TraceIn_station1Start[71] := BenchUut5.station1Start;
   TraceIn_station2Complete[71] := BenchUut5.station2Complete;
   TraceIn_station3Complete[71] := BenchUut5.station3Complete;
   TraceIn_station4Complete[71] := BenchUut5.station4Complete;
   TraceIn_processSequence_1[71] := BenchUut5.processSequence[1];
   TraceIn_processSequence_2[71] := BenchUut5.processSequence[2];
   TraceIn_processSequence_3[71] := BenchUut5.processSequence[3];
   TraceIn_processSequence_4[71] := BenchUut5.processSequence[4];
   TraceIn_processSequence_5[71] := BenchUut5.processSequence[5];
   TraceIn_processSequence_6[71] := BenchUut5.processSequence[6];
   TraceIn_processSequence_7[71] := BenchUut5.processSequence[7];
   TraceIn_processSequence_8[71] := BenchUut5.processSequence[8];
   BenchUut5();
   TraceOut_conveyorLeft[71] := BenchUut5.conveyorLeft;
   TraceOut_conveyorRight[71] := BenchUut5.conveyorRight;
   BenchCalls := BenchCalls + 1;
 72:
   BenchUut5.processLength := USINT#8;
   BenchUut5.sensor1 := FALSE;
   BenchUut5.sensor2 := FALSE;
   BenchUut5.sensor3 := FALSE;
   BenchUut5.sensor4 := FALSE;
   BenchUut5.sensor5 := FALSE;
   BenchUut5.station1Start := FALSE;
   BenchUut5.station2Complete := FALSE;
   BenchUut5.station3Complete := FALSE;
   BenchUut5.station4Complete := FALSE;
   BenchUut5.processSequence[1] := USINT#2;
   BenchUut5.processSequence[2] := USINT#3;
   BenchUut5.processSequence[3] := USINT#4;
   BenchUut5.processSequence[4] := USINT#3;
   BenchUut5.processSequence[5] := USINT#2;
   BenchUut5.processSequence[6] := USINT#4;
   BenchUut5.processSequence[7] := USINT#3;
   BenchUut5.processSequence[8] := USINT#5;
   TraceIn_processLength[72] := BenchUut5.processLength;
   TraceIn_sensor1[72] := BenchUut5.sensor1;
   TraceIn_sensor2[72] := BenchUut5.sensor2;
   TraceIn_sensor3[72] := BenchUut5.sensor3;
   TraceIn_sensor4[72] := BenchUut5.sensor4;
   TraceIn_sensor5[72] := BenchUut5.sensor5;
   TraceIn_station1Start[72] := BenchUut5.station1Start;
   TraceIn_station2Complete[72] := BenchUut5.station2Complete;
   TraceIn_station3Complete[72] := BenchUut5.station3Complete;
   TraceIn_station4Complete[72] := BenchUut5.station4Complete;
   TraceIn_processSequence_1[72] := BenchUut5.processSequence[1];
   TraceIn_processSequence_2[72] := BenchUut5.processSequence[2];
   TraceIn_processSequence_3[72] := BenchUut5.processSequence[3];
   TraceIn_processSequence_4[72] := BenchUut5.processSequence[4];
   TraceIn_processSequence_5[72] := BenchUut5.processSequence[5];
   TraceIn_processSequence_6[72] := BenchUut5.processSequence[6];
   TraceIn_processSequence_7[72] := BenchUut5.processSequence[7];
   TraceIn_processSequence_8[72] := BenchUut5.processSequence[8];
   BenchUut5();
   TraceOut_conveyorLeft[72] := BenchUut5.conveyorLeft;
   TraceOut_conveyorRight[72] := BenchUut5.conveyorRight;
   BenchCalls := BenchCalls + 1;
 73:
   BenchUut5.processLength := USINT#8;
   BenchUut5.sensor1 := FALSE;
   BenchUut5.sensor2 := FALSE;
   BenchUut5.sensor3 := FALSE;
   BenchUut5.sensor4 := FALSE;
   BenchUut5.sensor5 := FALSE;
   BenchUut5.station1Start := FALSE;
   BenchUut5.station2Complete := FALSE;
   BenchUut5.station3Complete := FALSE;
   BenchUut5.station4Complete := FALSE;
   BenchUut5.processSequence[1] := USINT#2;
   BenchUut5.processSequence[2] := USINT#3;
   BenchUut5.processSequence[3] := USINT#4;
   BenchUut5.processSequence[4] := USINT#3;
   BenchUut5.processSequence[5] := USINT#2;
   BenchUut5.processSequence[6] := USINT#4;
   BenchUut5.processSequence[7] := USINT#3;
   BenchUut5.processSequence[8] := USINT#5;
   TraceIn_processLength[73] := BenchUut5.processLength;
   TraceIn_sensor1[73] := BenchUut5.sensor1;
   TraceIn_sensor2[73] := BenchUut5.sensor2;
   TraceIn_sensor3[73] := BenchUut5.sensor3;
   TraceIn_sensor4[73] := BenchUut5.sensor4;
   TraceIn_sensor5[73] := BenchUut5.sensor5;
   TraceIn_station1Start[73] := BenchUut5.station1Start;
   TraceIn_station2Complete[73] := BenchUut5.station2Complete;
   TraceIn_station3Complete[73] := BenchUut5.station3Complete;
   TraceIn_station4Complete[73] := BenchUut5.station4Complete;
   TraceIn_processSequence_1[73] := BenchUut5.processSequence[1];
   TraceIn_processSequence_2[73] := BenchUut5.processSequence[2];
   TraceIn_processSequence_3[73] := BenchUut5.processSequence[3];
   TraceIn_processSequence_4[73] := BenchUut5.processSequence[4];
   TraceIn_processSequence_5[73] := BenchUut5.processSequence[5];
   TraceIn_processSequence_6[73] := BenchUut5.processSequence[6];
   TraceIn_processSequence_7[73] := BenchUut5.processSequence[7];
   TraceIn_processSequence_8[73] := BenchUut5.processSequence[8];
   BenchUut5();
   TraceOut_conveyorLeft[73] := BenchUut5.conveyorLeft;
   TraceOut_conveyorRight[73] := BenchUut5.conveyorRight;
   BenchCalls := BenchCalls + 1;
 74:
   BenchUut5.processLength := USINT#8;
   BenchUut5.sensor1 := FALSE;
   BenchUut5.sensor2 := TRUE;
   BenchUut5.sensor3 := FALSE;
   BenchUut5.sensor4 := FALSE;
   BenchUut5.sensor5 := FALSE;
   BenchUut5.station1Start := FALSE;
   BenchUut5.station2Complete := FALSE;
   BenchUut5.station3Complete := FALSE;
   BenchUut5.station4Complete := FALSE;
   BenchUut5.processSequence[1] := USINT#2;
   BenchUut5.processSequence[2] := USINT#3;
   BenchUut5.processSequence[3] := USINT#4;
   BenchUut5.processSequence[4] := USINT#3;
   BenchUut5.processSequence[5] := USINT#2;
   BenchUut5.processSequence[6] := USINT#4;
   BenchUut5.processSequence[7] := USINT#3;
   BenchUut5.processSequence[8] := USINT#5;
   TraceIn_processLength[74] := BenchUut5.processLength;
   TraceIn_sensor1[74] := BenchUut5.sensor1;
   TraceIn_sensor2[74] := BenchUut5.sensor2;
   TraceIn_sensor3[74] := BenchUut5.sensor3;
   TraceIn_sensor4[74] := BenchUut5.sensor4;
   TraceIn_sensor5[74] := BenchUut5.sensor5;
   TraceIn_station1Start[74] := BenchUut5.station1Start;
   TraceIn_station2Complete[74] := BenchUut5.station2Complete;
   TraceIn_station3Complete[74] := BenchUut5.station3Complete;
   TraceIn_station4Complete[74] := BenchUut5.station4Complete;
   TraceIn_processSequence_1[74] := BenchUut5.processSequence[1];
   TraceIn_processSequence_2[74] := BenchUut5.processSequence[2];
   TraceIn_processSequence_3[74] := BenchUut5.processSequence[3];
   TraceIn_processSequence_4[74] := BenchUut5.processSequence[4];
   TraceIn_processSequence_5[74] := BenchUut5.processSequence[5];
   TraceIn_processSequence_6[74] := BenchUut5.processSequence[6];
   TraceIn_processSequence_7[74] := BenchUut5.processSequence[7];
   TraceIn_processSequence_8[74] := BenchUut5.processSequence[8];
   BenchUut5();
   TraceOut_conveyorLeft[74] := BenchUut5.conveyorLeft;
   TraceOut_conveyorRight[74] := BenchUut5.conveyorRight;
   BenchCalls := BenchCalls + 1;
 75:
   BenchUut5.processLength := USINT#8;
   BenchUut5.sensor1 := FALSE;
   BenchUut5.sensor2 := TRUE;
   BenchUut5.sensor3 := FALSE;
   BenchUut5.sensor4 := FALSE;
   BenchUut5.sensor5 := FALSE;
   BenchUut5.station1Start := FALSE;
   BenchUut5.station2Complete := FALSE;
   BenchUut5.station3Complete := FALSE;
   BenchUut5.station4Complete := FALSE;
   BenchUut5.processSequence[1] := USINT#2;
   BenchUut5.processSequence[2] := USINT#3;
   BenchUut5.processSequence[3] := USINT#4;
   BenchUut5.processSequence[4] := USINT#3;
   BenchUut5.processSequence[5] := USINT#2;
   BenchUut5.processSequence[6] := USINT#4;
   BenchUut5.processSequence[7] := USINT#3;
   BenchUut5.processSequence[8] := USINT#5;
   TraceIn_processLength[75] := BenchUut5.processLength;
   TraceIn_sensor1[75] := BenchUut5.sensor1;
   TraceIn_sensor2[75] := BenchUut5.sensor2;
   TraceIn_sensor3[75] := BenchUut5.sensor3;
   TraceIn_sensor4[75] := BenchUut5.sensor4;
   TraceIn_sensor5[75] := BenchUut5.sensor5;
   TraceIn_station1Start[75] := BenchUut5.station1Start;
   TraceIn_station2Complete[75] := BenchUut5.station2Complete;
   TraceIn_station3Complete[75] := BenchUut5.station3Complete;
   TraceIn_station4Complete[75] := BenchUut5.station4Complete;
   TraceIn_processSequence_1[75] := BenchUut5.processSequence[1];
   TraceIn_processSequence_2[75] := BenchUut5.processSequence[2];
   TraceIn_processSequence_3[75] := BenchUut5.processSequence[3];
   TraceIn_processSequence_4[75] := BenchUut5.processSequence[4];
   TraceIn_processSequence_5[75] := BenchUut5.processSequence[5];
   TraceIn_processSequence_6[75] := BenchUut5.processSequence[6];
   TraceIn_processSequence_7[75] := BenchUut5.processSequence[7];
   TraceIn_processSequence_8[75] := BenchUut5.processSequence[8];
   BenchUut5();
   TraceOut_conveyorLeft[75] := BenchUut5.conveyorLeft;
   TraceOut_conveyorRight[75] := BenchUut5.conveyorRight;
   BenchCalls := BenchCalls + 1;
 76:
   BenchUut5.processLength := USINT#8;
   BenchUut5.sensor1 := FALSE;
   BenchUut5.sensor2 := TRUE;
   BenchUut5.sensor3 := FALSE;
   BenchUut5.sensor4 := FALSE;
   BenchUut5.sensor5 := FALSE;
   BenchUut5.station1Start := FALSE;
   BenchUut5.station2Complete := FALSE;
   BenchUut5.station3Complete := FALSE;
   BenchUut5.station4Complete := FALSE;
   BenchUut5.processSequence[1] := USINT#2;
   BenchUut5.processSequence[2] := USINT#3;
   BenchUut5.processSequence[3] := USINT#4;
   BenchUut5.processSequence[4] := USINT#3;
   BenchUut5.processSequence[5] := USINT#2;
   BenchUut5.processSequence[6] := USINT#4;
   BenchUut5.processSequence[7] := USINT#3;
   BenchUut5.processSequence[8] := USINT#5;
   TraceIn_processLength[76] := BenchUut5.processLength;
   TraceIn_sensor1[76] := BenchUut5.sensor1;
   TraceIn_sensor2[76] := BenchUut5.sensor2;
   TraceIn_sensor3[76] := BenchUut5.sensor3;
   TraceIn_sensor4[76] := BenchUut5.sensor4;
   TraceIn_sensor5[76] := BenchUut5.sensor5;
   TraceIn_station1Start[76] := BenchUut5.station1Start;
   TraceIn_station2Complete[76] := BenchUut5.station2Complete;
   TraceIn_station3Complete[76] := BenchUut5.station3Complete;
   TraceIn_station4Complete[76] := BenchUut5.station4Complete;
   TraceIn_processSequence_1[76] := BenchUut5.processSequence[1];
   TraceIn_processSequence_2[76] := BenchUut5.processSequence[2];
   TraceIn_processSequence_3[76] := BenchUut5.processSequence[3];
   TraceIn_processSequence_4[76] := BenchUut5.processSequence[4];
   TraceIn_processSequence_5[76] := BenchUut5.processSequence[5];
   TraceIn_processSequence_6[76] := BenchUut5.processSequence[6];
   TraceIn_processSequence_7[76] := BenchUut5.processSequence[7];
   TraceIn_processSequence_8[76] := BenchUut5.processSequence[8];
   BenchUut5();
   TraceOut_conveyorLeft[76] := BenchUut5.conveyorLeft;
   TraceOut_conveyorRight[76] := BenchUut5.conveyorRight;
   BenchCalls := BenchCalls + 1;
 77:
   BenchUut5.processLength := USINT#8;
   BenchUut5.sensor1 := FALSE;
   BenchUut5.sensor2 := TRUE;
   BenchUut5.sensor3 := FALSE;
   BenchUut5.sensor4 := FALSE;
   BenchUut5.sensor5 := FALSE;
   BenchUut5.station1Start := FALSE;
   BenchUut5.station2Complete := TRUE;
   BenchUut5.station3Complete := FALSE;
   BenchUut5.station4Complete := FALSE;
   BenchUut5.processSequence[1] := USINT#2;
   BenchUut5.processSequence[2] := USINT#3;
   BenchUut5.processSequence[3] := USINT#4;
   BenchUut5.processSequence[4] := USINT#3;
   BenchUut5.processSequence[5] := USINT#2;
   BenchUut5.processSequence[6] := USINT#4;
   BenchUut5.processSequence[7] := USINT#3;
   BenchUut5.processSequence[8] := USINT#5;
   TraceIn_processLength[77] := BenchUut5.processLength;
   TraceIn_sensor1[77] := BenchUut5.sensor1;
   TraceIn_sensor2[77] := BenchUut5.sensor2;
   TraceIn_sensor3[77] := BenchUut5.sensor3;
   TraceIn_sensor4[77] := BenchUut5.sensor4;
   TraceIn_sensor5[77] := BenchUut5.sensor5;
   TraceIn_station1Start[77] := BenchUut5.station1Start;
   TraceIn_station2Complete[77] := BenchUut5.station2Complete;
   TraceIn_station3Complete[77] := BenchUut5.station3Complete;
   TraceIn_station4Complete[77] := BenchUut5.station4Complete;
   TraceIn_processSequence_1[77] := BenchUut5.processSequence[1];
   TraceIn_processSequence_2[77] := BenchUut5.processSequence[2];
   TraceIn_processSequence_3[77] := BenchUut5.processSequence[3];
   TraceIn_processSequence_4[77] := BenchUut5.processSequence[4];
   TraceIn_processSequence_5[77] := BenchUut5.processSequence[5];
   TraceIn_processSequence_6[77] := BenchUut5.processSequence[6];
   TraceIn_processSequence_7[77] := BenchUut5.processSequence[7];
   TraceIn_processSequence_8[77] := BenchUut5.processSequence[8];
   BenchUut5();
   TraceOut_conveyorLeft[77] := BenchUut5.conveyorLeft;
   TraceOut_conveyorRight[77] := BenchUut5.conveyorRight;
   BenchCalls := BenchCalls + 1;
 78:
   BenchUut5.processLength := USINT#8;
   BenchUut5.sensor1 := FALSE;
   BenchUut5.sensor2 := FALSE;
   BenchUut5.sensor3 := FALSE;
   BenchUut5.sensor4 := FALSE;
   BenchUut5.sensor5 := FALSE;
   BenchUut5.station1Start := FALSE;
   BenchUut5.station2Complete := FALSE;
   BenchUut5.station3Complete := FALSE;
   BenchUut5.station4Complete := FALSE;
   BenchUut5.processSequence[1] := USINT#2;
   BenchUut5.processSequence[2] := USINT#3;
   BenchUut5.processSequence[3] := USINT#4;
   BenchUut5.processSequence[4] := USINT#3;
   BenchUut5.processSequence[5] := USINT#2;
   BenchUut5.processSequence[6] := USINT#4;
   BenchUut5.processSequence[7] := USINT#3;
   BenchUut5.processSequence[8] := USINT#5;
   TraceIn_processLength[78] := BenchUut5.processLength;
   TraceIn_sensor1[78] := BenchUut5.sensor1;
   TraceIn_sensor2[78] := BenchUut5.sensor2;
   TraceIn_sensor3[78] := BenchUut5.sensor3;
   TraceIn_sensor4[78] := BenchUut5.sensor4;
   TraceIn_sensor5[78] := BenchUut5.sensor5;
   TraceIn_station1Start[78] := BenchUut5.station1Start;
   TraceIn_station2Complete[78] := BenchUut5.station2Complete;
   TraceIn_station3Complete[78] := BenchUut5.station3Complete;
   TraceIn_station4Complete[78] := BenchUut5.station4Complete;
   TraceIn_processSequence_1[78] := BenchUut5.processSequence[1];
   TraceIn_processSequence_2[78] := BenchUut5.processSequence[2];
   TraceIn_processSequence_3[78] := BenchUut5.processSequence[3];
   TraceIn_processSequence_4[78] := BenchUut5.processSequence[4];
   TraceIn_processSequence_5[78] := BenchUut5.processSequence[5];
   TraceIn_processSequence_6[78] := BenchUut5.processSequence[6];
   TraceIn_processSequence_7[78] := BenchUut5.processSequence[7];
   TraceIn_processSequence_8[78] := BenchUut5.processSequence[8];
   BenchUut5();
   TraceOut_conveyorLeft[78] := BenchUut5.conveyorLeft;
   TraceOut_conveyorRight[78] := BenchUut5.conveyorRight;
   BenchCalls := BenchCalls + 1;
 79:
   BenchUut5.processLength := USINT#8;
   BenchUut5.sensor1 := FALSE;
   BenchUut5.sensor2 := FALSE;
   BenchUut5.sensor3 := FALSE;
   BenchUut5.sensor4 := FALSE;
   BenchUut5.sensor5 := FALSE;
   BenchUut5.station1Start := FALSE;
   BenchUut5.station2Complete := FALSE;
   BenchUut5.station3Complete := FALSE;
   BenchUut5.station4Complete := FALSE;
   BenchUut5.processSequence[1] := USINT#2;
   BenchUut5.processSequence[2] := USINT#3;
   BenchUut5.processSequence[3] := USINT#4;
   BenchUut5.processSequence[4] := USINT#3;
   BenchUut5.processSequence[5] := USINT#2;
   BenchUut5.processSequence[6] := USINT#4;
   BenchUut5.processSequence[7] := USINT#3;
   BenchUut5.processSequence[8] := USINT#5;
   TraceIn_processLength[79] := BenchUut5.processLength;
   TraceIn_sensor1[79] := BenchUut5.sensor1;
   TraceIn_sensor2[79] := BenchUut5.sensor2;
   TraceIn_sensor3[79] := BenchUut5.sensor3;
   TraceIn_sensor4[79] := BenchUut5.sensor4;
   TraceIn_sensor5[79] := BenchUut5.sensor5;
   TraceIn_station1Start[79] := BenchUut5.station1Start;
   TraceIn_station2Complete[79] := BenchUut5.station2Complete;
   TraceIn_station3Complete[79] := BenchUut5.station3Complete;
   TraceIn_station4Complete[79] := BenchUut5.station4Complete;
   TraceIn_processSequence_1[79] := BenchUut5.processSequence[1];
   TraceIn_processSequence_2[79] := BenchUut5.processSequence[2];
   TraceIn_processSequence_3[79] := BenchUut5.processSequence[3];
   TraceIn_processSequence_4[79] := BenchUut5.processSequence[4];
   TraceIn_processSequence_5[79] := BenchUut5.processSequence[5];
   TraceIn_processSequence_6[79] := BenchUut5.processSequence[6];
   TraceIn_processSequence_7[79] := BenchUut5.processSequence[7];
   TraceIn_processSequence_8[79] := BenchUut5.processSequence[8];
   BenchUut5();
   TraceOut_conveyorLeft[79] := BenchUut5.conveyorLeft;
   TraceOut_conveyorRight[79] := BenchUut5.conveyorRight;
   BenchCalls := BenchCalls + 1;
 80:
   BenchUut5.processLength := USINT#8;
   BenchUut5.sensor1 := FALSE;
   BenchUut5.sensor2 := FALSE;
   BenchUut5.sensor3 := FALSE;
   BenchUut5.sensor4 := TRUE;
   BenchUut5.sensor5 := FALSE;
   BenchUut5.station1Start := FALSE;
   BenchUut5.station2Complete := FALSE;
   BenchUut5.station3Complete := FALSE;
   BenchUut5.station4Complete := FALSE;
   BenchUut5.processSequence[1] := USINT#2;
   BenchUut5.processSequence[2] := USINT#3;
   BenchUut5.processSequence[3] := USINT#4;
   BenchUut5.processSequence[4] := USINT#3;
   BenchUut5.processSequence[5] := USINT#2;
   BenchUut5.processSequence[6] := USINT#4;
   BenchUut5.processSequence[7] := USINT#3;
   BenchUut5.processSequence[8] := USINT#5;
   TraceIn_processLength[80] := BenchUut5.processLength;
   TraceIn_sensor1[80] := BenchUut5.sensor1;
   TraceIn_sensor2[80] := BenchUut5.sensor2;
   TraceIn_sensor3[80] := BenchUut5.sensor3;
   TraceIn_sensor4[80] := BenchUut5.sensor4;
   TraceIn_sensor5[80] := BenchUut5.sensor5;
   TraceIn_station1Start[80] := BenchUut5.station1Start;
   TraceIn_station2Complete[80] := BenchUut5.station2Complete;
   TraceIn_station3Complete[80] := BenchUut5.station3Complete;
   TraceIn_station4Complete[80] := BenchUut5.station4Complete;
   TraceIn_processSequence_1[80] := BenchUut5.processSequence[1];
   TraceIn_processSequence_2[80] := BenchUut5.processSequence[2];
   TraceIn_processSequence_3[80] := BenchUut5.processSequence[3];
   TraceIn_processSequence_4[80] := BenchUut5.processSequence[4];
   TraceIn_processSequence_5[80] := BenchUut5.processSequence[5];
   TraceIn_processSequence_6[80] := BenchUut5.processSequence[6];
   TraceIn_processSequence_7[80] := BenchUut5.processSequence[7];
   TraceIn_processSequence_8[80] := BenchUut5.processSequence[8];
   BenchUut5();
   TraceOut_conveyorLeft[80] := BenchUut5.conveyorLeft;
   TraceOut_conveyorRight[80] := BenchUut5.conveyorRight;
   BenchCalls := BenchCalls + 1;
 81:
   BenchUut5.processLength := USINT#8;
   BenchUut5.sensor1 := FALSE;
   BenchUut5.sensor2 := FALSE;
   BenchUut5.sensor3 := FALSE;
   BenchUut5.sensor4 := TRUE;
   BenchUut5.sensor5 := FALSE;
   BenchUut5.station1Start := FALSE;
   BenchUut5.station2Complete := FALSE;
   BenchUut5.station3Complete := FALSE;
   BenchUut5.station4Complete := FALSE;
   BenchUut5.processSequence[1] := USINT#2;
   BenchUut5.processSequence[2] := USINT#3;
   BenchUut5.processSequence[3] := USINT#4;
   BenchUut5.processSequence[4] := USINT#3;
   BenchUut5.processSequence[5] := USINT#2;
   BenchUut5.processSequence[6] := USINT#4;
   BenchUut5.processSequence[7] := USINT#3;
   BenchUut5.processSequence[8] := USINT#5;
   TraceIn_processLength[81] := BenchUut5.processLength;
   TraceIn_sensor1[81] := BenchUut5.sensor1;
   TraceIn_sensor2[81] := BenchUut5.sensor2;
   TraceIn_sensor3[81] := BenchUut5.sensor3;
   TraceIn_sensor4[81] := BenchUut5.sensor4;
   TraceIn_sensor5[81] := BenchUut5.sensor5;
   TraceIn_station1Start[81] := BenchUut5.station1Start;
   TraceIn_station2Complete[81] := BenchUut5.station2Complete;
   TraceIn_station3Complete[81] := BenchUut5.station3Complete;
   TraceIn_station4Complete[81] := BenchUut5.station4Complete;
   TraceIn_processSequence_1[81] := BenchUut5.processSequence[1];
   TraceIn_processSequence_2[81] := BenchUut5.processSequence[2];
   TraceIn_processSequence_3[81] := BenchUut5.processSequence[3];
   TraceIn_processSequence_4[81] := BenchUut5.processSequence[4];
   TraceIn_processSequence_5[81] := BenchUut5.processSequence[5];
   TraceIn_processSequence_6[81] := BenchUut5.processSequence[6];
   TraceIn_processSequence_7[81] := BenchUut5.processSequence[7];
   TraceIn_processSequence_8[81] := BenchUut5.processSequence[8];
   BenchUut5();
   TraceOut_conveyorLeft[81] := BenchUut5.conveyorLeft;
   TraceOut_conveyorRight[81] := BenchUut5.conveyorRight;
   BenchCalls := BenchCalls + 1;
 82:
   BenchUut5.processLength := USINT#8;
   BenchUut5.sensor1 := FALSE;
   BenchUut5.sensor2 := FALSE;
   BenchUut5.sensor3 := FALSE;
   BenchUut5.sensor4 := TRUE;
   BenchUut5.sensor5 := FALSE;
   BenchUut5.station1Start := FALSE;
   BenchUut5.station2Complete := FALSE;
   BenchUut5.station3Complete := FALSE;
   BenchUut5.station4Complete := FALSE;
   BenchUut5.processSequence[1] := USINT#2;
   BenchUut5.processSequence[2] := USINT#3;
   BenchUut5.processSequence[3] := USINT#4;
   BenchUut5.processSequence[4] := USINT#3;
   BenchUut5.processSequence[5] := USINT#2;
   BenchUut5.processSequence[6] := USINT#4;
   BenchUut5.processSequence[7] := USINT#3;
   BenchUut5.processSequence[8] := USINT#5;
   TraceIn_processLength[82] := BenchUut5.processLength;
   TraceIn_sensor1[82] := BenchUut5.sensor1;
   TraceIn_sensor2[82] := BenchUut5.sensor2;
   TraceIn_sensor3[82] := BenchUut5.sensor3;
   TraceIn_sensor4[82] := BenchUut5.sensor4;
   TraceIn_sensor5[82] := BenchUut5.sensor5;
   TraceIn_station1Start[82] := BenchUut5.station1Start;
   TraceIn_station2Complete[82] := BenchUut5.station2Complete;
   TraceIn_station3Complete[82] := BenchUut5.station3Complete;
   TraceIn_station4Complete[82] := BenchUut5.station4Complete;
   TraceIn_processSequence_1[82] := BenchUut5.processSequence[1];
   TraceIn_processSequence_2[82] := BenchUut5.processSequence[2];
   TraceIn_processSequence_3[82] := BenchUut5.processSequence[3];
   TraceIn_processSequence_4[82] := BenchUut5.processSequence[4];
   TraceIn_processSequence_5[82] := BenchUut5.processSequence[5];
   TraceIn_processSequence_6[82] := BenchUut5.processSequence[6];
   TraceIn_processSequence_7[82] := BenchUut5.processSequence[7];
   TraceIn_processSequence_8[82] := BenchUut5.processSequence[8];
   BenchUut5();
   TraceOut_conveyorLeft[82] := BenchUut5.conveyorLeft;
   TraceOut_conveyorRight[82] := BenchUut5.conveyorRight;
   BenchCalls := BenchCalls + 1;
 83:
   BenchUut5.processLength := USINT#8;
   BenchUut5.sensor1 := FALSE;
   BenchUut5.sensor2 := FALSE;
   BenchUut5.sensor3 := FALSE;
   BenchUut5.sensor4 := TRUE;
   BenchUut5.sensor5 := FALSE;
   BenchUut5.station1Start := FALSE;
   BenchUut5.station2Complete := FALSE;
   BenchUut5.station3Complete := FALSE;
   BenchUut5.station4Complete := TRUE;
   BenchUut5.processSequence[1] := USINT#2;
   BenchUut5.processSequence[2] := USINT#3;
   BenchUut5.processSequence[3] := USINT#4;
   BenchUut5.processSequence[4] := USINT#3;
   BenchUut5.processSequence[5] := USINT#2;
   BenchUut5.processSequence[6] := USINT#4;
   BenchUut5.processSequence[7] := USINT#3;
   BenchUut5.processSequence[8] := USINT#5;
   TraceIn_processLength[83] := BenchUut5.processLength;
   TraceIn_sensor1[83] := BenchUut5.sensor1;
   TraceIn_sensor2[83] := BenchUut5.sensor2;
   TraceIn_sensor3[83] := BenchUut5.sensor3;
   TraceIn_sensor4[83] := BenchUut5.sensor4;
   TraceIn_sensor5[83] := BenchUut5.sensor5;
   TraceIn_station1Start[83] := BenchUut5.station1Start;
   TraceIn_station2Complete[83] := BenchUut5.station2Complete;
   TraceIn_station3Complete[83] := BenchUut5.station3Complete;
   TraceIn_station4Complete[83] := BenchUut5.station4Complete;
   TraceIn_processSequence_1[83] := BenchUut5.processSequence[1];
   TraceIn_processSequence_2[83] := BenchUut5.processSequence[2];
   TraceIn_processSequence_3[83] := BenchUut5.processSequence[3];
   TraceIn_processSequence_4[83] := BenchUut5.processSequence[4];
   TraceIn_processSequence_5[83] := BenchUut5.processSequence[5];
   TraceIn_processSequence_6[83] := BenchUut5.processSequence[6];
   TraceIn_processSequence_7[83] := BenchUut5.processSequence[7];
   TraceIn_processSequence_8[83] := BenchUut5.processSequence[8];
   BenchUut5();
   TraceOut_conveyorLeft[83] := BenchUut5.conveyorLeft;
   TraceOut_conveyorRight[83] := BenchUut5.conveyorRight;
   BenchCalls := BenchCalls + 1;
 84:
   BenchUut5.processLength := USINT#8;
   BenchUut5.sensor1 := FALSE;
   BenchUut5.sensor2 := FALSE;
   BenchUut5.sensor3 := FALSE;
   BenchUut5.sensor4 := FALSE;
   BenchUut5.sensor5 := FALSE;
   BenchUut5.station1Start := FALSE;
   BenchUut5.station2Complete := FALSE;
   BenchUut5.station3Complete := FALSE;
   BenchUut5.station4Complete := FALSE;
   BenchUut5.processSequence[1] := USINT#2;
   BenchUut5.processSequence[2] := USINT#3;
   BenchUut5.processSequence[3] := USINT#4;
   BenchUut5.processSequence[4] := USINT#3;
   BenchUut5.processSequence[5] := USINT#2;
   BenchUut5.processSequence[6] := USINT#4;
   BenchUut5.processSequence[7] := USINT#3;
   BenchUut5.processSequence[8] := USINT#5;
   TraceIn_processLength[84] := BenchUut5.processLength;
   TraceIn_sensor1[84] := BenchUut5.sensor1;
   TraceIn_sensor2[84] := BenchUut5.sensor2;
   TraceIn_sensor3[84] := BenchUut5.sensor3;
   TraceIn_sensor4[84] := BenchUut5.sensor4;
   TraceIn_sensor5[84] := BenchUut5.sensor5;
   TraceIn_station1Start[84] := BenchUut5.station1Start;
   TraceIn_station2Complete[84] := BenchUut5.station2Complete;
   TraceIn_station3Complete[84] := BenchUut5.station3Complete;
   TraceIn_station4Complete[84] := BenchUut5.station4Complete;
   TraceIn_processSequence_1[84] := BenchUut5.processSequence[1];
   TraceIn_processSequence_2[84] := BenchUut5.processSequence[2];
   TraceIn_processSequence_3[84] := BenchUut5.processSequence[3];
   TraceIn_processSequence_4[84] := BenchUut5.processSequence[4];
   TraceIn_processSequence_5[84] := BenchUut5.processSequence[5];
   TraceIn_processSequence_6[84] := BenchUut5.processSequence[6];
   TraceIn_processSequence_7[84] := BenchUut5.processSequence[7];
   TraceIn_processSequence_8[84] := BenchUut5.processSequence[8];
   BenchUut5();
   TraceOut_conveyorLeft[84] := BenchUut5.conveyorLeft;
   TraceOut_conveyorRight[84] := BenchUut5.conveyorRight;
   BenchCalls := BenchCalls + 1;
 85:
   BenchUut5.processLength := USINT#8;
   BenchUut5.sensor1 := FALSE;
   BenchUut5.sensor2 := FALSE;
   BenchUut5.sensor3 := FALSE;
   BenchUut5.sensor4 := FALSE;
   BenchUut5.sensor5 := FALSE;
   BenchUut5.station1Start := FALSE;
   BenchUut5.station2Complete := FALSE;
   BenchUut5.station3Complete := FALSE;
   BenchUut5.station4Complete := FALSE;
   BenchUut5.processSequence[1] := USINT#2;
   BenchUut5.processSequence[2] := USINT#3;
   BenchUut5.processSequence[3] := USINT#4;
   BenchUut5.processSequence[4] := USINT#3;
   BenchUut5.processSequence[5] := USINT#2;
   BenchUut5.processSequence[6] := USINT#4;
   BenchUut5.processSequence[7] := USINT#3;
   BenchUut5.processSequence[8] := USINT#5;
   TraceIn_processLength[85] := BenchUut5.processLength;
   TraceIn_sensor1[85] := BenchUut5.sensor1;
   TraceIn_sensor2[85] := BenchUut5.sensor2;
   TraceIn_sensor3[85] := BenchUut5.sensor3;
   TraceIn_sensor4[85] := BenchUut5.sensor4;
   TraceIn_sensor5[85] := BenchUut5.sensor5;
   TraceIn_station1Start[85] := BenchUut5.station1Start;
   TraceIn_station2Complete[85] := BenchUut5.station2Complete;
   TraceIn_station3Complete[85] := BenchUut5.station3Complete;
   TraceIn_station4Complete[85] := BenchUut5.station4Complete;
   TraceIn_processSequence_1[85] := BenchUut5.processSequence[1];
   TraceIn_processSequence_2[85] := BenchUut5.processSequence[2];
   TraceIn_processSequence_3[85] := BenchUut5.processSequence[3];
   TraceIn_processSequence_4[85] := BenchUut5.processSequence[4];
   TraceIn_processSequence_5[85] := BenchUut5.processSequence[5];
   TraceIn_processSequence_6[85] := BenchUut5.processSequence[6];
   TraceIn_processSequence_7[85] := BenchUut5.processSequence[7];
   TraceIn_processSequence_8[85] := BenchUut5.processSequence[8];
   BenchUut5();
   TraceOut_conveyorLeft[85] := BenchUut5.conveyorLeft;
   TraceOut_conveyorRight[85] := BenchUut5.conveyorRight;
   BenchCalls := BenchCalls + 1;
 86:
   BenchUut5.processLength := USINT#8;
   BenchUut5.sensor1 := FALSE;
   BenchUut5.sensor2 := FALSE;
   BenchUut5.sensor3 := TRUE;
   BenchUut5.sensor4 := FALSE;
   BenchUut5.sensor5 := FALSE;
   BenchUut5.station1Start := FALSE;
   BenchUut5.station2Complete := FALSE;
   BenchUut5.station3Complete := FALSE;
   BenchUut5.station4Complete := FALSE;
   BenchUut5.processSequence[1] := USINT#2;
   BenchUut5.processSequence[2] := USINT#3;
   BenchUut5.processSequence[3] := USINT#4;
   BenchUut5.processSequence[4] := USINT#3;
   BenchUut5.processSequence[5] := USINT#2;
   BenchUut5.processSequence[6] := USINT#4;
   BenchUut5.processSequence[7] := USINT#3;
   BenchUut5.processSequence[8] := USINT#5;
   TraceIn_processLength[86] := BenchUut5.processLength;
   TraceIn_sensor1[86] := BenchUut5.sensor1;
   TraceIn_sensor2[86] := BenchUut5.sensor2;
   TraceIn_sensor3[86] := BenchUut5.sensor3;
   TraceIn_sensor4[86] := BenchUut5.sensor4;
   TraceIn_sensor5[86] := BenchUut5.sensor5;
   TraceIn_station1Start[86] := BenchUut5.station1Start;
   TraceIn_station2Complete[86] := BenchUut5.station2Complete;
   TraceIn_station3Complete[86] := BenchUut5.station3Complete;
   TraceIn_station4Complete[86] := BenchUut5.station4Complete;
   TraceIn_processSequence_1[86] := BenchUut5.processSequence[1];
   TraceIn_processSequence_2[86] := BenchUut5.processSequence[2];
   TraceIn_processSequence_3[86] := BenchUut5.processSequence[3];
   TraceIn_processSequence_4[86] := BenchUut5.processSequence[4];
   TraceIn_processSequence_5[86] := BenchUut5.processSequence[5];
   TraceIn_processSequence_6[86] := BenchUut5.processSequence[6];
   TraceIn_processSequence_7[86] := BenchUut5.processSequence[7];
   TraceIn_processSequence_8[86] := BenchUut5.processSequence[8];
   BenchUut5();
   TraceOut_conveyorLeft[86] := BenchUut5.conveyorLeft;
   TraceOut_conveyorRight[86] := BenchUut5.conveyorRight;
   BenchCalls := BenchCalls + 1;
 87:
   BenchUut5.processLength := USINT#8;
   BenchUut5.sensor1 := FALSE;
   BenchUut5.sensor2 := FALSE;
   BenchUut5.sensor3 := TRUE;
   BenchUut5.sensor4 := FALSE;
   BenchUut5.sensor5 := FALSE;
   BenchUut5.station1Start := FALSE;
   BenchUut5.station2Complete := FALSE;
   BenchUut5.station3Complete := FALSE;
   BenchUut5.station4Complete := FALSE;
   BenchUut5.processSequence[1] := USINT#2;
   BenchUut5.processSequence[2] := USINT#3;
   BenchUut5.processSequence[3] := USINT#4;
   BenchUut5.processSequence[4] := USINT#3;
   BenchUut5.processSequence[5] := USINT#2;
   BenchUut5.processSequence[6] := USINT#4;
   BenchUut5.processSequence[7] := USINT#3;
   BenchUut5.processSequence[8] := USINT#5;
   TraceIn_processLength[87] := BenchUut5.processLength;
   TraceIn_sensor1[87] := BenchUut5.sensor1;
   TraceIn_sensor2[87] := BenchUut5.sensor2;
   TraceIn_sensor3[87] := BenchUut5.sensor3;
   TraceIn_sensor4[87] := BenchUut5.sensor4;
   TraceIn_sensor5[87] := BenchUut5.sensor5;
   TraceIn_station1Start[87] := BenchUut5.station1Start;
   TraceIn_station2Complete[87] := BenchUut5.station2Complete;
   TraceIn_station3Complete[87] := BenchUut5.station3Complete;
   TraceIn_station4Complete[87] := BenchUut5.station4Complete;
   TraceIn_processSequence_1[87] := BenchUut5.processSequence[1];
   TraceIn_processSequence_2[87] := BenchUut5.processSequence[2];
   TraceIn_processSequence_3[87] := BenchUut5.processSequence[3];
   TraceIn_processSequence_4[87] := BenchUut5.processSequence[4];
   TraceIn_processSequence_5[87] := BenchUut5.processSequence[5];
   TraceIn_processSequence_6[87] := BenchUut5.processSequence[6];
   TraceIn_processSequence_7[87] := BenchUut5.processSequence[7];
   TraceIn_processSequence_8[87] := BenchUut5.processSequence[8];
   BenchUut5();
   TraceOut_conveyorLeft[87] := BenchUut5.conveyorLeft;
   TraceOut_conveyorRight[87] := BenchUut5.conveyorRight;
   BenchCalls := BenchCalls + 1;
 88:
   BenchUut5.processLength := USINT#8;
   BenchUut5.sensor1 := FALSE;
   BenchUut5.sensor2 := FALSE;
   BenchUut5.sensor3 := TRUE;
   BenchUut5.sensor4 := FALSE;
   BenchUut5.sensor5 := FALSE;
   BenchUut5.station1Start := FALSE;
   BenchUut5.station2Complete := FALSE;
   BenchUut5.station3Complete := FALSE;
   BenchUut5.station4Complete := FALSE;
   BenchUut5.processSequence[1] := USINT#2;
   BenchUut5.processSequence[2] := USINT#3;
   BenchUut5.processSequence[3] := USINT#4;
   BenchUut5.processSequence[4] := USINT#3;
   BenchUut5.processSequence[5] := USINT#2;
   BenchUut5.processSequence[6] := USINT#4;
   BenchUut5.processSequence[7] := USINT#3;
   BenchUut5.processSequence[8] := USINT#5;
   TraceIn_processLength[88] := BenchUut5.processLength;
   TraceIn_sensor1[88] := BenchUut5.sensor1;
   TraceIn_sensor2[88] := BenchUut5.sensor2;
   TraceIn_sensor3[88] := BenchUut5.sensor3;
   TraceIn_sensor4[88] := BenchUut5.sensor4;
   TraceIn_sensor5[88] := BenchUut5.sensor5;
   TraceIn_station1Start[88] := BenchUut5.station1Start;
   TraceIn_station2Complete[88] := BenchUut5.station2Complete;
   TraceIn_station3Complete[88] := BenchUut5.station3Complete;
   TraceIn_station4Complete[88] := BenchUut5.station4Complete;
   TraceIn_processSequence_1[88] := BenchUut5.processSequence[1];
   TraceIn_processSequence_2[88] := BenchUut5.processSequence[2];
   TraceIn_processSequence_3[88] := BenchUut5.processSequence[3];
   TraceIn_processSequence_4[88] := BenchUut5.processSequence[4];
   TraceIn_processSequence_5[88] := BenchUut5.processSequence[5];
   TraceIn_processSequence_6[88] := BenchUut5.processSequence[6];
   TraceIn_processSequence_7[88] := BenchUut5.processSequence[7];
   TraceIn_processSequence_8[88] := BenchUut5.processSequence[8];
   BenchUut5();
   TraceOut_conveyorLeft[88] := BenchUut5.conveyorLeft;
   TraceOut_conveyorRight[88] := BenchUut5.conveyorRight;
   BenchCalls := BenchCalls + 1;
 89:
   BenchUut5.processLength := USINT#8;
   BenchUut5.sensor1 := FALSE;
   BenchUut5.sensor2 := FALSE;
   BenchUut5.sensor3 := TRUE;
   BenchUut5.sensor4 := FALSE;
   BenchUut5.sensor5 := FALSE;
   BenchUut5.station1Start := FALSE;
   BenchUut5.station2Complete := FALSE;
   BenchUut5.station3Complete := TRUE;
   BenchUut5.station4Complete := FALSE;
   BenchUut5.processSequence[1] := USINT#2;
   BenchUut5.processSequence[2] := USINT#3;
   BenchUut5.processSequence[3] := USINT#4;
   BenchUut5.processSequence[4] := USINT#3;
   BenchUut5.processSequence[5] := USINT#2;
   BenchUut5.processSequence[6] := USINT#4;
   BenchUut5.processSequence[7] := USINT#3;
   BenchUut5.processSequence[8] := USINT#5;
   TraceIn_processLength[89] := BenchUut5.processLength;
   TraceIn_sensor1[89] := BenchUut5.sensor1;
   TraceIn_sensor2[89] := BenchUut5.sensor2;
   TraceIn_sensor3[89] := BenchUut5.sensor3;
   TraceIn_sensor4[89] := BenchUut5.sensor4;
   TraceIn_sensor5[89] := BenchUut5.sensor5;
   TraceIn_station1Start[89] := BenchUut5.station1Start;
   TraceIn_station2Complete[89] := BenchUut5.station2Complete;
   TraceIn_station3Complete[89] := BenchUut5.station3Complete;
   TraceIn_station4Complete[89] := BenchUut5.station4Complete;
   TraceIn_processSequence_1[89] := BenchUut5.processSequence[1];
   TraceIn_processSequence_2[89] := BenchUut5.processSequence[2];
   TraceIn_processSequence_3[89] := BenchUut5.processSequence[3];
   TraceIn_processSequence_4[89] := BenchUut5.processSequence[4];
   TraceIn_processSequence_5[89] := BenchUut5.processSequence[5];
   TraceIn_processSequence_6[89] := BenchUut5.processSequence[6];
   TraceIn_processSequence_7[89] := BenchUut5.processSequence[7];
   TraceIn_processSequence_8[89] := BenchUut5.processSequence[8];
   BenchUut5();
   TraceOut_conveyorLeft[89] := BenchUut5.conveyorLeft;
   TraceOut_conveyorRight[89] := BenchUut5.conveyorRight;
   BenchCalls := BenchCalls + 1;
 90:
   BenchUut5.processLength := USINT#8;
   BenchUut5.sensor1 := FALSE;
   BenchUut5.sensor2 := FALSE;
   BenchUut5.sensor3 := FALSE;
   BenchUut5.sensor4 := FALSE;
   BenchUut5.sensor5 := FALSE;
   BenchUut5.station1Start := FALSE;
   BenchUut5.station2Complete := FALSE;
   BenchUut5.station3Complete := FALSE;
   BenchUut5.station4Complete := FALSE;
   BenchUut5.processSequence[1] := USINT#2;
   BenchUut5.processSequence[2] := USINT#3;
   BenchUut5.processSequence[3] := USINT#4;
   BenchUut5.processSequence[4] := USINT#3;
   BenchUut5.processSequence[5] := USINT#2;
   BenchUut5.processSequence[6] := USINT#4;
   BenchUut5.processSequence[7] := USINT#3;
   BenchUut5.processSequence[8] := USINT#5;
   TraceIn_processLength[90] := BenchUut5.processLength;
   TraceIn_sensor1[90] := BenchUut5.sensor1;
   TraceIn_sensor2[90] := BenchUut5.sensor2;
   TraceIn_sensor3[90] := BenchUut5.sensor3;
   TraceIn_sensor4[90] := BenchUut5.sensor4;
   TraceIn_sensor5[90] := BenchUut5.sensor5;
   TraceIn_station1Start[90] := BenchUut5.station1Start;
   TraceIn_station2Complete[90] := BenchUut5.station2Complete;
   TraceIn_station3Complete[90] := BenchUut5.station3Complete;
   TraceIn_station4Complete[90] := BenchUut5.station4Complete;
   TraceIn_processSequence_1[90] := BenchUut5.processSequence[1];
   TraceIn_processSequence_2[90] := BenchUut5.processSequence[2];
   TraceIn_processSequence_3[90] := BenchUut5.processSequence[3];
   TraceIn_processSequence_4[90] := BenchUut5.processSequence[4];
   TraceIn_processSequence_5[90] := BenchUut5.processSequence[5];
   TraceIn_processSequence_6[90] := BenchUut5.processSequence[6];
   TraceIn_processSequence_7[90] := BenchUut5.processSequence[7];
   TraceIn_processSequence_8[90] := BenchUut5.processSequence[8];
   BenchUut5();
   TraceOut_conveyorLeft[90] := BenchUut5.conveyorLeft;
   TraceOut_conveyorRight[90] := BenchUut5.conveyorRight;
   BenchCalls := BenchCalls + 1;
 91:
   BenchUut5.processLength := USINT#8;
   BenchUut5.sensor1 := FALSE;
   BenchUut5.sensor2 := FALSE;
   BenchUut5.sensor3 := FALSE;
   BenchUut5.sensor4 := FALSE;
   BenchUut5.sensor5 := FALSE;
   BenchUut5.station1Start := FALSE;
   BenchUut5.station2Complete := FALSE;
   BenchUut5.station3Complete := FALSE;
   BenchUut5.station4Complete := FALSE;
   BenchUut5.processSequence[1] := USINT#2;
   BenchUut5.processSequence[2] := USINT#3;
   BenchUut5.processSequence[3] := USINT#4;
   BenchUut5.processSequence[4] := USINT#3;
   BenchUut5.processSequence[5] := USINT#2;
   BenchUut5.processSequence[6] := USINT#4;
   BenchUut5.processSequence[7] := USINT#3;
   BenchUut5.processSequence[8] := USINT#5;
   TraceIn_processLength[91] := BenchUut5.processLength;
   TraceIn_sensor1[91] := BenchUut5.sensor1;
   TraceIn_sensor2[91] := BenchUut5.sensor2;
   TraceIn_sensor3[91] := BenchUut5.sensor3;
   TraceIn_sensor4[91] := BenchUut5.sensor4;
   TraceIn_sensor5[91] := BenchUut5.sensor5;
   TraceIn_station1Start[91] := BenchUut5.station1Start;
   TraceIn_station2Complete[91] := BenchUut5.station2Complete;
   TraceIn_station3Complete[91] := BenchUut5.station3Complete;
   TraceIn_station4Complete[91] := BenchUut5.station4Complete;
   TraceIn_processSequence_1[91] := BenchUut5.processSequence[1];
   TraceIn_processSequence_2[91] := BenchUut5.processSequence[2];
   TraceIn_processSequence_3[91] := BenchUut5.processSequence[3];
   TraceIn_processSequence_4[91] := BenchUut5.processSequence[4];
   TraceIn_processSequence_5[91] := BenchUut5.processSequence[5];
   TraceIn_processSequence_6[91] := BenchUut5.processSequence[6];
   TraceIn_processSequence_7[91] := BenchUut5.processSequence[7];
   TraceIn_processSequence_8[91] := BenchUut5.processSequence[8];
   BenchUut5();
   TraceOut_conveyorLeft[91] := BenchUut5.conveyorLeft;
   TraceOut_conveyorRight[91] := BenchUut5.conveyorRight;
   BenchCalls := BenchCalls + 1;
 92:
   BenchUut5.processLength := USINT#8;
   BenchUut5.sensor1 := FALSE;
   BenchUut5.sensor2 := FALSE;
   BenchUut5.sensor3 := FALSE;
   BenchUut5.sensor4 := FALSE;
   BenchUut5.sensor5 := TRUE;
   BenchUut5.station1Start := FALSE;
   BenchUut5.station2Complete := FALSE;
   BenchUut5.station3Complete := FALSE;
   BenchUut5.station4Complete := FALSE;
   BenchUut5.processSequence[1] := USINT#2;
   BenchUut5.processSequence[2] := USINT#3;
   BenchUut5.processSequence[3] := USINT#4;
   BenchUut5.processSequence[4] := USINT#3;
   BenchUut5.processSequence[5] := USINT#2;
   BenchUut5.processSequence[6] := USINT#4;
   BenchUut5.processSequence[7] := USINT#3;
   BenchUut5.processSequence[8] := USINT#5;
   TraceIn_processLength[92] := BenchUut5.processLength;
   TraceIn_sensor1[92] := BenchUut5.sensor1;
   TraceIn_sensor2[92] := BenchUut5.sensor2;
   TraceIn_sensor3[92] := BenchUut5.sensor3;
   TraceIn_sensor4[92] := BenchUut5.sensor4;
   TraceIn_sensor5[92] := BenchUut5.sensor5;
   TraceIn_station1Start[92] := BenchUut5.station1Start;
   TraceIn_station2Complete[92] := BenchUut5.station2Complete;
   TraceIn_station3Complete[92] := BenchUut5.station3Complete;
   TraceIn_station4Complete[92] := BenchUut5.station4Complete;
   TraceIn_processSequence_1[92] := BenchUut5.processSequence[1];
   TraceIn_processSequence_2[92] := BenchUut5.processSequence[2];
   TraceIn_processSequence_3[92] := BenchUut5.processSequence[3];
   TraceIn_processSequence_4[92] := BenchUut5.processSequence[4];
   TraceIn_processSequence_5[92] := BenchUut5.processSequence[5];
   TraceIn_processSequence_6[92] := BenchUut5.processSequence[6];
   TraceIn_processSequence_7[92] := BenchUut5.processSequence[7];
   TraceIn_processSequence_8[92] := BenchUut5.processSequence[8];
   BenchUut5();
   TraceOut_conveyorLeft[92] := BenchUut5.conveyorLeft;
   TraceOut_conveyorRight[92] := BenchUut5.conveyorRight;
   BenchCalls := BenchCalls + 1;
 93:
   BenchUut5.processLength := USINT#8;
   BenchUut5.sensor1 := TRUE;
   BenchUut5.sensor2 := FALSE;
   BenchUut5.sensor3 := FALSE;
   BenchUut5.sensor4 := FALSE;
   BenchUut5.sensor5 := FALSE;
   BenchUut5.station1Start := TRUE;
   BenchUut5.station2Complete := FALSE;
   BenchUut5.station3Complete := FALSE;
   BenchUut5.station4Complete := FALSE;
   BenchUut5.processSequence[1] := USINT#2;
   BenchUut5.processSequence[2] := USINT#3;
   BenchUut5.processSequence[3] := USINT#4;
   BenchUut5.processSequence[4] := USINT#3;
   BenchUut5.processSequence[5] := USINT#2;
   BenchUut5.processSequence[6] := USINT#4;
   BenchUut5.processSequence[7] := USINT#3;
   BenchUut5.processSequence[8] := USINT#5;
   TraceIn_processLength[93] := BenchUut5.processLength;
   TraceIn_sensor1[93] := BenchUut5.sensor1;
   TraceIn_sensor2[93] := BenchUut5.sensor2;
   TraceIn_sensor3[93] := BenchUut5.sensor3;
   TraceIn_sensor4[93] := BenchUut5.sensor4;
   TraceIn_sensor5[93] := BenchUut5.sensor5;
   TraceIn_station1Start[93] := BenchUut5.station1Start;
   TraceIn_station2Complete[93] := BenchUut5.station2Complete;
   TraceIn_station3Complete[93] := BenchUut5.station3Complete;
   TraceIn_station4Complete[93] := BenchUut5.station4Complete;
   TraceIn_processSequence_1[93] := BenchUut5.processSequence[1];
   TraceIn_processSequence_2[93] := BenchUut5.processSequence[2];
   TraceIn_processSequence_3[93] := BenchUut5.processSequence[3];
   TraceIn_processSequence_4[93] := BenchUut5.processSequence[4];
   TraceIn_processSequence_5[93] := BenchUut5.processSequence[5];
   TraceIn_processSequence_6[93] := BenchUut5.processSequence[6];
   TraceIn_processSequence_7[93] := BenchUut5.processSequence[7];
   TraceIn_processSequence_8[93] := BenchUut5.processSequence[8];
   BenchUut5();
   TraceOut_conveyorLeft[93] := BenchUut5.conveyorLeft;
   TraceOut_conveyorRight[93] := BenchUut5.conveyorRight;
   BenchCalls := BenchCalls + 1;
 94:
   BenchUut5.processLength := USINT#8;
   BenchUut5.sensor1 := FALSE;
   BenchUut5.sensor2 := FALSE;
   BenchUut5.sensor3 := FALSE;
   BenchUut5.sensor4 := FALSE;
   BenchUut5.sensor5 := FALSE;
   BenchUut5.station1Start := FALSE;
   BenchUut5.station2Complete := FALSE;
   BenchUut5.station3Complete := FALSE;
   BenchUut5.station4Complete := FALSE;
   BenchUut5.processSequence[1] := USINT#2;
   BenchUut5.processSequence[2] := USINT#3;
   BenchUut5.processSequence[3] := USINT#4;
   BenchUut5.processSequence[4] := USINT#3;
   BenchUut5.processSequence[5] := USINT#2;
   BenchUut5.processSequence[6] := USINT#4;
   BenchUut5.processSequence[7] := USINT#3;
   BenchUut5.processSequence[8] := USINT#5;
   TraceIn_processLength[94] := BenchUut5.processLength;
   TraceIn_sensor1[94] := BenchUut5.sensor1;
   TraceIn_sensor2[94] := BenchUut5.sensor2;
   TraceIn_sensor3[94] := BenchUut5.sensor3;
   TraceIn_sensor4[94] := BenchUut5.sensor4;
   TraceIn_sensor5[94] := BenchUut5.sensor5;
   TraceIn_station1Start[94] := BenchUut5.station1Start;
   TraceIn_station2Complete[94] := BenchUut5.station2Complete;
   TraceIn_station3Complete[94] := BenchUut5.station3Complete;
   TraceIn_station4Complete[94] := BenchUut5.station4Complete;
   TraceIn_processSequence_1[94] := BenchUut5.processSequence[1];
   TraceIn_processSequence_2[94] := BenchUut5.processSequence[2];
   TraceIn_processSequence_3[94] := BenchUut5.processSequence[3];
   TraceIn_processSequence_4[94] := BenchUut5.processSequence[4];
   TraceIn_processSequence_5[94] := BenchUut5.processSequence[5];
   TraceIn_processSequence_6[94] := BenchUut5.processSequence[6];
   TraceIn_processSequence_7[94] := BenchUut5.processSequence[7];
   TraceIn_processSequence_8[94] := BenchUut5.processSequence[8];
   BenchUut5();
   TraceOut_conveyorLeft[94] := BenchUut5.conveyorLeft;
   TraceOut_conveyorRight[94] := BenchUut5.conveyorRight;
   BenchCalls := BenchCalls + 1;
 95:
   BenchUut5.processLength := USINT#8;
   BenchUut5.sensor1 := FALSE;
   BenchUut5.sensor2 := FALSE;
   BenchUut5.sensor3 := FALSE;
   BenchUut5.sensor4 := FALSE;
   BenchUut5.sensor5 := FALSE;
   BenchUut5.station1Start := FALSE;
   BenchUut5.station2Complete := FALSE;
   BenchUut5.station3Complete := FALSE;
   BenchUut5.station4Complete := FALSE;
   BenchUut5.processSequence[1] := USINT#2;
   BenchUut5.processSequence[2] := USINT#3;
   BenchUut5.processSequence[3] := USINT#4;
   BenchUut5.processSequence[4] := USINT#3;
   BenchUut5.processSequence[5] := USINT#2;
   BenchUut5.processSequence[6] := USINT#4;
   BenchUut5.processSequence[7] := USINT#3;
   BenchUut5.processSequence[8] := USINT#5;
   TraceIn_processLength[95] := BenchUut5.processLength;
   TraceIn_sensor1[95] := BenchUut5.sensor1;
   TraceIn_sensor2[95] := BenchUut5.sensor2;
   TraceIn_sensor3[95] := BenchUut5.sensor3;
   TraceIn_sensor4[95] := BenchUut5.sensor4;
   TraceIn_sensor5[95] := BenchUut5.sensor5;
   TraceIn_station1Start[95] := BenchUut5.station1Start;
   TraceIn_station2Complete[95] := BenchUut5.station2Complete;
   TraceIn_station3Complete[95] := BenchUut5.station3Complete;
   TraceIn_station4Complete[95] := BenchUut5.station4Complete;
   TraceIn_processSequence_1[95] := BenchUut5.processSequence[1];
   TraceIn_processSequence_2[95] := BenchUut5.processSequence[2];
   TraceIn_processSequence_3[95] := BenchUut5.processSequence[3];
   TraceIn_processSequence_4[95] := BenchUut5.processSequence[4];
   TraceIn_processSequence_5[95] := BenchUut5.processSequence[5];
   TraceIn_processSequence_6[95] := BenchUut5.processSequence[6];
   TraceIn_processSequence_7[95] := BenchUut5.processSequence[7];
   TraceIn_processSequence_8[95] := BenchUut5.processSequence[8];
   BenchUut5();
   TraceOut_conveyorLeft[95] := BenchUut5.conveyorLeft;
   TraceOut_conveyorRight[95] := BenchUut5.conveyorRight;
   BenchCalls := BenchCalls + 1;
 96:
   BenchUut5.processLength := USINT#8;
   BenchUut5.sensor1 := FALSE;
   BenchUut5.sensor2 := TRUE;
   BenchUut5.sensor3 := FALSE;
   BenchUut5.sensor4 := FALSE;
   BenchUut5.sensor5 := FALSE;
   BenchUut5.station1Start := FALSE;
   BenchUut5.station2Complete := FALSE;
   BenchUut5.station3Complete := FALSE;
   BenchUut5.station4Complete := FALSE;
   BenchUut5.processSequence[1] := USINT#2;
   BenchUut5.processSequence[2] := USINT#3;
   BenchUut5.processSequence[3] := USINT#4;
   BenchUut5.processSequence[4] := USINT#3;
   BenchUut5.processSequence[5] := USINT#2;
   BenchUut5.processSequence[6] := USINT#4;
   BenchUut5.processSequence[7] := USINT#3;
   BenchUut5.processSequence[8] := USINT#5;
   TraceIn_processLength[96] := BenchUut5.processLength;
   TraceIn_sensor1[96] := BenchUut5.sensor1;
   TraceIn_sensor2[96] := BenchUut5.sensor2;
   TraceIn_sensor3[96] := BenchUut5.sensor3;
   TraceIn_sensor4[96] := BenchUut5.sensor4;
   TraceIn_sensor5[96] := BenchUut5.sensor5;
   TraceIn_station1Start[96] := BenchUut5.station1Start;
   TraceIn_station2Complete[96] := BenchUut5.station2Complete;
   TraceIn_station3Complete[96] := BenchUut5.station3Complete;
   TraceIn_station4Complete[96] := BenchUut5.station4Complete;
   TraceIn_processSequence_1[96] := BenchUut5.processSequence[1];
   TraceIn_processSequence_2[96] := BenchUut5.processSequence[2];
   TraceIn_processSequence_3[96] := BenchUut5.processSequence[3];
   TraceIn_processSequence_4[96] := BenchUut5.processSequence[4];
   TraceIn_processSequence_5[96] := BenchUut5.processSequence[5];
   TraceIn_processSequence_6[96] := BenchUut5.processSequence[6];
   TraceIn_processSequence_7[96] := BenchUut5.processSequence[7];
   TraceIn_processSequence_8[96] := BenchUut5.processSequence[8];
   BenchUut5();
   TraceOut_conveyorLeft[96] := BenchUut5.conveyorLeft;
   TraceOut_conveyorRight[96] := BenchUut5.conveyorRight;
   BenchCalls := BenchCalls + 1;
 97:
   BenchUut5.processLength := USINT#8;
   BenchUut5.sensor1 := FALSE;
   BenchUut5.sensor2 := TRUE;
   BenchUut5.sensor3 := FALSE;
   BenchUut5.sensor4 := FALSE;
   BenchUut5.sensor5 := FALSE;
   BenchUut5.station1Start := FALSE;
   BenchUut5.station2Complete := FALSE;
   BenchUut5.station3Complete := FALSE;
   BenchUut5.station4Complete := FALSE;
   BenchUut5.processSequence[1] := USINT#2;
   BenchUut5.processSequence[2] := USINT#3;
   BenchUut5.processSequence[3] := USINT#4;
   BenchUut5.processSequence[4] := USINT#3;
   BenchUut5.processSequence[5] := USINT#2;
   BenchUut5.processSequence[6] := USINT#4;
   BenchUut5.processSequence[7] := USINT#3;
   BenchUut5.processSequence[8] := USINT#5;
   TraceIn_processLength[97] := BenchUut5.processLength;
   TraceIn_sensor1[97] := BenchUut5.sensor1;
   TraceIn_sensor2[97] := BenchUut5.sensor2;
   TraceIn_sensor3[97] := BenchUut5.sensor3;
   TraceIn_sensor4[97] := BenchUut5.sensor4;
   TraceIn_sensor5[97] := BenchUut5.sensor5;
   TraceIn_station1Start[97] := BenchUut5.station1Start;
   TraceIn_station2Complete[97] := BenchUut5.station2Complete;
   TraceIn_station3Complete[97] := BenchUut5.station3Complete;
   TraceIn_station4Complete[97] := BenchUut5.station4Complete;
   TraceIn_processSequence_1[97] := BenchUut5.processSequence[1];
   TraceIn_processSequence_2[97] := BenchUut5.processSequence[2];
   TraceIn_processSequence_3[97] := BenchUut5.processSequence[3];
   TraceIn_processSequence_4[97] := BenchUut5.processSequence[4];
   TraceIn_processSequence_5[97] := BenchUut5.processSequence[5];
   TraceIn_processSequence_6[97] := BenchUut5.processSequence[6];
   TraceIn_processSequence_7[97] := BenchUut5.processSequence[7];
   TraceIn_processSequence_8[97] := BenchUut5.processSequence[8];
   BenchUut5();
   TraceOut_conveyorLeft[97] := BenchUut5.conveyorLeft;
   TraceOut_conveyorRight[97] := BenchUut5.conveyorRight;
   BenchCalls := BenchCalls + 1;
 98:
   BenchUut5.processLength := USINT#8;
   BenchUut5.sensor1 := FALSE;
   BenchUut5.sensor2 := TRUE;
   BenchUut5.sensor3 := FALSE;
   BenchUut5.sensor4 := FALSE;
   BenchUut5.sensor5 := FALSE;
   BenchUut5.station1Start := FALSE;
   BenchUut5.station2Complete := FALSE;
   BenchUut5.station3Complete := FALSE;
   BenchUut5.station4Complete := FALSE;
   BenchUut5.processSequence[1] := USINT#2;
   BenchUut5.processSequence[2] := USINT#3;
   BenchUut5.processSequence[3] := USINT#4;
   BenchUut5.processSequence[4] := USINT#3;
   BenchUut5.processSequence[5] := USINT#2;
   BenchUut5.processSequence[6] := USINT#4;
   BenchUut5.processSequence[7] := USINT#3;
   BenchUut5.processSequence[8] := USINT#5;
   TraceIn_processLength[98] := BenchUut5.processLength;
   TraceIn_sensor1[98] := BenchUut5.sensor1;
   TraceIn_sensor2[98] := BenchUut5.sensor2;
   TraceIn_sensor3[98] := BenchUut5.sensor3;
   TraceIn_sensor4[98] := BenchUut5.sensor4;
   TraceIn_sensor5[98] := BenchUut5.sensor5;
   TraceIn_station1Start[98] := BenchUut5.station1Start;
   TraceIn_station2Complete[98] := BenchUut5.station2Complete;
   TraceIn_station3Complete[98] := BenchUut5.station3Complete;
   TraceIn_station4Complete[98] := BenchUut5.station4Complete;
   TraceIn_processSequence_1[98] := BenchUut5.processSequence[1];
   TraceIn_processSequence_2[98] := BenchUut5.processSequence[2];
   TraceIn_processSequence_3[98] := BenchUut5.processSequence[3];
   TraceIn_processSequence_4[98] := BenchUut5.processSequence[4];
   TraceIn_processSequence_5[98] := BenchUut5.processSequence[5];
   TraceIn_processSequence_6[98] := BenchUut5.processSequence[6];
   TraceIn_processSequence_7[98] := BenchUut5.processSequence[7];
   TraceIn_processSequence_8[98] := BenchUut5.processSequence[8];
   BenchUut5();
   TraceOut_conveyorLeft[98] := BenchUut5.conveyorLeft;
   TraceOut_conveyorRight[98] := BenchUut5.conveyorRight;
   BenchCalls := BenchCalls + 1;
 99:
   BenchUut5.processLength := USINT#8;
   BenchUut5.sensor1 := FALSE;
   BenchUut5.sensor2 := TRUE;
   BenchUut5.sensor3 := FALSE;
   BenchUut5.sensor4 := FALSE;
   BenchUut5.sensor5 := FALSE;
   BenchUut5.station1Start := FALSE;
   BenchUut5.station2Complete := TRUE;
   BenchUut5.station3Complete := FALSE;
   BenchUut5.station4Complete := FALSE;
   BenchUut5.processSequence[1] := USINT#2;
   BenchUut5.processSequence[2] := USINT#3;
   BenchUut5.processSequence[3] := USINT#4;
   BenchUut5.processSequence[4] := USINT#3;
   BenchUut5.processSequence[5] := USINT#2;
   BenchUut5.processSequence[6] := USINT#4;
   BenchUut5.processSequence[7] := USINT#3;
   BenchUut5.processSequence[8] := USINT#5;
   TraceIn_processLength[99] := BenchUut5.processLength;
   TraceIn_sensor1[99] := BenchUut5.sensor1;
   TraceIn_sensor2[99] := BenchUut5.sensor2;
   TraceIn_sensor3[99] := BenchUut5.sensor3;
   TraceIn_sensor4[99] := BenchUut5.sensor4;
   TraceIn_sensor5[99] := BenchUut5.sensor5;
   TraceIn_station1Start[99] := BenchUut5.station1Start;
   TraceIn_station2Complete[99] := BenchUut5.station2Complete;
   TraceIn_station3Complete[99] := BenchUut5.station3Complete;
   TraceIn_station4Complete[99] := BenchUut5.station4Complete;
   TraceIn_processSequence_1[99] := BenchUut5.processSequence[1];
   TraceIn_processSequence_2[99] := BenchUut5.processSequence[2];
   TraceIn_processSequence_3[99] := BenchUut5.processSequence[3];
   TraceIn_processSequence_4[99] := BenchUut5.processSequence[4];
   TraceIn_processSequence_5[99] := BenchUut5.processSequence[5];
   TraceIn_processSequence_6[99] := BenchUut5.processSequence[6];
   TraceIn_processSequence_7[99] := BenchUut5.processSequence[7];
   TraceIn_processSequence_8[99] := BenchUut5.processSequence[8];
   BenchUut5();
   TraceOut_conveyorLeft[99] := BenchUut5.conveyorLeft;
   TraceOut_conveyorRight[99] := BenchUut5.conveyorRight;
   BenchCalls := BenchCalls + 1;
 100:
   BenchUut5.processLength := USINT#8;
   BenchUut5.sensor1 := FALSE;
   BenchUut5.sensor2 := FALSE;
   BenchUut5.sensor3 := FALSE;
   BenchUut5.sensor4 := FALSE;
   BenchUut5.sensor5 := FALSE;
   BenchUut5.station1Start := FALSE;
   BenchUut5.station2Complete := FALSE;
   BenchUut5.station3Complete := FALSE;
   BenchUut5.station4Complete := FALSE;
   BenchUut5.processSequence[1] := USINT#2;
   BenchUut5.processSequence[2] := USINT#3;
   BenchUut5.processSequence[3] := USINT#4;
   BenchUut5.processSequence[4] := USINT#3;
   BenchUut5.processSequence[5] := USINT#2;
   BenchUut5.processSequence[6] := USINT#4;
   BenchUut5.processSequence[7] := USINT#3;
   BenchUut5.processSequence[8] := USINT#5;
   TraceIn_processLength[100] := BenchUut5.processLength;
   TraceIn_sensor1[100] := BenchUut5.sensor1;
   TraceIn_sensor2[100] := BenchUut5.sensor2;
   TraceIn_sensor3[100] := BenchUut5.sensor3;
   TraceIn_sensor4[100] := BenchUut5.sensor4;
   TraceIn_sensor5[100] := BenchUut5.sensor5;
   TraceIn_station1Start[100] := BenchUut5.station1Start;
   TraceIn_station2Complete[100] := BenchUut5.station2Complete;
   TraceIn_station3Complete[100] := BenchUut5.station3Complete;
   TraceIn_station4Complete[100] := BenchUut5.station4Complete;
   TraceIn_processSequence_1[100] := BenchUut5.processSequence[1];
   TraceIn_processSequence_2[100] := BenchUut5.processSequence[2];
   TraceIn_processSequence_3[100] := BenchUut5.processSequence[3];
   TraceIn_processSequence_4[100] := BenchUut5.processSequence[4];
   TraceIn_processSequence_5[100] := BenchUut5.processSequence[5];
   TraceIn_processSequence_6[100] := BenchUut5.processSequence[6];
   TraceIn_processSequence_7[100] := BenchUut5.processSequence[7];
   TraceIn_processSequence_8[100] := BenchUut5.processSequence[8];
   BenchUut5();
   TraceOut_conveyorLeft[100] := BenchUut5.conveyorLeft;
   TraceOut_conveyorRight[100] := BenchUut5.conveyorRight;
   BenchCalls := BenchCalls + 1;
 101:
   BenchUut5.processLength := USINT#8;
   BenchUut5.sensor1 := FALSE;
   BenchUut5.sensor2 := FALSE;
   BenchUut5.sensor3 := FALSE;
   BenchUut5.sensor4 := FALSE;
   BenchUut5.sensor5 := FALSE;
   BenchUut5.station1Start := FALSE;
   BenchUut5.station2Complete := FALSE;
   BenchUut5.station3Complete := FALSE;
   BenchUut5.station4Complete := FALSE;
   BenchUut5.processSequence[1] := USINT#2;
   BenchUut5.processSequence[2] := USINT#3;
   BenchUut5.processSequence[3] := USINT#4;
   BenchUut5.processSequence[4] := USINT#3;
   BenchUut5.processSequence[5] := USINT#2;
   BenchUut5.processSequence[6] := USINT#4;
   BenchUut5.processSequence[7] := USINT#3;
   BenchUut5.processSequence[8] := USINT#5;
   TraceIn_processLength[101] := BenchUut5.processLength;
   TraceIn_sensor1[101] := BenchUut5.sensor1;
   TraceIn_sensor2[101] := BenchUut5.sensor2;
   TraceIn_sensor3[101] := BenchUut5.sensor3;
   TraceIn_sensor4[101] := BenchUut5.sensor4;
   TraceIn_sensor5[101] := BenchUut5.sensor5;
   TraceIn_station1Start[101] := BenchUut5.station1Start;
   TraceIn_station2Complete[101] := BenchUut5.station2Complete;
   TraceIn_station3Complete[101] := BenchUut5.station3Complete;
   TraceIn_station4Complete[101] := BenchUut5.station4Complete;
   TraceIn_processSequence_1[101] := BenchUut5.processSequence[1];
   TraceIn_processSequence_2[101] := BenchUut5.processSequence[2];
   TraceIn_processSequence_3[101] := BenchUut5.processSequence[3];
   TraceIn_processSequence_4[101] := BenchUut5.processSequence[4];
   TraceIn_processSequence_5[101] := BenchUut5.processSequence[5];
   TraceIn_processSequence_6[101] := BenchUut5.processSequence[6];
   TraceIn_processSequence_7[101] := BenchUut5.processSequence[7];
   TraceIn_processSequence_8[101] := BenchUut5.processSequence[8];
   BenchUut5();
   TraceOut_conveyorLeft[101] := BenchUut5.conveyorLeft;
   TraceOut_conveyorRight[101] := BenchUut5.conveyorRight;
   BenchCalls := BenchCalls + 1;
 102:
   BenchUut5.processLength := USINT#8;
   BenchUut5.sensor1 := FALSE;
   BenchUut5.sensor2 := FALSE;
   BenchUut5.sensor3 := TRUE;
   BenchUut5.sensor4 := FALSE;
   BenchUut5.sensor5 := FALSE;
   BenchUut5.station1Start := FALSE;
   BenchUut5.station2Complete := FALSE;
   BenchUut5.station3Complete := FALSE;
   BenchUut5.station4Complete := FALSE;
   BenchUut5.processSequence[1] := USINT#2;
   BenchUut5.processSequence[2] := USINT#3;
   BenchUut5.processSequence[3] := USINT#4;
   BenchUut5.processSequence[4] := USINT#3;
   BenchUut5.processSequence[5] := USINT#2;
   BenchUut5.processSequence[6] := USINT#4;
   BenchUut5.processSequence[7] := USINT#3;
   BenchUut5.processSequence[8] := USINT#5;
   TraceIn_processLength[102] := BenchUut5.processLength;
   TraceIn_sensor1[102] := BenchUut5.sensor1;
   TraceIn_sensor2[102] := BenchUut5.sensor2;
   TraceIn_sensor3[102] := BenchUut5.sensor3;
   TraceIn_sensor4[102] := BenchUut5.sensor4;
   TraceIn_sensor5[102] := BenchUut5.sensor5;
   TraceIn_station1Start[102] := BenchUut5.station1Start;
   TraceIn_station2Complete[102] := BenchUut5.station2Complete;
   TraceIn_station3Complete[102] := BenchUut5.station3Complete;
   TraceIn_station4Complete[102] := BenchUut5.station4Complete;
   TraceIn_processSequence_1[102] := BenchUut5.processSequence[1];
   TraceIn_processSequence_2[102] := BenchUut5.processSequence[2];
   TraceIn_processSequence_3[102] := BenchUut5.processSequence[3];
   TraceIn_processSequence_4[102] := BenchUut5.processSequence[4];
   TraceIn_processSequence_5[102] := BenchUut5.processSequence[5];
   TraceIn_processSequence_6[102] := BenchUut5.processSequence[6];
   TraceIn_processSequence_7[102] := BenchUut5.processSequence[7];
   TraceIn_processSequence_8[102] := BenchUut5.processSequence[8];
   BenchUut5();
   TraceOut_conveyorLeft[102] := BenchUut5.conveyorLeft;
   TraceOut_conveyorRight[102] := BenchUut5.conveyorRight;
   BenchCalls := BenchCalls + 1;
 103:
   BenchUut5.processLength := USINT#8;
   BenchUut5.sensor1 := FALSE;
   BenchUut5.sensor2 := FALSE;
   BenchUut5.sensor3 := TRUE;
   BenchUut5.sensor4 := FALSE;
   BenchUut5.sensor5 := FALSE;
   BenchUut5.station1Start := FALSE;
   BenchUut5.station2Complete := FALSE;
   BenchUut5.station3Complete := FALSE;
   BenchUut5.station4Complete := FALSE;
   BenchUut5.processSequence[1] := USINT#2;
   BenchUut5.processSequence[2] := USINT#3;
   BenchUut5.processSequence[3] := USINT#4;
   BenchUut5.processSequence[4] := USINT#3;
   BenchUut5.processSequence[5] := USINT#2;
   BenchUut5.processSequence[6] := USINT#4;
   BenchUut5.processSequence[7] := USINT#3;
   BenchUut5.processSequence[8] := USINT#5;
   TraceIn_processLength[103] := BenchUut5.processLength;
   TraceIn_sensor1[103] := BenchUut5.sensor1;
   TraceIn_sensor2[103] := BenchUut5.sensor2;
   TraceIn_sensor3[103] := BenchUut5.sensor3;
   TraceIn_sensor4[103] := BenchUut5.sensor4;
   TraceIn_sensor5[103] := BenchUut5.sensor5;
   TraceIn_station1Start[103] := BenchUut5.station1Start;
   TraceIn_station2Complete[103] := BenchUut5.station2Complete;
   TraceIn_station3Complete[103] := BenchUut5.station3Complete;
   TraceIn_station4Complete[103] := BenchUut5.station4Complete;
   TraceIn_processSequence_1[103] := BenchUut5.processSequence[1];
   TraceIn_processSequence_2[103] := BenchUut5.processSequence[2];
   TraceIn_processSequence_3[103] := BenchUut5.processSequence[3];
   TraceIn_processSequence_4[103] := BenchUut5.processSequence[4];
   TraceIn_processSequence_5[103] := BenchUut5.processSequence[5];
   TraceIn_processSequence_6[103] := BenchUut5.processSequence[6];
   TraceIn_processSequence_7[103] := BenchUut5.processSequence[7];
   TraceIn_processSequence_8[103] := BenchUut5.processSequence[8];
   BenchUut5();
   TraceOut_conveyorLeft[103] := BenchUut5.conveyorLeft;
   TraceOut_conveyorRight[103] := BenchUut5.conveyorRight;
   BenchCalls := BenchCalls + 1;
 104:
   BenchUut5.processLength := USINT#8;
   BenchUut5.sensor1 := FALSE;
   BenchUut5.sensor2 := FALSE;
   BenchUut5.sensor3 := TRUE;
   BenchUut5.sensor4 := FALSE;
   BenchUut5.sensor5 := FALSE;
   BenchUut5.station1Start := FALSE;
   BenchUut5.station2Complete := FALSE;
   BenchUut5.station3Complete := FALSE;
   BenchUut5.station4Complete := FALSE;
   BenchUut5.processSequence[1] := USINT#2;
   BenchUut5.processSequence[2] := USINT#3;
   BenchUut5.processSequence[3] := USINT#4;
   BenchUut5.processSequence[4] := USINT#3;
   BenchUut5.processSequence[5] := USINT#2;
   BenchUut5.processSequence[6] := USINT#4;
   BenchUut5.processSequence[7] := USINT#3;
   BenchUut5.processSequence[8] := USINT#5;
   TraceIn_processLength[104] := BenchUut5.processLength;
   TraceIn_sensor1[104] := BenchUut5.sensor1;
   TraceIn_sensor2[104] := BenchUut5.sensor2;
   TraceIn_sensor3[104] := BenchUut5.sensor3;
   TraceIn_sensor4[104] := BenchUut5.sensor4;
   TraceIn_sensor5[104] := BenchUut5.sensor5;
   TraceIn_station1Start[104] := BenchUut5.station1Start;
   TraceIn_station2Complete[104] := BenchUut5.station2Complete;
   TraceIn_station3Complete[104] := BenchUut5.station3Complete;
   TraceIn_station4Complete[104] := BenchUut5.station4Complete;
   TraceIn_processSequence_1[104] := BenchUut5.processSequence[1];
   TraceIn_processSequence_2[104] := BenchUut5.processSequence[2];
   TraceIn_processSequence_3[104] := BenchUut5.processSequence[3];
   TraceIn_processSequence_4[104] := BenchUut5.processSequence[4];
   TraceIn_processSequence_5[104] := BenchUut5.processSequence[5];
   TraceIn_processSequence_6[104] := BenchUut5.processSequence[6];
   TraceIn_processSequence_7[104] := BenchUut5.processSequence[7];
   TraceIn_processSequence_8[104] := BenchUut5.processSequence[8];
   BenchUut5();
   TraceOut_conveyorLeft[104] := BenchUut5.conveyorLeft;
   TraceOut_conveyorRight[104] := BenchUut5.conveyorRight;
   BenchCalls := BenchCalls + 1;
 105:
   BenchUut5.processLength := USINT#8;
   BenchUut5.sensor1 := FALSE;
   BenchUut5.sensor2 := FALSE;
   BenchUut5.sensor3 := TRUE;
   BenchUut5.sensor4 := FALSE;
   BenchUut5.sensor5 := FALSE;
   BenchUut5.station1Start := FALSE;
   BenchUut5.station2Complete := FALSE;
   BenchUut5.station3Complete := TRUE;
   BenchUut5.station4Complete := FALSE;
   BenchUut5.processSequence[1] := USINT#2;
   BenchUut5.processSequence[2] := USINT#3;
   BenchUut5.processSequence[3] := USINT#4;
   BenchUut5.processSequence[4] := USINT#3;
   BenchUut5.processSequence[5] := USINT#2;
   BenchUut5.processSequence[6] := USINT#4;
   BenchUut5.processSequence[7] := USINT#3;
   BenchUut5.processSequence[8] := USINT#5;
   TraceIn_processLength[105] := BenchUut5.processLength;
   TraceIn_sensor1[105] := BenchUut5.sensor1;
   TraceIn_sensor2[105] := BenchUut5.sensor2;
   TraceIn_sensor3[105] := BenchUut5.sensor3;
   TraceIn_sensor4[105] := BenchUut5.sensor4;
   TraceIn_sensor5[105] := BenchUut5.sensor5;
   TraceIn_station1Start[105] := BenchUut5.station1Start;
   TraceIn_station2Complete[105] := BenchUut5.station2Complete;
   TraceIn_station3Complete[105] := BenchUut5.station3Complete;
   TraceIn_station4Complete[105] := BenchUut5.station4Complete;
   TraceIn_processSequence_1[105] := BenchUut5.processSequence[1];
   TraceIn_processSequence_2[105] := BenchUut5.processSequence[2];
   TraceIn_processSequence_3[105] := BenchUut5.processSequence[3];
   TraceIn_processSequence_4[105] := BenchUut5.processSequence[4];
   TraceIn_processSequence_5[105] := BenchUut5.processSequence[5];
   TraceIn_processSequence_6[105] := BenchUut5.processSequence[6];
   TraceIn_processSequence_7[105] := BenchUut5.processSequence[7];
   TraceIn_processSequence_8[105] := BenchUut5.processSequence[8];
   BenchUut5();
   TraceOut_conveyorLeft[105] := BenchUut5.conveyorLeft;
   TraceOut_conveyorRight[105] := BenchUut5.conveyorRight;
   BenchCalls := BenchCalls + 1;
 106:
   BenchUut5.processLength := USINT#8;
   BenchUut5.sensor1 := FALSE;
   BenchUut5.sensor2 := FALSE;
   BenchUut5.sensor3 := FALSE;
   BenchUut5.sensor4 := FALSE;
   BenchUut5.sensor5 := FALSE;
   BenchUut5.station1Start := FALSE;
   BenchUut5.station2Complete := FALSE;
   BenchUut5.station3Complete := FALSE;
   BenchUut5.station4Complete := FALSE;
   BenchUut5.processSequence[1] := USINT#2;
   BenchUut5.processSequence[2] := USINT#3;
   BenchUut5.processSequence[3] := USINT#4;
   BenchUut5.processSequence[4] := USINT#3;
   BenchUut5.processSequence[5] := USINT#2;
   BenchUut5.processSequence[6] := USINT#4;
   BenchUut5.processSequence[7] := USINT#3;
   BenchUut5.processSequence[8] := USINT#5;
   TraceIn_processLength[106] := BenchUut5.processLength;
   TraceIn_sensor1[106] := BenchUut5.sensor1;
   TraceIn_sensor2[106] := BenchUut5.sensor2;
   TraceIn_sensor3[106] := BenchUut5.sensor3;
   TraceIn_sensor4[106] := BenchUut5.sensor4;
   TraceIn_sensor5[106] := BenchUut5.sensor5;
   TraceIn_station1Start[106] := BenchUut5.station1Start;
   TraceIn_station2Complete[106] := BenchUut5.station2Complete;
   TraceIn_station3Complete[106] := BenchUut5.station3Complete;
   TraceIn_station4Complete[106] := BenchUut5.station4Complete;
   TraceIn_processSequence_1[106] := BenchUut5.processSequence[1];
   TraceIn_processSequence_2[106] := BenchUut5.processSequence[2];
   TraceIn_processSequence_3[106] := BenchUut5.processSequence[3];
   TraceIn_processSequence_4[106] := BenchUut5.processSequence[4];
   TraceIn_processSequence_5[106] := BenchUut5.processSequence[5];
   TraceIn_processSequence_6[106] := BenchUut5.processSequence[6];
   TraceIn_processSequence_7[106] := BenchUut5.processSequence[7];
   TraceIn_processSequence_8[106] := BenchUut5.processSequence[8];
   BenchUut5();
   TraceOut_conveyorLeft[106] := BenchUut5.conveyorLeft;
   TraceOut_conveyorRight[106] := BenchUut5.conveyorRight;
   BenchCalls := BenchCalls + 1;
 107:
   BenchUut5.processLength := USINT#8;
   BenchUut5.sensor1 := FALSE;
   BenchUut5.sensor2 := FALSE;
   BenchUut5.sensor3 := FALSE;
   BenchUut5.sensor4 := FALSE;
   BenchUut5.sensor5 := FALSE;
   BenchUut5.station1Start := FALSE;
   BenchUut5.station2Complete := FALSE;
   BenchUut5.station3Complete := FALSE;
   BenchUut5.station4Complete := FALSE;
   BenchUut5.processSequence[1] := USINT#2;
   BenchUut5.processSequence[2] := USINT#3;
   BenchUut5.processSequence[3] := USINT#4;
   BenchUut5.processSequence[4] := USINT#3;
   BenchUut5.processSequence[5] := USINT#2;
   BenchUut5.processSequence[6] := USINT#4;
   BenchUut5.processSequence[7] := USINT#3;
   BenchUut5.processSequence[8] := USINT#5;
   TraceIn_processLength[107] := BenchUut5.processLength;
   TraceIn_sensor1[107] := BenchUut5.sensor1;
   TraceIn_sensor2[107] := BenchUut5.sensor2;
   TraceIn_sensor3[107] := BenchUut5.sensor3;
   TraceIn_sensor4[107] := BenchUut5.sensor4;
   TraceIn_sensor5[107] := BenchUut5.sensor5;
   TraceIn_station1Start[107] := BenchUut5.station1Start;
   TraceIn_station2Complete[107] := BenchUut5.station2Complete;
   TraceIn_station3Complete[107] := BenchUut5.station3Complete;
   TraceIn_station4Complete[107] := BenchUut5.station4Complete;
   TraceIn_processSequence_1[107] := BenchUut5.processSequence[1];
   TraceIn_processSequence_2[107] := BenchUut5.processSequence[2];
   TraceIn_processSequence_3[107] := BenchUut5.processSequence[3];
   TraceIn_processSequence_4[107] := BenchUut5.processSequence[4];
   TraceIn_processSequence_5[107] := BenchUut5.processSequence[5];
   TraceIn_processSequence_6[107] := BenchUut5.processSequence[6];
   TraceIn_processSequence_7[107] := BenchUut5.processSequence[7];
   TraceIn_processSequence_8[107] := BenchUut5.processSequence[8];
   BenchUut5();
   TraceOut_conveyorLeft[107] := BenchUut5.conveyorLeft;
   TraceOut_conveyorRight[107] := BenchUut5.conveyorRight;
   BenchCalls := BenchCalls + 1;
 108:
   BenchUut5.processLength := USINT#8;
   BenchUut5.sensor1 := FALSE;
   BenchUut5.sensor2 := FALSE;
   BenchUut5.sensor3 := FALSE;
   BenchUut5.sensor4 := TRUE;
   BenchUut5.sensor5 := FALSE;
   BenchUut5.station1Start := FALSE;
   BenchUut5.station2Complete := FALSE;
   BenchUut5.station3Complete := FALSE;
   BenchUut5.station4Complete := FALSE;
   BenchUut5.processSequence[1] := USINT#2;
   BenchUut5.processSequence[2] := USINT#3;
   BenchUut5.processSequence[3] := USINT#4;
   BenchUut5.processSequence[4] := USINT#3;
   BenchUut5.processSequence[5] := USINT#2;
   BenchUut5.processSequence[6] := USINT#4;
   BenchUut5.processSequence[7] := USINT#3;
   BenchUut5.processSequence[8] := USINT#5;
   TraceIn_processLength[108] := BenchUut5.processLength;
   TraceIn_sensor1[108] := BenchUut5.sensor1;
   TraceIn_sensor2[108] := BenchUut5.sensor2;
   TraceIn_sensor3[108] := BenchUut5.sensor3;
   TraceIn_sensor4[108] := BenchUut5.sensor4;
   TraceIn_sensor5[108] := BenchUut5.sensor5;
   TraceIn_station1Start[108] := BenchUut5.station1Start;
   TraceIn_station2Complete[108] := BenchUut5.station2Complete;
   TraceIn_station3Complete[108] := BenchUut5.station3Complete;
   TraceIn_station4Complete[108] := BenchUut5.station4Complete;
   TraceIn_processSequence_1[108] := BenchUut5.processSequence[1];
   TraceIn_processSequence_2[108] := BenchUut5.processSequence[2];
   TraceIn_processSequence_3[108] := BenchUut5.processSequence[3];
   TraceIn_processSequence_4[108] := BenchUut5.processSequence[4];
   TraceIn_processSequence_5[108] := BenchUut5.processSequence[5];
   TraceIn_processSequence_6[108] := BenchUut5.processSequence[6];
   TraceIn_processSequence_7[108] := BenchUut5.processSequence[7];
   TraceIn_processSequence_8[108] := BenchUut5.processSequence[8];
   BenchUut5();
   TraceOut_conveyorLeft[108] := BenchUut5.conveyorLeft;
   TraceOut_conveyorRight[108] := BenchUut5.conveyorRight;
   BenchCalls := BenchCalls + 1;
 109:
   BenchUut5.processLength := USINT#8;
   BenchUut5.sensor1 := FALSE;
   BenchUut5.sensor2 := FALSE;
   BenchUut5.sensor3 := FALSE;
   BenchUut5.sensor4 := TRUE;
   BenchUut5.sensor5 := FALSE;
   BenchUut5.station1Start := FALSE;
   BenchUut5.station2Complete := FALSE;
   BenchUut5.station3Complete := FALSE;
   BenchUut5.station4Complete := FALSE;
   BenchUut5.processSequence[1] := USINT#2;
   BenchUut5.processSequence[2] := USINT#3;
   BenchUut5.processSequence[3] := USINT#4;
   BenchUut5.processSequence[4] := USINT#3;
   BenchUut5.processSequence[5] := USINT#2;
   BenchUut5.processSequence[6] := USINT#4;
   BenchUut5.processSequence[7] := USINT#3;
   BenchUut5.processSequence[8] := USINT#5;
   TraceIn_processLength[109] := BenchUut5.processLength;
   TraceIn_sensor1[109] := BenchUut5.sensor1;
   TraceIn_sensor2[109] := BenchUut5.sensor2;
   TraceIn_sensor3[109] := BenchUut5.sensor3;
   TraceIn_sensor4[109] := BenchUut5.sensor4;
   TraceIn_sensor5[109] := BenchUut5.sensor5;
   TraceIn_station1Start[109] := BenchUut5.station1Start;
   TraceIn_station2Complete[109] := BenchUut5.station2Complete;
   TraceIn_station3Complete[109] := BenchUut5.station3Complete;
   TraceIn_station4Complete[109] := BenchUut5.station4Complete;
   TraceIn_processSequence_1[109] := BenchUut5.processSequence[1];
   TraceIn_processSequence_2[109] := BenchUut5.processSequence[2];
   TraceIn_processSequence_3[109] := BenchUut5.processSequence[3];
   TraceIn_processSequence_4[109] := BenchUut5.processSequence[4];
   TraceIn_processSequence_5[109] := BenchUut5.processSequence[5];
   TraceIn_processSequence_6[109] := BenchUut5.processSequence[6];
   TraceIn_processSequence_7[109] := BenchUut5.processSequence[7];
   TraceIn_processSequence_8[109] := BenchUut5.processSequence[8];
   BenchUut5();
   TraceOut_conveyorLeft[109] := BenchUut5.conveyorLeft;
   TraceOut_conveyorRight[109] := BenchUut5.conveyorRight;
   BenchCalls := BenchCalls + 1;
 110:
   BenchUut5.processLength := USINT#8;
   BenchUut5.sensor1 := FALSE;
   BenchUut5.sensor2 := FALSE;
   BenchUut5.sensor3 := FALSE;
   BenchUut5.sensor4 := TRUE;
   BenchUut5.sensor5 := FALSE;
   BenchUut5.station1Start := FALSE;
   BenchUut5.station2Complete := FALSE;
   BenchUut5.station3Complete := FALSE;
   BenchUut5.station4Complete := FALSE;
   BenchUut5.processSequence[1] := USINT#2;
   BenchUut5.processSequence[2] := USINT#3;
   BenchUut5.processSequence[3] := USINT#4;
   BenchUut5.processSequence[4] := USINT#3;
   BenchUut5.processSequence[5] := USINT#2;
   BenchUut5.processSequence[6] := USINT#4;
   BenchUut5.processSequence[7] := USINT#3;
   BenchUut5.processSequence[8] := USINT#5;
   TraceIn_processLength[110] := BenchUut5.processLength;
   TraceIn_sensor1[110] := BenchUut5.sensor1;
   TraceIn_sensor2[110] := BenchUut5.sensor2;
   TraceIn_sensor3[110] := BenchUut5.sensor3;
   TraceIn_sensor4[110] := BenchUut5.sensor4;
   TraceIn_sensor5[110] := BenchUut5.sensor5;
   TraceIn_station1Start[110] := BenchUut5.station1Start;
   TraceIn_station2Complete[110] := BenchUut5.station2Complete;
   TraceIn_station3Complete[110] := BenchUut5.station3Complete;
   TraceIn_station4Complete[110] := BenchUut5.station4Complete;
   TraceIn_processSequence_1[110] := BenchUut5.processSequence[1];
   TraceIn_processSequence_2[110] := BenchUut5.processSequence[2];
   TraceIn_processSequence_3[110] := BenchUut5.processSequence[3];
   TraceIn_processSequence_4[110] := BenchUut5.processSequence[4];
   TraceIn_processSequence_5[110] := BenchUut5.processSequence[5];
   TraceIn_processSequence_6[110] := BenchUut5.processSequence[6];
   TraceIn_processSequence_7[110] := BenchUut5.processSequence[7];
   TraceIn_processSequence_8[110] := BenchUut5.processSequence[8];
   BenchUut5();
   TraceOut_conveyorLeft[110] := BenchUut5.conveyorLeft;
   TraceOut_conveyorRight[110] := BenchUut5.conveyorRight;
   BenchCalls := BenchCalls + 1;
 111:
   BenchUut5.processLength := USINT#8;
   BenchUut5.sensor1 := FALSE;
   BenchUut5.sensor2 := FALSE;
   BenchUut5.sensor3 := FALSE;
   BenchUut5.sensor4 := TRUE;
   BenchUut5.sensor5 := FALSE;
   BenchUut5.station1Start := FALSE;
   BenchUut5.station2Complete := FALSE;
   BenchUut5.station3Complete := FALSE;
   BenchUut5.station4Complete := TRUE;
   BenchUut5.processSequence[1] := USINT#2;
   BenchUut5.processSequence[2] := USINT#3;
   BenchUut5.processSequence[3] := USINT#4;
   BenchUut5.processSequence[4] := USINT#3;
   BenchUut5.processSequence[5] := USINT#2;
   BenchUut5.processSequence[6] := USINT#4;
   BenchUut5.processSequence[7] := USINT#3;
   BenchUut5.processSequence[8] := USINT#5;
   TraceIn_processLength[111] := BenchUut5.processLength;
   TraceIn_sensor1[111] := BenchUut5.sensor1;
   TraceIn_sensor2[111] := BenchUut5.sensor2;
   TraceIn_sensor3[111] := BenchUut5.sensor3;
   TraceIn_sensor4[111] := BenchUut5.sensor4;
   TraceIn_sensor5[111] := BenchUut5.sensor5;
   TraceIn_station1Start[111] := BenchUut5.station1Start;
   TraceIn_station2Complete[111] := BenchUut5.station2Complete;
   TraceIn_station3Complete[111] := BenchUut5.station3Complete;
   TraceIn_station4Complete[111] := BenchUut5.station4Complete;
   TraceIn_processSequence_1[111] := BenchUut5.processSequence[1];
   TraceIn_processSequence_2[111] := BenchUut5.processSequence[2];
   TraceIn_processSequence_3[111] := BenchUut5.processSequence[3];
   TraceIn_processSequence_4[111] := BenchUut5.processSequence[4];
   TraceIn_processSequence_5[111] := BenchUut5.processSequence[5];
   TraceIn_processSequence_6[111] := BenchUut5.processSequence[6];
   TraceIn_processSequence_7[111] := BenchUut5.processSequence[7];
   TraceIn_processSequence_8[111] := BenchUut5.processSequence[8];
   BenchUut5();
   TraceOut_conveyorLeft[111] := BenchUut5.conveyorLeft;
   TraceOut_conveyorRight[111] := BenchUut5.conveyorRight;
   BenchCalls := BenchCalls + 1;
 112:
   BenchUut5.processLength := USINT#8;
   BenchUut5.sensor1 := FALSE;
   BenchUut5.sensor2 := FALSE;
   BenchUut5.sensor3 := FALSE;
   BenchUut5.sensor4 := FALSE;
   BenchUut5.sensor5 := FALSE;
   BenchUut5.station1Start := FALSE;
   BenchUut5.station2Complete := FALSE;
   BenchUut5.station3Complete := FALSE;
   BenchUut5.station4Complete := FALSE;
   BenchUut5.processSequence[1] := USINT#2;
   BenchUut5.processSequence[2] := USINT#3;
   BenchUut5.processSequence[3] := USINT#4;
   BenchUut5.processSequence[4] := USINT#3;
   BenchUut5.processSequence[5] := USINT#2;
   BenchUut5.processSequence[6] := USINT#4;
   BenchUut5.processSequence[7] := USINT#3;
   BenchUut5.processSequence[8] := USINT#5;
   TraceIn_processLength[112] := BenchUut5.processLength;
   TraceIn_sensor1[112] := BenchUut5.sensor1;
   TraceIn_sensor2[112] := BenchUut5.sensor2;
   TraceIn_sensor3[112] := BenchUut5.sensor3;
   TraceIn_sensor4[112] := BenchUut5.sensor4;
   TraceIn_sensor5[112] := BenchUut5.sensor5;
   TraceIn_station1Start[112] := BenchUut5.station1Start;
   TraceIn_station2Complete[112] := BenchUut5.station2Complete;
   TraceIn_station3Complete[112] := BenchUut5.station3Complete;
   TraceIn_station4Complete[112] := BenchUut5.station4Complete;
   TraceIn_processSequence_1[112] := BenchUut5.processSequence[1];
   TraceIn_processSequence_2[112] := BenchUut5.processSequence[2];
   TraceIn_processSequence_3[112] := BenchUut5.processSequence[3];
   TraceIn_processSequence_4[112] := BenchUut5.processSequence[4];
   TraceIn_processSequence_5[112] := BenchUut5.processSequence[5];
   TraceIn_processSequence_6[112] := BenchUut5.processSequence[6];
   TraceIn_processSequence_7[112] := BenchUut5.processSequence[7];
   TraceIn_processSequence_8[112] := BenchUut5.processSequence[8];
   BenchUut5();
   TraceOut_conveyorLeft[112] := BenchUut5.conveyorLeft;
   TraceOut_conveyorRight[112] := BenchUut5.conveyorRight;
   BenchCalls := BenchCalls + 1;
 113:
   BenchUut5.processLength := USINT#8;
   BenchUut5.sensor1 := FALSE;
   BenchUut5.sensor2 := FALSE;
   BenchUut5.sensor3 := FALSE;
   BenchUut5.sensor4 := FALSE;
   BenchUut5.sensor5 := FALSE;
   BenchUut5.station1Start := FALSE;
   BenchUut5.station2Complete := FALSE;
   BenchUut5.station3Complete := FALSE;
   BenchUut5.station4Complete := FALSE;
   BenchUut5.processSequence[1] := USINT#2;
   BenchUut5.processSequence[2] := USINT#3;
   BenchUut5.processSequence[3] := USINT#4;
   BenchUut5.processSequence[4] := USINT#3;
   BenchUut5.processSequence[5] := USINT#2;
   BenchUut5.processSequence[6] := USINT#4;
   BenchUut5.processSequence[7] := USINT#3;
   BenchUut5.processSequence[8] := USINT#5;
   TraceIn_processLength[113] := BenchUut5.processLength;
   TraceIn_sensor1[113] := BenchUut5.sensor1;
   TraceIn_sensor2[113] := BenchUut5.sensor2;
   TraceIn_sensor3[113] := BenchUut5.sensor3;
   TraceIn_sensor4[113] := BenchUut5.sensor4;
   TraceIn_sensor5[113] := BenchUut5.sensor5;
   TraceIn_station1Start[113] := BenchUut5.station1Start;
   TraceIn_station2Complete[113] := BenchUut5.station2Complete;
   TraceIn_station3Complete[113] := BenchUut5.station3Complete;
   TraceIn_station4Complete[113] := BenchUut5.station4Complete;
   TraceIn_processSequence_1[113] := BenchUut5.processSequence[1];
   TraceIn_processSequence_2[113] := BenchUut5.processSequence[2];
   TraceIn_processSequence_3[113] := BenchUut5.processSequence[3];
   TraceIn_processSequence_4[113] := BenchUut5.processSequence[4];
   TraceIn_processSequence_5[113] := BenchUut5.processSequence[5];
   TraceIn_processSequence_6[113] := BenchUut5.processSequence[6];
   TraceIn_processSequence_7[113] := BenchUut5.processSequence[7];
   TraceIn_processSequence_8[113] := BenchUut5.processSequence[8];
   BenchUut5();
   TraceOut_conveyorLeft[113] := BenchUut5.conveyorLeft;
   TraceOut_conveyorRight[113] := BenchUut5.conveyorRight;
   BenchCalls := BenchCalls + 1;
 114:
   BenchUut5.processLength := USINT#8;
   BenchUut5.sensor1 := FALSE;
   BenchUut5.sensor2 := FALSE;
   BenchUut5.sensor3 := TRUE;
   BenchUut5.sensor4 := FALSE;
   BenchUut5.sensor5 := FALSE;
   BenchUut5.station1Start := FALSE;
   BenchUut5.station2Complete := FALSE;
   BenchUut5.station3Complete := FALSE;
   BenchUut5.station4Complete := FALSE;
   BenchUut5.processSequence[1] := USINT#2;
   BenchUut5.processSequence[2] := USINT#3;
   BenchUut5.processSequence[3] := USINT#4;
   BenchUut5.processSequence[4] := USINT#3;
   BenchUut5.processSequence[5] := USINT#2;
   BenchUut5.processSequence[6] := USINT#4;
   BenchUut5.processSequence[7] := USINT#3;
   BenchUut5.processSequence[8] := USINT#5;
   TraceIn_processLength[114] := BenchUut5.processLength;
   TraceIn_sensor1[114] := BenchUut5.sensor1;
   TraceIn_sensor2[114] := BenchUut5.sensor2;
   TraceIn_sensor3[114] := BenchUut5.sensor3;
   TraceIn_sensor4[114] := BenchUut5.sensor4;
   TraceIn_sensor5[114] := BenchUut5.sensor5;
   TraceIn_station1Start[114] := BenchUut5.station1Start;
   TraceIn_station2Complete[114] := BenchUut5.station2Complete;
   TraceIn_station3Complete[114] := BenchUut5.station3Complete;
   TraceIn_station4Complete[114] := BenchUut5.station4Complete;
   TraceIn_processSequence_1[114] := BenchUut5.processSequence[1];
   TraceIn_processSequence_2[114] := BenchUut5.processSequence[2];
   TraceIn_processSequence_3[114] := BenchUut5.processSequence[3];
   TraceIn_processSequence_4[114] := BenchUut5.processSequence[4];
   TraceIn_processSequence_5[114] := BenchUut5.processSequence[5];
   TraceIn_processSequence_6[114] := BenchUut5.processSequence[6];
   TraceIn_processSequence_7[114] := BenchUut5.processSequence[7];
   TraceIn_processSequence_8[114] := BenchUut5.processSequence[8];
   BenchUut5();
   TraceOut_conveyorLeft[114] := BenchUut5.conveyorLeft;
   TraceOut_conveyorRight[114] := BenchUut5.conveyorRight;
   BenchCalls := BenchCalls + 1;
 115:
   BenchUut5.processLength := USINT#8;
   BenchUut5.sensor1 := FALSE;
   BenchUut5.sensor2 := FALSE;
   BenchUut5.sensor3 := TRUE;
   BenchUut5.sensor4 := FALSE;
   BenchUut5.sensor5 := FALSE;
   BenchUut5.station1Start := FALSE;
   BenchUut5.station2Complete := FALSE;
   BenchUut5.station3Complete := FALSE;
   BenchUut5.station4Complete := FALSE;
   BenchUut5.processSequence[1] := USINT#2;
   BenchUut5.processSequence[2] := USINT#3;
   BenchUut5.processSequence[3] := USINT#4;
   BenchUut5.processSequence[4] := USINT#3;
   BenchUut5.processSequence[5] := USINT#2;
   BenchUut5.processSequence[6] := USINT#4;
   BenchUut5.processSequence[7] := USINT#3;
   BenchUut5.processSequence[8] := USINT#5;
   TraceIn_processLength[115] := BenchUut5.processLength;
   TraceIn_sensor1[115] := BenchUut5.sensor1;
   TraceIn_sensor2[115] := BenchUut5.sensor2;
   TraceIn_sensor3[115] := BenchUut5.sensor3;
   TraceIn_sensor4[115] := BenchUut5.sensor4;
   TraceIn_sensor5[115] := BenchUut5.sensor5;
   TraceIn_station1Start[115] := BenchUut5.station1Start;
   TraceIn_station2Complete[115] := BenchUut5.station2Complete;
   TraceIn_station3Complete[115] := BenchUut5.station3Complete;
   TraceIn_station4Complete[115] := BenchUut5.station4Complete;
   TraceIn_processSequence_1[115] := BenchUut5.processSequence[1];
   TraceIn_processSequence_2[115] := BenchUut5.processSequence[2];
   TraceIn_processSequence_3[115] := BenchUut5.processSequence[3];
   TraceIn_processSequence_4[115] := BenchUut5.processSequence[4];
   TraceIn_processSequence_5[115] := BenchUut5.processSequence[5];
   TraceIn_processSequence_6[115] := BenchUut5.processSequence[6];
   TraceIn_processSequence_7[115] := BenchUut5.processSequence[7];
   TraceIn_processSequence_8[115] := BenchUut5.processSequence[8];
   BenchUut5();
   TraceOut_conveyorLeft[115] := BenchUut5.conveyorLeft;
   TraceOut_conveyorRight[115] := BenchUut5.conveyorRight;
   BenchCalls := BenchCalls + 1;
 116:
   BenchUut5.processLength := USINT#8;
   BenchUut5.sensor1 := FALSE;
   BenchUut5.sensor2 := FALSE;
   BenchUut5.sensor3 := TRUE;
   BenchUut5.sensor4 := FALSE;
   BenchUut5.sensor5 := FALSE;
   BenchUut5.station1Start := FALSE;
   BenchUut5.station2Complete := FALSE;
   BenchUut5.station3Complete := FALSE;
   BenchUut5.station4Complete := FALSE;
   BenchUut5.processSequence[1] := USINT#2;
   BenchUut5.processSequence[2] := USINT#3;
   BenchUut5.processSequence[3] := USINT#4;
   BenchUut5.processSequence[4] := USINT#3;
   BenchUut5.processSequence[5] := USINT#2;
   BenchUut5.processSequence[6] := USINT#4;
   BenchUut5.processSequence[7] := USINT#3;
   BenchUut5.processSequence[8] := USINT#5;
   TraceIn_processLength[116] := BenchUut5.processLength;
   TraceIn_sensor1[116] := BenchUut5.sensor1;
   TraceIn_sensor2[116] := BenchUut5.sensor2;
   TraceIn_sensor3[116] := BenchUut5.sensor3;
   TraceIn_sensor4[116] := BenchUut5.sensor4;
   TraceIn_sensor5[116] := BenchUut5.sensor5;
   TraceIn_station1Start[116] := BenchUut5.station1Start;
   TraceIn_station2Complete[116] := BenchUut5.station2Complete;
   TraceIn_station3Complete[116] := BenchUut5.station3Complete;
   TraceIn_station4Complete[116] := BenchUut5.station4Complete;
   TraceIn_processSequence_1[116] := BenchUut5.processSequence[1];
   TraceIn_processSequence_2[116] := BenchUut5.processSequence[2];
   TraceIn_processSequence_3[116] := BenchUut5.processSequence[3];
   TraceIn_processSequence_4[116] := BenchUut5.processSequence[4];
   TraceIn_processSequence_5[116] := BenchUut5.processSequence[5];
   TraceIn_processSequence_6[116] := BenchUut5.processSequence[6];
   TraceIn_processSequence_7[116] := BenchUut5.processSequence[7];
   TraceIn_processSequence_8[116] := BenchUut5.processSequence[8];
   BenchUut5();
   TraceOut_conveyorLeft[116] := BenchUut5.conveyorLeft;
   TraceOut_conveyorRight[116] := BenchUut5.conveyorRight;
   BenchCalls := BenchCalls + 1;
 117:
   BenchUut5.processLength := USINT#8;
   BenchUut5.sensor1 := FALSE;
   BenchUut5.sensor2 := FALSE;
   BenchUut5.sensor3 := TRUE;
   BenchUut5.sensor4 := FALSE;
   BenchUut5.sensor5 := FALSE;
   BenchUut5.station1Start := FALSE;
   BenchUut5.station2Complete := FALSE;
   BenchUut5.station3Complete := TRUE;
   BenchUut5.station4Complete := FALSE;
   BenchUut5.processSequence[1] := USINT#2;
   BenchUut5.processSequence[2] := USINT#3;
   BenchUut5.processSequence[3] := USINT#4;
   BenchUut5.processSequence[4] := USINT#3;
   BenchUut5.processSequence[5] := USINT#2;
   BenchUut5.processSequence[6] := USINT#4;
   BenchUut5.processSequence[7] := USINT#3;
   BenchUut5.processSequence[8] := USINT#5;
   TraceIn_processLength[117] := BenchUut5.processLength;
   TraceIn_sensor1[117] := BenchUut5.sensor1;
   TraceIn_sensor2[117] := BenchUut5.sensor2;
   TraceIn_sensor3[117] := BenchUut5.sensor3;
   TraceIn_sensor4[117] := BenchUut5.sensor4;
   TraceIn_sensor5[117] := BenchUut5.sensor5;
   TraceIn_station1Start[117] := BenchUut5.station1Start;
   TraceIn_station2Complete[117] := BenchUut5.station2Complete;
   TraceIn_station3Complete[117] := BenchUut5.station3Complete;
   TraceIn_station4Complete[117] := BenchUut5.station4Complete;
   TraceIn_processSequence_1[117] := BenchUut5.processSequence[1];
   TraceIn_processSequence_2[117] := BenchUut5.processSequence[2];
   TraceIn_processSequence_3[117] := BenchUut5.processSequence[3];
   TraceIn_processSequence_4[117] := BenchUut5.processSequence[4];
   TraceIn_processSequence_5[117] := BenchUut5.processSequence[5];
   TraceIn_processSequence_6[117] := BenchUut5.processSequence[6];
   TraceIn_processSequence_7[117] := BenchUut5.processSequence[7];
   TraceIn_processSequence_8[117] := BenchUut5.processSequence[8];
   BenchUut5();
   TraceOut_conveyorLeft[117] := BenchUut5.conveyorLeft;
   TraceOut_conveyorRight[117] := BenchUut5.conveyorRight;
   BenchCalls := BenchCalls + 1;
 118:
   BenchUut5.processLength := USINT#8;
   BenchUut5.sensor1 := FALSE;
   BenchUut5.sensor2 := FALSE;
   BenchUut5.sensor3 := FALSE;
   BenchUut5.sensor4 := FALSE;
   BenchUut5.sensor5 := FALSE;
   BenchUut5.station1Start := FALSE;
   BenchUut5.station2Complete := FALSE;
   BenchUut5.station3Complete := FALSE;
   BenchUut5.station4Complete := FALSE;
   BenchUut5.processSequence[1] := USINT#2;
   BenchUut5.processSequence[2] := USINT#3;
   BenchUut5.processSequence[3] := USINT#4;
   BenchUut5.processSequence[4] := USINT#3;
   BenchUut5.processSequence[5] := USINT#2;
   BenchUut5.processSequence[6] := USINT#4;
   BenchUut5.processSequence[7] := USINT#3;
   BenchUut5.processSequence[8] := USINT#5;
   TraceIn_processLength[118] := BenchUut5.processLength;
   TraceIn_sensor1[118] := BenchUut5.sensor1;
   TraceIn_sensor2[118] := BenchUut5.sensor2;
   TraceIn_sensor3[118] := BenchUut5.sensor3;
   TraceIn_sensor4[118] := BenchUut5.sensor4;
   TraceIn_sensor5[118] := BenchUut5.sensor5;
   TraceIn_station1Start[118] := BenchUut5.station1Start;
   TraceIn_station2Complete[118] := BenchUut5.station2Complete;
   TraceIn_station3Complete[118] := BenchUut5.station3Complete;
   TraceIn_station4Complete[118] := BenchUut5.station4Complete;
   TraceIn_processSequence_1[118] := BenchUut5.processSequence[1];
   TraceIn_processSequence_2[118] := BenchUut5.processSequence[2];
   TraceIn_processSequence_3[118] := BenchUut5.processSequence[3];
   TraceIn_processSequence_4[118] := BenchUut5.processSequence[4];
   TraceIn_processSequence_5[118] := BenchUut5.processSequence[5];
   TraceIn_processSequence_6[118] := BenchUut5.processSequence[6];
   TraceIn_processSequence_7[118] := BenchUut5.processSequence[7];
   TraceIn_processSequence_8[118] := BenchUut5.processSequence[8];
   BenchUut5();
   TraceOut_conveyorLeft[118] := BenchUut5.conveyorLeft;
   TraceOut_conveyorRight[118] := BenchUut5.conveyorRight;
   BenchCalls := BenchCalls + 1;
 119:
   BenchUut5.processLength := USINT#8;
   BenchUut5.sensor1 := FALSE;
   BenchUut5.sensor2 := FALSE;
   BenchUut5.sensor3 := FALSE;
   BenchUut5.sensor4 := FALSE;
   BenchUut5.sensor5 := FALSE;
   BenchUut5.station1Start := FALSE;
   BenchUut5.station2Complete := FALSE;
   BenchUut5.station3Complete := FALSE;
   BenchUut5.station4Complete := FALSE;
   BenchUut5.processSequence[1] := USINT#2;
   BenchUut5.processSequence[2] := USINT#3;
   BenchUut5.processSequence[3] := USINT#4;
   BenchUut5.processSequence[4] := USINT#3;
   BenchUut5.processSequence[5] := USINT#2;
   BenchUut5.processSequence[6] := USINT#4;
   BenchUut5.processSequence[7] := USINT#3;
   BenchUut5.processSequence[8] := USINT#5;
   TraceIn_processLength[119] := BenchUut5.processLength;
   TraceIn_sensor1[119] := BenchUut5.sensor1;
   TraceIn_sensor2[119] := BenchUut5.sensor2;
   TraceIn_sensor3[119] := BenchUut5.sensor3;
   TraceIn_sensor4[119] := BenchUut5.sensor4;
   TraceIn_sensor5[119] := BenchUut5.sensor5;
   TraceIn_station1Start[119] := BenchUut5.station1Start;
   TraceIn_station2Complete[119] := BenchUut5.station2Complete;
   TraceIn_station3Complete[119] := BenchUut5.station3Complete;
   TraceIn_station4Complete[119] := BenchUut5.station4Complete;
   TraceIn_processSequence_1[119] := BenchUut5.processSequence[1];
   TraceIn_processSequence_2[119] := BenchUut5.processSequence[2];
   TraceIn_processSequence_3[119] := BenchUut5.processSequence[3];
   TraceIn_processSequence_4[119] := BenchUut5.processSequence[4];
   TraceIn_processSequence_5[119] := BenchUut5.processSequence[5];
   TraceIn_processSequence_6[119] := BenchUut5.processSequence[6];
   TraceIn_processSequence_7[119] := BenchUut5.processSequence[7];
   TraceIn_processSequence_8[119] := BenchUut5.processSequence[8];
   BenchUut5();
   TraceOut_conveyorLeft[119] := BenchUut5.conveyorLeft;
   TraceOut_conveyorRight[119] := BenchUut5.conveyorRight;
   BenchCalls := BenchCalls + 1;
 120:
   BenchUut5.processLength := USINT#8;
   BenchUut5.sensor1 := FALSE;
   BenchUut5.sensor2 := TRUE;
   BenchUut5.sensor3 := FALSE;
   BenchUut5.sensor4 := FALSE;
   BenchUut5.sensor5 := FALSE;
   BenchUut5.station1Start := FALSE;
   BenchUut5.station2Complete := FALSE;
   BenchUut5.station3Complete := FALSE;
   BenchUut5.station4Complete := FALSE;
   BenchUut5.processSequence[1] := USINT#2;
   BenchUut5.processSequence[2] := USINT#3;
   BenchUut5.processSequence[3] := USINT#4;
   BenchUut5.processSequence[4] := USINT#3;
   BenchUut5.processSequence[5] := USINT#2;
   BenchUut5.processSequence[6] := USINT#4;
   BenchUut5.processSequence[7] := USINT#3;
   BenchUut5.processSequence[8] := USINT#5;
   TraceIn_processLength[120] := BenchUut5.processLength;
   TraceIn_sensor1[120] := BenchUut5.sensor1;
   TraceIn_sensor2[120] := BenchUut5.sensor2;
   TraceIn_sensor3[120] := BenchUut5.sensor3;
   TraceIn_sensor4[120] := BenchUut5.sensor4;
   TraceIn_sensor5[120] := BenchUut5.sensor5;
   TraceIn_station1Start[120] := BenchUut5.station1Start;
   TraceIn_station2Complete[120] := BenchUut5.station2Complete;
   TraceIn_station3Complete[120] := BenchUut5.station3Complete;
   TraceIn_station4Complete[120] := BenchUut5.station4Complete;
   TraceIn_processSequence_1[120] := BenchUut5.processSequence[1];
   TraceIn_processSequence_2[120] := BenchUut5.processSequence[2];
   TraceIn_processSequence_3[120] := BenchUut5.processSequence[3];
   TraceIn_processSequence_4[120] := BenchUut5.processSequence[4];
   TraceIn_processSequence_5[120] := BenchUut5.processSequence[5];
   TraceIn_processSequence_6[120] := BenchUut5.processSequence[6];
   TraceIn_processSequence_7[120] := BenchUut5.processSequence[7];
   TraceIn_processSequence_8[120] := BenchUut5.processSequence[8];
   BenchUut5();
   TraceOut_conveyorLeft[120] := BenchUut5.conveyorLeft;
   TraceOut_conveyorRight[120] := BenchUut5.conveyorRight;
   BenchCalls := BenchCalls + 1;
 121:
   BenchUut5.processLength := USINT#8;
   BenchUut5.sensor1 := FALSE;
   BenchUut5.sensor2 := TRUE;
   BenchUut5.sensor3 := FALSE;
   BenchUut5.sensor4 := FALSE;
   BenchUut5.sensor5 := FALSE;
   BenchUut5.station1Start := FALSE;
   BenchUut5.station2Complete := FALSE;
   BenchUut5.station3Complete := FALSE;
   BenchUut5.station4Complete := FALSE;
   BenchUut5.processSequence[1] := USINT#2;
   BenchUut5.processSequence[2] := USINT#3;
   BenchUut5.processSequence[3] := USINT#4;
   BenchUut5.processSequence[4] := USINT#3;
   BenchUut5.processSequence[5] := USINT#2;
   BenchUut5.processSequence[6] := USINT#4;
   BenchUut5.processSequence[7] := USINT#3;
   BenchUut5.processSequence[8] := USINT#5;
   TraceIn_processLength[121] := BenchUut5.processLength;
   TraceIn_sensor1[121] := BenchUut5.sensor1;
   TraceIn_sensor2[121] := BenchUut5.sensor2;
   TraceIn_sensor3[121] := BenchUut5.sensor3;
   TraceIn_sensor4[121] := BenchUut5.sensor4;
   TraceIn_sensor5[121] := BenchUut5.sensor5;
   TraceIn_station1Start[121] := BenchUut5.station1Start;
   TraceIn_station2Complete[121] := BenchUut5.station2Complete;
   TraceIn_station3Complete[121] := BenchUut5.station3Complete;
   TraceIn_station4Complete[121] := BenchUut5.station4Complete;
   TraceIn_processSequence_1[121] := BenchUut5.processSequence[1];
   TraceIn_processSequence_2[121] := BenchUut5.processSequence[2];
   TraceIn_processSequence_3[121] := BenchUut5.processSequence[3];
   TraceIn_processSequence_4[121] := BenchUut5.processSequence[4];
   TraceIn_processSequence_5[121] := BenchUut5.processSequence[5];
   TraceIn_processSequence_6[121] := BenchUut5.processSequence[6];
   TraceIn_processSequence_7[121] := BenchUut5.processSequence[7];
   TraceIn_processSequence_8[121] := BenchUut5.processSequence[8];
   BenchUut5();
   TraceOut_conveyorLeft[121] := BenchUut5.conveyorLeft;
   TraceOut_conveyorRight[121] := BenchUut5.conveyorRight;
   BenchCalls := BenchCalls + 1;
 122:
   BenchUut5.processLength := USINT#8;
   BenchUut5.sensor1 := FALSE;
   BenchUut5.sensor2 := TRUE;
   BenchUut5.sensor3 := FALSE;
   BenchUut5.sensor4 := FALSE;
   BenchUut5.sensor5 := FALSE;
   BenchUut5.station1Start := FALSE;
   BenchUut5.station2Complete := FALSE;
   BenchUut5.station3Complete := FALSE;
   BenchUut5.station4Complete := FALSE;
   BenchUut5.processSequence[1] := USINT#2;
   BenchUut5.processSequence[2] := USINT#3;
   BenchUut5.processSequence[3] := USINT#4;
   BenchUut5.processSequence[4] := USINT#3;
   BenchUut5.processSequence[5] := USINT#2;
   BenchUut5.processSequence[6] := USINT#4;
   BenchUut5.processSequence[7] := USINT#3;
   BenchUut5.processSequence[8] := USINT#5;
   TraceIn_processLength[122] := BenchUut5.processLength;
   TraceIn_sensor1[122] := BenchUut5.sensor1;
   TraceIn_sensor2[122] := BenchUut5.sensor2;
   TraceIn_sensor3[122] := BenchUut5.sensor3;
   TraceIn_sensor4[122] := BenchUut5.sensor4;
   TraceIn_sensor5[122] := BenchUut5.sensor5;
   TraceIn_station1Start[122] := BenchUut5.station1Start;
   TraceIn_station2Complete[122] := BenchUut5.station2Complete;
   TraceIn_station3Complete[122] := BenchUut5.station3Complete;
   TraceIn_station4Complete[122] := BenchUut5.station4Complete;
   TraceIn_processSequence_1[122] := BenchUut5.processSequence[1];
   TraceIn_processSequence_2[122] := BenchUut5.processSequence[2];
   TraceIn_processSequence_3[122] := BenchUut5.processSequence[3];
   TraceIn_processSequence_4[122] := BenchUut5.processSequence[4];
   TraceIn_processSequence_5[122] := BenchUut5.processSequence[5];
   TraceIn_processSequence_6[122] := BenchUut5.processSequence[6];
   TraceIn_processSequence_7[122] := BenchUut5.processSequence[7];
   TraceIn_processSequence_8[122] := BenchUut5.processSequence[8];
   BenchUut5();
   TraceOut_conveyorLeft[122] := BenchUut5.conveyorLeft;
   TraceOut_conveyorRight[122] := BenchUut5.conveyorRight;
   BenchCalls := BenchCalls + 1;
 123:
   BenchUut5.processLength := USINT#8;
   BenchUut5.sensor1 := FALSE;
   BenchUut5.sensor2 := TRUE;
   BenchUut5.sensor3 := FALSE;
   BenchUut5.sensor4 := FALSE;
   BenchUut5.sensor5 := FALSE;
   BenchUut5.station1Start := FALSE;
   BenchUut5.station2Complete := TRUE;
   BenchUut5.station3Complete := FALSE;
   BenchUut5.station4Complete := FALSE;
   BenchUut5.processSequence[1] := USINT#2;
   BenchUut5.processSequence[2] := USINT#3;
   BenchUut5.processSequence[3] := USINT#4;
   BenchUut5.processSequence[4] := USINT#3;
   BenchUut5.processSequence[5] := USINT#2;
   BenchUut5.processSequence[6] := USINT#4;
   BenchUut5.processSequence[7] := USINT#3;
   BenchUut5.processSequence[8] := USINT#5;
   TraceIn_processLength[123] := BenchUut5.processLength;
   TraceIn_sensor1[123] := BenchUut5.sensor1;
   TraceIn_sensor2[123] := BenchUut5.sensor2;
   TraceIn_sensor3[123] := BenchUut5.sensor3;
   TraceIn_sensor4[123] := BenchUut5.sensor4;
   TraceIn_sensor5[123] := BenchUut5.sensor5;
   TraceIn_station1Start[123] := BenchUut5.station1Start;
   TraceIn_station2Complete[123] := BenchUut5.station2Complete;
   TraceIn_station3Complete[123] := BenchUut5.station3Complete;
   TraceIn_station4Complete[123] := BenchUut5.station4Complete;
   TraceIn_processSequence_1[123] := BenchUut5.processSequence[1];
   TraceIn_processSequence_2[123] := BenchUut5.processSequence[2];
   TraceIn_processSequence_3[123] := BenchUut5.processSequence[3];
   TraceIn_processSequence_4[123] := BenchUut5.processSequence[4];
   TraceIn_processSequence_5[123] := BenchUut5.processSequence[5];
   TraceIn_processSequence_6[123] := BenchUut5.processSequence[6];
   TraceIn_processSequence_7[123] := BenchUut5.processSequence[7];
   TraceIn_processSequence_8[123] := BenchUut5.processSequence[8];
   BenchUut5();
   TraceOut_conveyorLeft[123] := BenchUut5.conveyorLeft;
   TraceOut_conveyorRight[123] := BenchUut5.conveyorRight;
   BenchCalls := BenchCalls + 1;
 124:
   BenchUut5.processLength := USINT#8;
   BenchUut5.sensor1 := FALSE;
   BenchUut5.sensor2 := FALSE;
   BenchUut5.sensor3 := FALSE;
   BenchUut5.sensor4 := FALSE;
   BenchUut5.sensor5 := FALSE;
   BenchUut5.station1Start := FALSE;
   BenchUut5.station2Complete := FALSE;
   BenchUut5.station3Complete := FALSE;
   BenchUut5.station4Complete := FALSE;
   BenchUut5.processSequence[1] := USINT#2;
   BenchUut5.processSequence[2] := USINT#3;
   BenchUut5.processSequence[3] := USINT#4;
   BenchUut5.processSequence[4] := USINT#3;
   BenchUut5.processSequence[5] := USINT#2;
   BenchUut5.processSequence[6] := USINT#4;
   BenchUut5.processSequence[7] := USINT#3;
   BenchUut5.processSequence[8] := USINT#5;
   TraceIn_processLength[124] := BenchUut5.processLength;
   TraceIn_sensor1[124] := BenchUut5.sensor1;
   TraceIn_sensor2[124] := BenchUut5.sensor2;
   TraceIn_sensor3[124] := BenchUut5.sensor3;
   TraceIn_sensor4[124] := BenchUut5.sensor4;
   TraceIn_sensor5[124] := BenchUut5.sensor5;
   TraceIn_station1Start[124] := BenchUut5.station1Start;
   TraceIn_station2Complete[124] := BenchUut5.station2Complete;
   TraceIn_station3Complete[124] := BenchUut5.station3Complete;
   TraceIn_station4Complete[124] := BenchUut5.station4Complete;
   TraceIn_processSequence_1[124] := BenchUut5.processSequence[1];
   TraceIn_processSequence_2[124] := BenchUut5.processSequence[2];
   TraceIn_processSequence_3[124] := BenchUut5.processSequence[3];
   TraceIn_processSequence_4[124] := BenchUut5.processSequence[4];
   TraceIn_processSequence_5[124] := BenchUut5.processSequence[5];
   TraceIn_processSequence_6[124] := BenchUut5.processSequence[6];
   TraceIn_processSequence_7[124] := BenchUut5.processSequence[7];
   TraceIn_processSequence_8[124] := BenchUut5.processSequence[8];
   BenchUut5();
   TraceOut_conveyorLeft[124] := BenchUut5.conveyorLeft;
   TraceOut_conveyorRight[124] := BenchUut5.conveyorRight;
   BenchCalls := BenchCalls + 1;
 125:
   BenchUut5.processLength := USINT#8;
   BenchUut5.sensor1 := FALSE;
   BenchUut5.sensor2 := FALSE;
   BenchUut5.sensor3 := FALSE;
   BenchUut5.sensor4 := FALSE;
   BenchUut5.sensor5 := FALSE;
   BenchUut5.station1Start := FALSE;
   BenchUut5.station2Complete := FALSE;
   BenchUut5.station3Complete := FALSE;
   BenchUut5.station4Complete := FALSE;
   BenchUut5.processSequence[1] := USINT#2;
   BenchUut5.processSequence[2] := USINT#3;
   BenchUut5.processSequence[3] := USINT#4;
   BenchUut5.processSequence[4] := USINT#3;
   BenchUut5.processSequence[5] := USINT#2;
   BenchUut5.processSequence[6] := USINT#4;
   BenchUut5.processSequence[7] := USINT#3;
   BenchUut5.processSequence[8] := USINT#5;
   TraceIn_processLength[125] := BenchUut5.processLength;
   TraceIn_sensor1[125] := BenchUut5.sensor1;
   TraceIn_sensor2[125] := BenchUut5.sensor2;
   TraceIn_sensor3[125] := BenchUut5.sensor3;
   TraceIn_sensor4[125] := BenchUut5.sensor4;
   TraceIn_sensor5[125] := BenchUut5.sensor5;
   TraceIn_station1Start[125] := BenchUut5.station1Start;
   TraceIn_station2Complete[125] := BenchUut5.station2Complete;
   TraceIn_station3Complete[125] := BenchUut5.station3Complete;
   TraceIn_station4Complete[125] := BenchUut5.station4Complete;
   TraceIn_processSequence_1[125] := BenchUut5.processSequence[1];
   TraceIn_processSequence_2[125] := BenchUut5.processSequence[2];
   TraceIn_processSequence_3[125] := BenchUut5.processSequence[3];
   TraceIn_processSequence_4[125] := BenchUut5.processSequence[4];
   TraceIn_processSequence_5[125] := BenchUut5.processSequence[5];
   TraceIn_processSequence_6[125] := BenchUut5.processSequence[6];
   TraceIn_processSequence_7[125] := BenchUut5.processSequence[7];
   TraceIn_processSequence_8[125] := BenchUut5.processSequence[8];
   BenchUut5();
   TraceOut_conveyorLeft[125] := BenchUut5.conveyorLeft;
   TraceOut_conveyorRight[125] := BenchUut5.conveyorRight;
   BenchCalls := BenchCalls + 1;
 126:
   BenchUut5.processLength := USINT#8;
   BenchUut5.sensor1 := FALSE;
   BenchUut5.sensor2 := FALSE;
   BenchUut5.sensor3 := FALSE;
   BenchUut5.sensor4 := TRUE;
   BenchUut5.sensor5 := FALSE;
   BenchUut5.station1Start := FALSE;
   BenchUut5.station2Complete := FALSE;
   BenchUut5.station3Complete := FALSE;
   BenchUut5.station4Complete := FALSE;
   BenchUut5.processSequence[1] := USINT#2;
   BenchUut5.processSequence[2] := USINT#3;
   BenchUut5.processSequence[3] := USINT#4;
   BenchUut5.processSequence[4] := USINT#3;
   BenchUut5.processSequence[5] := USINT#2;
   BenchUut5.processSequence[6] := USINT#4;
   BenchUut5.processSequence[7] := USINT#3;
   BenchUut5.processSequence[8] := USINT#5;
   TraceIn_processLength[126] := BenchUut5.processLength;
   TraceIn_sensor1[126] := BenchUut5.sensor1;
   TraceIn_sensor2[126] := BenchUut5.sensor2;
   TraceIn_sensor3[126] := BenchUut5.sensor3;
   TraceIn_sensor4[126] := BenchUut5.sensor4;
   TraceIn_sensor5[126] := BenchUut5.sensor5;
   TraceIn_station1Start[126] := BenchUut5.station1Start;
   TraceIn_station2Complete[126] := BenchUut5.station2Complete;
   TraceIn_station3Complete[126] := BenchUut5.station3Complete;
   TraceIn_station4Complete[126] := BenchUut5.station4Complete;
   TraceIn_processSequence_1[126] := BenchUut5.processSequence[1];
   TraceIn_processSequence_2[126] := BenchUut5.processSequence[2];
   TraceIn_processSequence_3[126] := BenchUut5.processSequence[3];
   TraceIn_processSequence_4[126] := BenchUut5.processSequence[4];
   TraceIn_processSequence_5[126] := BenchUut5.processSequence[5];
   TraceIn_processSequence_6[126] := BenchUut5.processSequence[6];
   TraceIn_processSequence_7[126] := BenchUut5.processSequence[7];
   TraceIn_processSequence_8[126] := BenchUut5.processSequence[8];
   BenchUut5();
   TraceOut_conveyorLeft[126] := BenchUut5.conveyorLeft;
   TraceOut_conveyorRight[126] := BenchUut5.conveyorRight;
   BenchCalls := BenchCalls + 1;
 127:
   BenchUut5.processLength := USINT#8;
   BenchUut5.sensor1 := FALSE;
   BenchUut5.sensor2 := FALSE;
   BenchUut5.sensor3 := FALSE;
   BenchUut5.sensor4 := TRUE;
   BenchUut5.sensor5 := FALSE;
   BenchUut5.station1Start := FALSE;
   BenchUut5.station2Complete := FALSE;
   BenchUut5.station3Complete := FALSE;
   BenchUut5.station4Complete := FALSE;
   BenchUut5.processSequence[1] := USINT#2;
   BenchUut5.processSequence[2] := USINT#3;
   BenchUut5.processSequence[3] := USINT#4;
   BenchUut5.processSequence[4] := USINT#3;
   BenchUut5.processSequence[5] := USINT#2;
   BenchUut5.processSequence[6] := USINT#4;
   BenchUut5.processSequence[7] := USINT#3;
   BenchUut5.processSequence[8] := USINT#5;
   TraceIn_processLength[127] := BenchUut5.processLength;
   TraceIn_sensor1[127] := BenchUut5.sensor1;
   TraceIn_sensor2[127] := BenchUut5.sensor2;
   TraceIn_sensor3[127] := BenchUut5.sensor3;
   TraceIn_sensor4[127] := BenchUut5.sensor4;
   TraceIn_sensor5[127] := BenchUut5.sensor5;
   TraceIn_station1Start[127] := BenchUut5.station1Start;
   TraceIn_station2Complete[127] := BenchUut5.station2Complete;
   TraceIn_station3Complete[127] := BenchUut5.station3Complete;
   TraceIn_station4Complete[127] := BenchUut5.station4Complete;
   TraceIn_processSequence_1[127] := BenchUut5.processSequence[1];
   TraceIn_processSequence_2[127] := BenchUut5.processSequence[2];
   TraceIn_processSequence_3[127] := BenchUut5.processSequence[3];
   TraceIn_processSequence_4[127] := BenchUut5.processSequence[4];
   TraceIn_processSequence_5[127] := BenchUut5.processSequence[5];
   TraceIn_processSequence_6[127] := BenchUut5.processSequence[6];
   TraceIn_processSequence_7[127] := BenchUut5.processSequence[7];
   TraceIn_processSequence_8[127] := BenchUut5.processSequence[8];
   BenchUut5();
   TraceOut_conveyorLeft[127] := BenchUut5.conveyorLeft;
   TraceOut_conveyorRight[127] := BenchUut5.conveyorRight;
   BenchCalls := BenchCalls + 1;
 128:
   BenchUut5.processLength := USINT#8;
   BenchUut5.sensor1 := FALSE;
   BenchUut5.sensor2 := FALSE;
   BenchUut5.sensor3 := FALSE;
   BenchUut5.sensor4 := TRUE;
   BenchUut5.sensor5 := FALSE;
   BenchUut5.station1Start := FALSE;
   BenchUut5.station2Complete := FALSE;
   BenchUut5.station3Complete := FALSE;
   BenchUut5.station4Complete := FALSE;
   BenchUut5.processSequence[1] := USINT#2;
   BenchUut5.processSequence[2] := USINT#3;
   BenchUut5.processSequence[3] := USINT#4;
   BenchUut5.processSequence[4] := USINT#3;
   BenchUut5.processSequence[5] := USINT#2;
   BenchUut5.processSequence[6] := USINT#4;
   BenchUut5.processSequence[7] := USINT#3;
   BenchUut5.processSequence[8] := USINT#5;
   TraceIn_processLength[128] := BenchUut5.processLength;
   TraceIn_sensor1[128] := BenchUut5.sensor1;
   TraceIn_sensor2[128] := BenchUut5.sensor2;
   TraceIn_sensor3[128] := BenchUut5.sensor3;
   TraceIn_sensor4[128] := BenchUut5.sensor4;
   TraceIn_sensor5[128] := BenchUut5.sensor5;
   TraceIn_station1Start[128] := BenchUut5.station1Start;
   TraceIn_station2Complete[128] := BenchUut5.station2Complete;
   TraceIn_station3Complete[128] := BenchUut5.station3Complete;
   TraceIn_station4Complete[128] := BenchUut5.station4Complete;
   TraceIn_processSequence_1[128] := BenchUut5.processSequence[1];
   TraceIn_processSequence_2[128] := BenchUut5.processSequence[2];
   TraceIn_processSequence_3[128] := BenchUut5.processSequence[3];
   TraceIn_processSequence_4[128] := BenchUut5.processSequence[4];
   TraceIn_processSequence_5[128] := BenchUut5.processSequence[5];
   TraceIn_processSequence_6[128] := BenchUut5.processSequence[6];
   TraceIn_processSequence_7[128] := BenchUut5.processSequence[7];
   TraceIn_processSequence_8[128] := BenchUut5.processSequence[8];
   BenchUut5();
   TraceOut_conveyorLeft[128] := BenchUut5.conveyorLeft;
   TraceOut_conveyorRight[128] := BenchUut5.conveyorRight;
   BenchCalls := BenchCalls + 1;
 129:
   BenchUut5.processLength := USINT#8;
   BenchUut5.sensor1 := FALSE;
   BenchUut5.sensor2 := FALSE;
   BenchUut5.sensor3 := FALSE;
   BenchUut5.sensor4 := TRUE;
   BenchUut5.sensor5 := FALSE;
   BenchUut5.station1Start := FALSE;
   BenchUut5.station2Complete := FALSE;
   BenchUut5.station3Complete := FALSE;
   BenchUut5.station4Complete := TRUE;
   BenchUut5.processSequence[1] := USINT#2;
   BenchUut5.processSequence[2] := USINT#3;
   BenchUut5.processSequence[3] := USINT#4;
   BenchUut5.processSequence[4] := USINT#3;
   BenchUut5.processSequence[5] := USINT#2;
   BenchUut5.processSequence[6] := USINT#4;
   BenchUut5.processSequence[7] := USINT#3;
   BenchUut5.processSequence[8] := USINT#5;
   TraceIn_processLength[129] := BenchUut5.processLength;
   TraceIn_sensor1[129] := BenchUut5.sensor1;
   TraceIn_sensor2[129] := BenchUut5.sensor2;
   TraceIn_sensor3[129] := BenchUut5.sensor3;
   TraceIn_sensor4[129] := BenchUut5.sensor4;
   TraceIn_sensor5[129] := BenchUut5.sensor5;
   TraceIn_station1Start[129] := BenchUut5.station1Start;
   TraceIn_station2Complete[129] := BenchUut5.station2Complete;
   TraceIn_station3Complete[129] := BenchUut5.station3Complete;
   TraceIn_station4Complete[129] := BenchUut5.station4Complete;
   TraceIn_processSequence_1[129] := BenchUut5.processSequence[1];
   TraceIn_processSequence_2[129] := BenchUut5.processSequence[2];
   TraceIn_processSequence_3[129] := BenchUut5.processSequence[3];
   TraceIn_processSequence_4[129] := BenchUut5.processSequence[4];
   TraceIn_processSequence_5[129] := BenchUut5.processSequence[5];
   TraceIn_processSequence_6[129] := BenchUut5.processSequence[6];
   TraceIn_processSequence_7[129] := BenchUut5.processSequence[7];
   TraceIn_processSequence_8[129] := BenchUut5.processSequence[8];
   BenchUut5();
   TraceOut_conveyorLeft[129] := BenchUut5.conveyorLeft;
   TraceOut_conveyorRight[129] := BenchUut5.conveyorRight;
   BenchCalls := BenchCalls + 1;
 130:
   BenchUut5.processLength := USINT#8;
   BenchUut5.sensor1 := FALSE;
   BenchUut5.sensor2 := FALSE;
   BenchUut5.sensor3 := FALSE;
   BenchUut5.sensor4 := FALSE;
   BenchUut5.sensor5 := FALSE;
   BenchUut5.station1Start := FALSE;
   BenchUut5.station2Complete := FALSE;
   BenchUut5.station3Complete := FALSE;
   BenchUut5.station4Complete := FALSE;
   BenchUut5.processSequence[1] := USINT#2;
   BenchUut5.processSequence[2] := USINT#3;
   BenchUut5.processSequence[3] := USINT#4;
   BenchUut5.processSequence[4] := USINT#3;
   BenchUut5.processSequence[5] := USINT#2;
   BenchUut5.processSequence[6] := USINT#4;
   BenchUut5.processSequence[7] := USINT#3;
   BenchUut5.processSequence[8] := USINT#5;
   TraceIn_processLength[130] := BenchUut5.processLength;
   TraceIn_sensor1[130] := BenchUut5.sensor1;
   TraceIn_sensor2[130] := BenchUut5.sensor2;
   TraceIn_sensor3[130] := BenchUut5.sensor3;
   TraceIn_sensor4[130] := BenchUut5.sensor4;
   TraceIn_sensor5[130] := BenchUut5.sensor5;
   TraceIn_station1Start[130] := BenchUut5.station1Start;
   TraceIn_station2Complete[130] := BenchUut5.station2Complete;
   TraceIn_station3Complete[130] := BenchUut5.station3Complete;
   TraceIn_station4Complete[130] := BenchUut5.station4Complete;
   TraceIn_processSequence_1[130] := BenchUut5.processSequence[1];
   TraceIn_processSequence_2[130] := BenchUut5.processSequence[2];
   TraceIn_processSequence_3[130] := BenchUut5.processSequence[3];
   TraceIn_processSequence_4[130] := BenchUut5.processSequence[4];
   TraceIn_processSequence_5[130] := BenchUut5.processSequence[5];
   TraceIn_processSequence_6[130] := BenchUut5.processSequence[6];
   TraceIn_processSequence_7[130] := BenchUut5.processSequence[7];
   TraceIn_processSequence_8[130] := BenchUut5.processSequence[8];
   BenchUut5();
   TraceOut_conveyorLeft[130] := BenchUut5.conveyorLeft;
   TraceOut_conveyorRight[130] := BenchUut5.conveyorRight;
   BenchCalls := BenchCalls + 1;
 131:
   BenchUut5.processLength := USINT#8;
   BenchUut5.sensor1 := FALSE;
   BenchUut5.sensor2 := FALSE;
   BenchUut5.sensor3 := FALSE;
   BenchUut5.sensor4 := FALSE;
   BenchUut5.sensor5 := FALSE;
   BenchUut5.station1Start := FALSE;
   BenchUut5.station2Complete := FALSE;
   BenchUut5.station3Complete := FALSE;
   BenchUut5.station4Complete := FALSE;
   BenchUut5.processSequence[1] := USINT#2;
   BenchUut5.processSequence[2] := USINT#3;
   BenchUut5.processSequence[3] := USINT#4;
   BenchUut5.processSequence[4] := USINT#3;
   BenchUut5.processSequence[5] := USINT#2;
   BenchUut5.processSequence[6] := USINT#4;
   BenchUut5.processSequence[7] := USINT#3;
   BenchUut5.processSequence[8] := USINT#5;
   TraceIn_processLength[131] := BenchUut5.processLength;
   TraceIn_sensor1[131] := BenchUut5.sensor1;
   TraceIn_sensor2[131] := BenchUut5.sensor2;
   TraceIn_sensor3[131] := BenchUut5.sensor3;
   TraceIn_sensor4[131] := BenchUut5.sensor4;
   TraceIn_sensor5[131] := BenchUut5.sensor5;
   TraceIn_station1Start[131] := BenchUut5.station1Start;
   TraceIn_station2Complete[131] := BenchUut5.station2Complete;
   TraceIn_station3Complete[131] := BenchUut5.station3Complete;
   TraceIn_station4Complete[131] := BenchUut5.station4Complete;
   TraceIn_processSequence_1[131] := BenchUut5.processSequence[1];
   TraceIn_processSequence_2[131] := BenchUut5.processSequence[2];
   TraceIn_processSequence_3[131] := BenchUut5.processSequence[3];
   TraceIn_processSequence_4[131] := BenchUut5.processSequence[4];
   TraceIn_processSequence_5[131] := BenchUut5.processSequence[5];
   TraceIn_processSequence_6[131] := BenchUut5.processSequence[6];
   TraceIn_processSequence_7[131] := BenchUut5.processSequence[7];
   TraceIn_processSequence_8[131] := BenchUut5.processSequence[8];
   BenchUut5();
   TraceOut_conveyorLeft[131] := BenchUut5.conveyorLeft;
   TraceOut_conveyorRight[131] := BenchUut5.conveyorRight;
   BenchCalls := BenchCalls + 1;
 132:
   BenchUut5.processLength := USINT#8;
   BenchUut5.sensor1 := FALSE;
   BenchUut5.sensor2 := FALSE;
   BenchUut5.sensor3 := TRUE;
   BenchUut5.sensor4 := FALSE;
   BenchUut5.sensor5 := FALSE;
   BenchUut5.station1Start := FALSE;
   BenchUut5.station2Complete := FALSE;
   BenchUut5.station3Complete := FALSE;
   BenchUut5.station4Complete := FALSE;
   BenchUut5.processSequence[1] := USINT#2;
   BenchUut5.processSequence[2] := USINT#3;
   BenchUut5.processSequence[3] := USINT#4;
   BenchUut5.processSequence[4] := USINT#3;
   BenchUut5.processSequence[5] := USINT#2;
   BenchUut5.processSequence[6] := USINT#4;
   BenchUut5.processSequence[7] := USINT#3;
   BenchUut5.processSequence[8] := USINT#5;
   TraceIn_processLength[132] := BenchUut5.processLength;
   TraceIn_sensor1[132] := BenchUut5.sensor1;
   TraceIn_sensor2[132] := BenchUut5.sensor2;
   TraceIn_sensor3[132] := BenchUut5.sensor3;
   TraceIn_sensor4[132] := BenchUut5.sensor4;
   TraceIn_sensor5[132] := BenchUut5.sensor5;
   TraceIn_station1Start[132] := BenchUut5.station1Start;
   TraceIn_station2Complete[132] := BenchUut5.station2Complete;
   TraceIn_station3Complete[132] := BenchUut5.station3Complete;
   TraceIn_station4Complete[132] := BenchUut5.station4Complete;
   TraceIn_processSequence_1[132] := BenchUut5.processSequence[1];
   TraceIn_processSequence_2[132] := BenchUut5.processSequence[2];
   TraceIn_processSequence_3[132] := BenchUut5.processSequence[3];
   TraceIn_processSequence_4[132] := BenchUut5.processSequence[4];
   TraceIn_processSequence_5[132] := BenchUut5.processSequence[5];
   TraceIn_processSequence_6[132] := BenchUut5.processSequence[6];
   TraceIn_processSequence_7[132] := BenchUut5.processSequence[7];
   TraceIn_processSequence_8[132] := BenchUut5.processSequence[8];
   BenchUut5();
   TraceOut_conveyorLeft[132] := BenchUut5.conveyorLeft;
   TraceOut_conveyorRight[132] := BenchUut5.conveyorRight;
   BenchCalls := BenchCalls + 1;
 133:
   BenchUut5.processLength := USINT#8;
   BenchUut5.sensor1 := FALSE;
   BenchUut5.sensor2 := FALSE;
   BenchUut5.sensor3 := TRUE;
   BenchUut5.sensor4 := FALSE;
   BenchUut5.sensor5 := FALSE;
   BenchUut5.station1Start := FALSE;
   BenchUut5.station2Complete := FALSE;
   BenchUut5.station3Complete := FALSE;
   BenchUut5.station4Complete := FALSE;
   BenchUut5.processSequence[1] := USINT#2;
   BenchUut5.processSequence[2] := USINT#3;
   BenchUut5.processSequence[3] := USINT#4;
   BenchUut5.processSequence[4] := USINT#3;
   BenchUut5.processSequence[5] := USINT#2;
   BenchUut5.processSequence[6] := USINT#4;
   BenchUut5.processSequence[7] := USINT#3;
   BenchUut5.processSequence[8] := USINT#5;
   TraceIn_processLength[133] := BenchUut5.processLength;
   TraceIn_sensor1[133] := BenchUut5.sensor1;
   TraceIn_sensor2[133] := BenchUut5.sensor2;
   TraceIn_sensor3[133] := BenchUut5.sensor3;
   TraceIn_sensor4[133] := BenchUut5.sensor4;
   TraceIn_sensor5[133] := BenchUut5.sensor5;
   TraceIn_station1Start[133] := BenchUut5.station1Start;
   TraceIn_station2Complete[133] := BenchUut5.station2Complete;
   TraceIn_station3Complete[133] := BenchUut5.station3Complete;
   TraceIn_station4Complete[133] := BenchUut5.station4Complete;
   TraceIn_processSequence_1[133] := BenchUut5.processSequence[1];
   TraceIn_processSequence_2[133] := BenchUut5.processSequence[2];
   TraceIn_processSequence_3[133] := BenchUut5.processSequence[3];
   TraceIn_processSequence_4[133] := BenchUut5.processSequence[4];
   TraceIn_processSequence_5[133] := BenchUut5.processSequence[5];
   TraceIn_processSequence_6[133] := BenchUut5.processSequence[6];
   TraceIn_processSequence_7[133] := BenchUut5.processSequence[7];
   TraceIn_processSequence_8[133] := BenchUut5.processSequence[8];
   BenchUut5();
   TraceOut_conveyorLeft[133] := BenchUut5.conveyorLeft;
   TraceOut_conveyorRight[133] := BenchUut5.conveyorRight;
   BenchCalls := BenchCalls + 1;
 134:
   BenchUut5.processLength := USINT#8;
   BenchUut5.sensor1 := FALSE;
   BenchUut5.sensor2 := FALSE;
   BenchUut5.sensor3 := TRUE;
   BenchUut5.sensor4 := FALSE;
   BenchUut5.sensor5 := FALSE;
   BenchUut5.station1Start := FALSE;
   BenchUut5.station2Complete := FALSE;
   BenchUut5.station3Complete := FALSE;
   BenchUut5.station4Complete := FALSE;
   BenchUut5.processSequence[1] := USINT#2;
   BenchUut5.processSequence[2] := USINT#3;
   BenchUut5.processSequence[3] := USINT#4;
   BenchUut5.processSequence[4] := USINT#3;
   BenchUut5.processSequence[5] := USINT#2;
   BenchUut5.processSequence[6] := USINT#4;
   BenchUut5.processSequence[7] := USINT#3;
   BenchUut5.processSequence[8] := USINT#5;
   TraceIn_processLength[134] := BenchUut5.processLength;
   TraceIn_sensor1[134] := BenchUut5.sensor1;
   TraceIn_sensor2[134] := BenchUut5.sensor2;
   TraceIn_sensor3[134] := BenchUut5.sensor3;
   TraceIn_sensor4[134] := BenchUut5.sensor4;
   TraceIn_sensor5[134] := BenchUut5.sensor5;
   TraceIn_station1Start[134] := BenchUut5.station1Start;
   TraceIn_station2Complete[134] := BenchUut5.station2Complete;
   TraceIn_station3Complete[134] := BenchUut5.station3Complete;
   TraceIn_station4Complete[134] := BenchUut5.station4Complete;
   TraceIn_processSequence_1[134] := BenchUut5.processSequence[1];
   TraceIn_processSequence_2[134] := BenchUut5.processSequence[2];
   TraceIn_processSequence_3[134] := BenchUut5.processSequence[3];
   TraceIn_processSequence_4[134] := BenchUut5.processSequence[4];
   TraceIn_processSequence_5[134] := BenchUut5.processSequence[5];
   TraceIn_processSequence_6[134] := BenchUut5.processSequence[6];
   TraceIn_processSequence_7[134] := BenchUut5.processSequence[7];
   TraceIn_processSequence_8[134] := BenchUut5.processSequence[8];
   BenchUut5();
   TraceOut_conveyorLeft[134] := BenchUut5.conveyorLeft;
   TraceOut_conveyorRight[134] := BenchUut5.conveyorRight;
   BenchCalls := BenchCalls + 1;
 135:
   BenchUut5.processLength := USINT#8;
   BenchUut5.sensor1 := FALSE;
   BenchUut5.sensor2 := FALSE;
   BenchUut5.sensor3 := TRUE;
   BenchUut5.sensor4 := FALSE;
   BenchUut5.sensor5 := FALSE;
   BenchUut5.station1Start := FALSE;
   BenchUut5.station2Complete := FALSE;
   BenchUut5.station3Complete := TRUE;
   BenchUut5.station4Complete := FALSE;
   BenchUut5.processSequence[1] := USINT#2;
   BenchUut5.processSequence[2] := USINT#3;
   BenchUut5.processSequence[3] := USINT#4;
   BenchUut5.processSequence[4] := USINT#3;
   BenchUut5.processSequence[5] := USINT#2;
   BenchUut5.processSequence[6] := USINT#4;
   BenchUut5.processSequence[7] := USINT#3;
   BenchUut5.processSequence[8] := USINT#5;
   TraceIn_processLength[135] := BenchUut5.processLength;
   TraceIn_sensor1[135] := BenchUut5.sensor1;
   TraceIn_sensor2[135] := BenchUut5.sensor2;
   TraceIn_sensor3[135] := BenchUut5.sensor3;
   TraceIn_sensor4[135] := BenchUut5.sensor4;
   TraceIn_sensor5[135] := BenchUut5.sensor5;
   TraceIn_station1Start[135] := BenchUut5.station1Start;
   TraceIn_station2Complete[135] := BenchUut5.station2Complete;
   TraceIn_station3Complete[135] := BenchUut5.station3Complete;
   TraceIn_station4Complete[135] := BenchUut5.station4Complete;
   TraceIn_processSequence_1[135] := BenchUut5.processSequence[1];
   TraceIn_processSequence_2[135] := BenchUut5.processSequence[2];
   TraceIn_processSequence_3[135] := BenchUut5.processSequence[3];
   TraceIn_processSequence_4[135] := BenchUut5.processSequence[4];
   TraceIn_processSequence_5[135] := BenchUut5.processSequence[5];
   TraceIn_processSequence_6[135] := BenchUut5.processSequence[6];
   TraceIn_processSequence_7[135] := BenchUut5.processSequence[7];
   TraceIn_processSequence_8[135] := BenchUut5.processSequence[8];
   BenchUut5();
   TraceOut_conveyorLeft[135] := BenchUut5.conveyorLeft;
   TraceOut_conveyorRight[135] := BenchUut5.conveyorRight;
   BenchCalls := BenchCalls + 1;
 136:
   BenchUut5.processLength := USINT#8;
   BenchUut5.sensor1 := FALSE;
   BenchUut5.sensor2 := FALSE;
   BenchUut5.sensor3 := FALSE;
   BenchUut5.sensor4 := FALSE;
   BenchUut5.sensor5 := FALSE;
   BenchUut5.station1Start := FALSE;
   BenchUut5.station2Complete := FALSE;
   BenchUut5.station3Complete := FALSE;
   BenchUut5.station4Complete := FALSE;
   BenchUut5.processSequence[1] := USINT#2;
   BenchUut5.processSequence[2] := USINT#3;
   BenchUut5.processSequence[3] := USINT#4;
   BenchUut5.processSequence[4] := USINT#3;
   BenchUut5.processSequence[5] := USINT#2;
   BenchUut5.processSequence[6] := USINT#4;
   BenchUut5.processSequence[7] := USINT#3;
   BenchUut5.processSequence[8] := USINT#5;
   TraceIn_processLength[136] := BenchUut5.processLength;
   TraceIn_sensor1[136] := BenchUut5.sensor1;
   TraceIn_sensor2[136] := BenchUut5.sensor2;
   TraceIn_sensor3[136] := BenchUut5.sensor3;
   TraceIn_sensor4[136] := BenchUut5.sensor4;
   TraceIn_sensor5[136] := BenchUut5.sensor5;
   TraceIn_station1Start[136] := BenchUut5.station1Start;
   TraceIn_station2Complete[136] := BenchUut5.station2Complete;
   TraceIn_station3Complete[136] := BenchUut5.station3Complete;
   TraceIn_station4Complete[136] := BenchUut5.station4Complete;
   TraceIn_processSequence_1[136] := BenchUut5.processSequence[1];
   TraceIn_processSequence_2[136] := BenchUut5.processSequence[2];
   TraceIn_processSequence_3[136] := BenchUut5.processSequence[3];
   TraceIn_processSequence_4[136] := BenchUut5.processSequence[4];
   TraceIn_processSequence_5[136] := BenchUut5.processSequence[5];
   TraceIn_processSequence_6[136] := BenchUut5.processSequence[6];
   TraceIn_processSequence_7[136] := BenchUut5.processSequence[7];
   TraceIn_processSequence_8[136] := BenchUut5.processSequence[8];
   BenchUut5();
   TraceOut_conveyorLeft[136] := BenchUut5.conveyorLeft;
   TraceOut_conveyorRight[136] := BenchUut5.conveyorRight;
   BenchCalls := BenchCalls + 1;
 137:
   BenchUut5.processLength := USINT#8;
   BenchUut5.sensor1 := FALSE;
   BenchUut5.sensor2 := FALSE;
   BenchUut5.sensor3 := FALSE;
   BenchUut5.sensor4 := FALSE;
   BenchUut5.sensor5 := FALSE;
   BenchUut5.station1Start := FALSE;
   BenchUut5.station2Complete := FALSE;
   BenchUut5.station3Complete := FALSE;
   BenchUut5.station4Complete := FALSE;
   BenchUut5.processSequence[1] := USINT#2;
   BenchUut5.processSequence[2] := USINT#3;
   BenchUut5.processSequence[3] := USINT#4;
   BenchUut5.processSequence[4] := USINT#3;
   BenchUut5.processSequence[5] := USINT#2;
   BenchUut5.processSequence[6] := USINT#4;
   BenchUut5.processSequence[7] := USINT#3;
   BenchUut5.processSequence[8] := USINT#5;
   TraceIn_processLength[137] := BenchUut5.processLength;
   TraceIn_sensor1[137] := BenchUut5.sensor1;
   TraceIn_sensor2[137] := BenchUut5.sensor2;
   TraceIn_sensor3[137] := BenchUut5.sensor3;
   TraceIn_sensor4[137] := BenchUut5.sensor4;
   TraceIn_sensor5[137] := BenchUut5.sensor5;
   TraceIn_station1Start[137] := BenchUut5.station1Start;
   TraceIn_station2Complete[137] := BenchUut5.station2Complete;
   TraceIn_station3Complete[137] := BenchUut5.station3Complete;
   TraceIn_station4Complete[137] := BenchUut5.station4Complete;
   TraceIn_processSequence_1[137] := BenchUut5.processSequence[1];
   TraceIn_processSequence_2[137] := BenchUut5.processSequence[2];
   TraceIn_processSequence_3[137] := BenchUut5.processSequence[3];
   TraceIn_processSequence_4[137] := BenchUut5.processSequence[4];
   TraceIn_processSequence_5[137] := BenchUut5.processSequence[5];
   TraceIn_processSequence_6[137] := BenchUut5.processSequence[6];
   TraceIn_processSequence_7[137] := BenchUut5.processSequence[7];
   TraceIn_processSequence_8[137] := BenchUut5.processSequence[8];
   BenchUut5();
   TraceOut_conveyorLeft[137] := BenchUut5.conveyorLeft;
   TraceOut_conveyorRight[137] := BenchUut5.conveyorRight;
   BenchCalls := BenchCalls + 1;
 138:
   BenchUut5.processLength := USINT#8;
   BenchUut5.sensor1 := FALSE;
   BenchUut5.sensor2 := FALSE;
   BenchUut5.sensor3 := FALSE;
   BenchUut5.sensor4 := FALSE;
   BenchUut5.sensor5 := TRUE;
   BenchUut5.station1Start := FALSE;
   BenchUut5.station2Complete := FALSE;
   BenchUut5.station3Complete := FALSE;
   BenchUut5.station4Complete := FALSE;
   BenchUut5.processSequence[1] := USINT#2;
   BenchUut5.processSequence[2] := USINT#3;
   BenchUut5.processSequence[3] := USINT#4;
   BenchUut5.processSequence[4] := USINT#3;
   BenchUut5.processSequence[5] := USINT#2;
   BenchUut5.processSequence[6] := USINT#4;
   BenchUut5.processSequence[7] := USINT#3;
   BenchUut5.processSequence[8] := USINT#5;
   TraceIn_processLength[138] := BenchUut5.processLength;
   TraceIn_sensor1[138] := BenchUut5.sensor1;
   TraceIn_sensor2[138] := BenchUut5.sensor2;
   TraceIn_sensor3[138] := BenchUut5.sensor3;
   TraceIn_sensor4[138] := BenchUut5.sensor4;
   TraceIn_sensor5[138] := BenchUut5.sensor5;
   TraceIn_station1Start[138] := BenchUut5.station1Start;
   TraceIn_station2Complete[138] := BenchUut5.station2Complete;
   TraceIn_station3Complete[138] := BenchUut5.station3Complete;
   TraceIn_station4Complete[138] := BenchUut5.station4Complete;
   TraceIn_processSequence_1[138] := BenchUut5.processSequence[1];
   TraceIn_processSequence_2[138] := BenchUut5.processSequence[2];
   TraceIn_processSequence_3[138] := BenchUut5.processSequence[3];
   TraceIn_processSequence_4[138] := BenchUut5.processSequence[4];
   TraceIn_processSequence_5[138] := BenchUut5.processSequence[5];
   TraceIn_processSequence_6[138] := BenchUut5.processSequence[6];
   TraceIn_processSequence_7[138] := BenchUut5.processSequence[7];
   TraceIn_processSequence_8[138] := BenchUut5.processSequence[8];
   BenchUut5();
   TraceOut_conveyorLeft[138] := BenchUut5.conveyorLeft;
   TraceOut_conveyorRight[138] := BenchUut5.conveyorRight;
   BenchCalls := BenchCalls + 1;
 139:
   BenchUut6.processLength := USINT#2;
   BenchUut6.sensor1 := FALSE;
   BenchUut6.sensor2 := FALSE;
   BenchUut6.sensor3 := FALSE;
   BenchUut6.sensor4 := FALSE;
   BenchUut6.sensor5 := FALSE;
   BenchUut6.station1Start := FALSE;
   BenchUut6.station2Complete := FALSE;
   BenchUut6.station3Complete := FALSE;
   BenchUut6.station4Complete := FALSE;
   BenchUut6.processSequence[1] := USINT#3;
   BenchUut6.processSequence[2] := USINT#5;
   BenchUut6.processSequence[3] := USINT#0;
   BenchUut6.processSequence[4] := USINT#0;
   BenchUut6.processSequence[5] := USINT#0;
   BenchUut6.processSequence[6] := USINT#0;
   BenchUut6.processSequence[7] := USINT#0;
   BenchUut6.processSequence[8] := USINT#0;
   TraceIn_processLength[139] := BenchUut6.processLength;
   TraceIn_sensor1[139] := BenchUut6.sensor1;
   TraceIn_sensor2[139] := BenchUut6.sensor2;
   TraceIn_sensor3[139] := BenchUut6.sensor3;
   TraceIn_sensor4[139] := BenchUut6.sensor4;
   TraceIn_sensor5[139] := BenchUut6.sensor5;
   TraceIn_station1Start[139] := BenchUut6.station1Start;
   TraceIn_station2Complete[139] := BenchUut6.station2Complete;
   TraceIn_station3Complete[139] := BenchUut6.station3Complete;
   TraceIn_station4Complete[139] := BenchUut6.station4Complete;
   TraceIn_processSequence_1[139] := BenchUut6.processSequence[1];
   TraceIn_processSequence_2[139] := BenchUut6.processSequence[2];
   TraceIn_processSequence_3[139] := BenchUut6.processSequence[3];
   TraceIn_processSequence_4[139] := BenchUut6.processSequence[4];
   TraceIn_processSequence_5[139] := BenchUut6.processSequence[5];
   TraceIn_processSequence_6[139] := BenchUut6.processSequence[6];
   TraceIn_processSequence_7[139] := BenchUut6.processSequence[7];
   TraceIn_processSequence_8[139] := BenchUut6.processSequence[8];
   BenchUut6();
   TraceOut_conveyorLeft[139] := BenchUut6.conveyorLeft;
   TraceOut_conveyorRight[139] := BenchUut6.conveyorRight;
   BenchCalls := BenchCalls + 1;
 140:
   BenchUut6.processLength := USINT#2;
   BenchUut6.sensor1 := FALSE;
   BenchUut6.sensor2 := FALSE;
   BenchUut6.sensor3 := FALSE;
   BenchUut6.sensor4 := FALSE;
   BenchUut6.sensor5 := FALSE;
   BenchUut6.station1Start := TRUE;
   BenchUut6.station2Complete := FALSE;
   BenchUut6.station3Complete := FALSE;
   BenchUut6.station4Complete := FALSE;
   BenchUut6.processSequence[1] := USINT#3;
   BenchUut6.processSequence[2] := USINT#5;
   BenchUut6.processSequence[3] := USINT#0;
   BenchUut6.processSequence[4] := USINT#0;
   BenchUut6.processSequence[5] := USINT#0;
   BenchUut6.processSequence[6] := USINT#0;
   BenchUut6.processSequence[7] := USINT#0;
   BenchUut6.processSequence[8] := USINT#0;
   TraceIn_processLength[140] := BenchUut6.processLength;
   TraceIn_sensor1[140] := BenchUut6.sensor1;
   TraceIn_sensor2[140] := BenchUut6.sensor2;
   TraceIn_sensor3[140] := BenchUut6.sensor3;
   TraceIn_sensor4[140] := BenchUut6.sensor4;
   TraceIn_sensor5[140] := BenchUut6.sensor5;
   TraceIn_station1Start[140] := BenchUut6.station1Start;
   TraceIn_station2Complete[140] := BenchUut6.station2Complete;
   TraceIn_station3Complete[140] := BenchUut6.station3Complete;
   TraceIn_station4Complete[140] := BenchUut6.station4Complete;
   TraceIn_processSequence_1[140] := BenchUut6.processSequence[1];
   TraceIn_processSequence_2[140] := BenchUut6.processSequence[2];
   TraceIn_processSequence_3[140] := BenchUut6.processSequence[3];
   TraceIn_processSequence_4[140] := BenchUut6.processSequence[4];
   TraceIn_processSequence_5[140] := BenchUut6.processSequence[5];
   TraceIn_processSequence_6[140] := BenchUut6.processSequence[6];
   TraceIn_processSequence_7[140] := BenchUut6.processSequence[7];
   TraceIn_processSequence_8[140] := BenchUut6.processSequence[8];
   BenchUut6();
   TraceOut_conveyorLeft[140] := BenchUut6.conveyorLeft;
   TraceOut_conveyorRight[140] := BenchUut6.conveyorRight;
   BenchCalls := BenchCalls + 1;
 141:
   BenchUut6.processLength := USINT#2;
   BenchUut6.sensor1 := TRUE;
   BenchUut6.sensor2 := FALSE;
   BenchUut6.sensor3 := FALSE;
   BenchUut6.sensor4 := FALSE;
   BenchUut6.sensor5 := FALSE;
   BenchUut6.station1Start := TRUE;
   BenchUut6.station2Complete := FALSE;
   BenchUut6.station3Complete := FALSE;
   BenchUut6.station4Complete := FALSE;
   BenchUut6.processSequence[1] := USINT#3;
   BenchUut6.processSequence[2] := USINT#5;
   BenchUut6.processSequence[3] := USINT#0;
   BenchUut6.processSequence[4] := USINT#0;
   BenchUut6.processSequence[5] := USINT#0;
   BenchUut6.processSequence[6] := USINT#0;
   BenchUut6.processSequence[7] := USINT#0;
   BenchUut6.processSequence[8] := USINT#0;
   TraceIn_processLength[141] := BenchUut6.processLength;
   TraceIn_sensor1[141] := BenchUut6.sensor1;
   TraceIn_sensor2[141] := BenchUut6.sensor2;
   TraceIn_sensor3[141] := BenchUut6.sensor3;
   TraceIn_sensor4[141] := BenchUut6.sensor4;
   TraceIn_sensor5[141] := BenchUut6.sensor5;
   TraceIn_station1Start[141] := BenchUut6.station1Start;
   TraceIn_station2Complete[141] := BenchUut6.station2Complete;
   TraceIn_station3Complete[141] := BenchUut6.station3Complete;
   TraceIn_station4Complete[141] := BenchUut6.station4Complete;
   TraceIn_processSequence_1[141] := BenchUut6.processSequence[1];
   TraceIn_processSequence_2[141] := BenchUut6.processSequence[2];
   TraceIn_processSequence_3[141] := BenchUut6.processSequence[3];
   TraceIn_processSequence_4[141] := BenchUut6.processSequence[4];
   TraceIn_processSequence_5[141] := BenchUut6.processSequence[5];
   TraceIn_processSequence_6[141] := BenchUut6.processSequence[6];
   TraceIn_processSequence_7[141] := BenchUut6.processSequence[7];
   TraceIn_processSequence_8[141] := BenchUut6.processSequence[8];
   BenchUut6();
   TraceOut_conveyorLeft[141] := BenchUut6.conveyorLeft;
   TraceOut_conveyorRight[141] := BenchUut6.conveyorRight;
   BenchCalls := BenchCalls + 1;
 142:
   BenchUut6.processLength := USINT#2;
   BenchUut6.sensor1 := TRUE;
   BenchUut6.sensor2 := FALSE;
   BenchUut6.sensor3 := FALSE;
   BenchUut6.sensor4 := FALSE;
   BenchUut6.sensor5 := FALSE;
   BenchUut6.station1Start := FALSE;
   BenchUut6.station2Complete := FALSE;
   BenchUut6.station3Complete := FALSE;
   BenchUut6.station4Complete := FALSE;
   BenchUut6.processSequence[1] := USINT#3;
   BenchUut6.processSequence[2] := USINT#5;
   BenchUut6.processSequence[3] := USINT#0;
   BenchUut6.processSequence[4] := USINT#0;
   BenchUut6.processSequence[5] := USINT#0;
   BenchUut6.processSequence[6] := USINT#0;
   BenchUut6.processSequence[7] := USINT#0;
   BenchUut6.processSequence[8] := USINT#0;
   TraceIn_processLength[142] := BenchUut6.processLength;
   TraceIn_sensor1[142] := BenchUut6.sensor1;
   TraceIn_sensor2[142] := BenchUut6.sensor2;
   TraceIn_sensor3[142] := BenchUut6.sensor3;
   TraceIn_sensor4[142] := BenchUut6.sensor4;
   TraceIn_sensor5[142] := BenchUut6.sensor5;
   TraceIn_station1Start[142] := BenchUut6.station1Start;
   TraceIn_station2Complete[142] := BenchUut6.station2Complete;
   TraceIn_station3Complete[142] := BenchUut6.station3Complete;
   TraceIn_station4Complete[142] := BenchUut6.station4Complete;
   TraceIn_processSequence_1[142] := BenchUut6.processSequence[1];
   TraceIn_processSequence_2[142] := BenchUut6.processSequence[2];
   TraceIn_processSequence_3[142] := BenchUut6.processSequence[3];
   TraceIn_processSequence_4[142] := BenchUut6.processSequence[4];
   TraceIn_processSequence_5[142] := BenchUut6.processSequence[5];
   TraceIn_processSequence_6[142] := BenchUut6.processSequence[6];
   TraceIn_processSequence_7[142] := BenchUut6.processSequence[7];
   TraceIn_processSequence_8[142] := BenchUut6.processSequence[8];
   BenchUut6();
   TraceOut_conveyorLeft[142] := BenchUut6.conveyorLeft;
   TraceOut_conveyorRight[142] := BenchUut6.conveyorRight;
   BenchCalls := BenchCalls + 1;
 143:
   BenchUut6.processLength := USINT#2;
   BenchUut6.sensor1 := TRUE;
   BenchUut6.sensor2 := FALSE;
   BenchUut6.sensor3 := FALSE;
   BenchUut6.sensor4 := FALSE;
   BenchUut6.sensor5 := FALSE;
   BenchUut6.station1Start := TRUE;
   BenchUut6.station2Complete := FALSE;
   BenchUut6.station3Complete := FALSE;
   BenchUut6.station4Complete := FALSE;
   BenchUut6.processSequence[1] := USINT#3;
   BenchUut6.processSequence[2] := USINT#5;
   BenchUut6.processSequence[3] := USINT#0;
   BenchUut6.processSequence[4] := USINT#0;
   BenchUut6.processSequence[5] := USINT#0;
   BenchUut6.processSequence[6] := USINT#0;
   BenchUut6.processSequence[7] := USINT#0;
   BenchUut6.processSequence[8] := USINT#0;
   TraceIn_processLength[143] := BenchUut6.processLength;
   TraceIn_sensor1[143] := BenchUut6.sensor1;
   TraceIn_sensor2[143] := BenchUut6.sensor2;
   TraceIn_sensor3[143] := BenchUut6.sensor3;
   TraceIn_sensor4[143] := BenchUut6.sensor4;
   TraceIn_sensor5[143] := BenchUut6.sensor5;
   TraceIn_station1Start[143] := BenchUut6.station1Start;
   TraceIn_station2Complete[143] := BenchUut6.station2Complete;
   TraceIn_station3Complete[143] := BenchUut6.station3Complete;
   TraceIn_station4Complete[143] := BenchUut6.station4Complete;
   TraceIn_processSequence_1[143] := BenchUut6.processSequence[1];
   TraceIn_processSequence_2[143] := BenchUut6.processSequence[2];
   TraceIn_processSequence_3[143] := BenchUut6.processSequence[3];
   TraceIn_processSequence_4[143] := BenchUut6.processSequence[4];
   TraceIn_processSequence_5[143] := BenchUut6.processSequence[5];
   TraceIn_processSequence_6[143] := BenchUut6.processSequence[6];
   TraceIn_processSequence_7[143] := BenchUut6.processSequence[7];
   TraceIn_processSequence_8[143] := BenchUut6.processSequence[8];
   BenchUut6();
   TraceOut_conveyorLeft[143] := BenchUut6.conveyorLeft;
   TraceOut_conveyorRight[143] := BenchUut6.conveyorRight;
   BenchCalls := BenchCalls + 1;
 144:
   BenchUut6.processLength := USINT#2;
   BenchUut6.sensor1 := FALSE;
   BenchUut6.sensor2 := FALSE;
   BenchUut6.sensor3 := TRUE;
   BenchUut6.sensor4 := FALSE;
   BenchUut6.sensor5 := FALSE;
   BenchUut6.station1Start := TRUE;
   BenchUut6.station2Complete := FALSE;
   BenchUut6.station3Complete := FALSE;
   BenchUut6.station4Complete := FALSE;
   BenchUut6.processSequence[1] := USINT#3;
   BenchUut6.processSequence[2] := USINT#5;
   BenchUut6.processSequence[3] := USINT#0;
   BenchUut6.processSequence[4] := USINT#0;
   BenchUut6.processSequence[5] := USINT#0;
   BenchUut6.processSequence[6] := USINT#0;
   BenchUut6.processSequence[7] := USINT#0;
   BenchUut6.processSequence[8] := USINT#0;
   TraceIn_processLength[144] := BenchUut6.processLength;
   TraceIn_sensor1[144] := BenchUut6.sensor1;
   TraceIn_sensor2[144] := BenchUut6.sensor2;
   TraceIn_sensor3[144] := BenchUut6.sensor3;
   TraceIn_sensor4[144] := BenchUut6.sensor4;
   TraceIn_sensor5[144] := BenchUut6.sensor5;
   TraceIn_station1Start[144] := BenchUut6.station1Start;
   TraceIn_station2Complete[144] := BenchUut6.station2Complete;
   TraceIn_station3Complete[144] := BenchUut6.station3Complete;
   TraceIn_station4Complete[144] := BenchUut6.station4Complete;
   TraceIn_processSequence_1[144] := BenchUut6.processSequence[1];
   TraceIn_processSequence_2[144] := BenchUut6.processSequence[2];
   TraceIn_processSequence_3[144] := BenchUut6.processSequence[3];
   TraceIn_processSequence_4[144] := BenchUut6.processSequence[4];
   TraceIn_processSequence_5[144] := BenchUut6.processSequence[5];
   TraceIn_processSequence_6[144] := BenchUut6.processSequence[6];
   TraceIn_processSequence_7[144] := BenchUut6.processSequence[7];
   TraceIn_processSequence_8[144] := BenchUut6.processSequence[8];
   BenchUut6();
   TraceOut_conveyorLeft[144] := BenchUut6.conveyorLeft;
   TraceOut_conveyorRight[144] := BenchUut6.conveyorRight;
   BenchCalls := BenchCalls + 1;
 145:
   BenchUut6.processLength := USINT#2;
   BenchUut6.sensor1 := FALSE;
   BenchUut6.sensor2 := FALSE;
   BenchUut6.sensor3 := TRUE;
   BenchUut6.sensor4 := FALSE;
   BenchUut6.sensor5 := FALSE;
   BenchUut6.station1Start := FALSE;
   BenchUut6.station2Complete := FALSE;
   BenchUut6.station3Complete := TRUE;
   BenchUut6.station4Complete := FALSE;
   BenchUut6.processSequence[1] := USINT#3;
   BenchUut6.processSequence[2] := USINT#5;
   BenchUut6.processSequence[3] := USINT#0;
   BenchUut6.processSequence[4] := USINT#0;
   BenchUut6.processSequence[5] := USINT#0;
   BenchUut6.processSequence[6] := USINT#0;
   BenchUut6.processSequence[7] := USINT#0;
   BenchUut6.processSequence[8] := USINT#0;
   TraceIn_processLength[145] := BenchUut6.processLength;
   TraceIn_sensor1[145] := BenchUut6.sensor1;
   TraceIn_sensor2[145] := BenchUut6.sensor2;
   TraceIn_sensor3[145] := BenchUut6.sensor3;
   TraceIn_sensor4[145] := BenchUut6.sensor4;
   TraceIn_sensor5[145] := BenchUut6.sensor5;
   TraceIn_station1Start[145] := BenchUut6.station1Start;
   TraceIn_station2Complete[145] := BenchUut6.station2Complete;
   TraceIn_station3Complete[145] := BenchUut6.station3Complete;
   TraceIn_station4Complete[145] := BenchUut6.station4Complete;
   TraceIn_processSequence_1[145] := BenchUut6.processSequence[1];
   TraceIn_processSequence_2[145] := BenchUut6.processSequence[2];
   TraceIn_processSequence_3[145] := BenchUut6.processSequence[3];
   TraceIn_processSequence_4[145] := BenchUut6.processSequence[4];
   TraceIn_processSequence_5[145] := BenchUut6.processSequence[5];
   TraceIn_processSequence_6[145] := BenchUut6.processSequence[6];
   TraceIn_processSequence_7[145] := BenchUut6.processSequence[7];
   TraceIn_processSequence_8[145] := BenchUut6.processSequence[8];
   BenchUut6();
   TraceOut_conveyorLeft[145] := BenchUut6.conveyorLeft;
   TraceOut_conveyorRight[145] := BenchUut6.conveyorRight;
   BenchCalls := BenchCalls + 1;
 146:
   BenchUut6.processLength := USINT#2;
   BenchUut6.sensor1 := FALSE;
   BenchUut6.sensor2 := FALSE;
   BenchUut6.sensor3 := FALSE;
   BenchUut6.sensor4 := FALSE;
   BenchUut6.sensor5 := TRUE;
   BenchUut6.station1Start := FALSE;
   BenchUut6.station2Complete := FALSE;
   BenchUut6.station3Complete := FALSE;
   BenchUut6.station4Complete := FALSE;
   BenchUut6.processSequence[1] := USINT#3;
   BenchUut6.processSequence[2] := USINT#5;
   BenchUut6.processSequence[3] := USINT#0;
   BenchUut6.processSequence[4] := USINT#0;
   BenchUut6.processSequence[5] := USINT#0;
   BenchUut6.processSequence[6] := USINT#0;
   BenchUut6.processSequence[7] := USINT#0;
   BenchUut6.processSequence[8] := USINT#0;
   TraceIn_processLength[146] := BenchUut6.processLength;
   TraceIn_sensor1[146] := BenchUut6.sensor1;
   TraceIn_sensor2[146] := BenchUut6.sensor2;
   TraceIn_sensor3[146] := BenchUut6.sensor3;
   TraceIn_sensor4[146] := BenchUut6.sensor4;
   TraceIn_sensor5[146] := BenchUut6.sensor5;
   TraceIn_station1Start[146] := BenchUut6.station1Start;
   TraceIn_station2Complete[146] := BenchUut6.station2Complete;
   TraceIn_station3Complete[146] := BenchUut6.station3Complete;
   TraceIn_station4Complete[146] := BenchUut6.station4Complete;
   TraceIn_processSequence_1[146] := BenchUut6.processSequence[1];
   TraceIn_processSequence_2[146] := BenchUut6.processSequence[2];
   TraceIn_processSequence_3[146] := BenchUut6.processSequence[3];
   TraceIn_processSequence_4[146] := BenchUut6.processSequence[4];
   TraceIn_processSequence_5[146] := BenchUut6.processSequence[5];
   TraceIn_processSequence_6[146] := BenchUut6.processSequence[6];
   TraceIn_processSequence_7[146] := BenchUut6.processSequence[7];
   TraceIn_processSequence_8[146] := BenchUut6.processSequence[8];
   BenchUut6();
   TraceOut_conveyorLeft[146] := BenchUut6.conveyorLeft;
   TraceOut_conveyorRight[146] := BenchUut6.conveyorRight;
   BenchCalls := BenchCalls + 1;
 147:
   BenchUut6.processLength := USINT#2;
   BenchUut6.sensor1 := TRUE;
   BenchUut6.sensor2 := FALSE;
   BenchUut6.sensor3 := FALSE;
   BenchUut6.sensor4 := FALSE;
   BenchUut6.sensor5 := FALSE;
   BenchUut6.station1Start := TRUE;
   BenchUut6.station2Complete := FALSE;
   BenchUut6.station3Complete := FALSE;
   BenchUut6.station4Complete := FALSE;
   BenchUut6.processSequence[1] := USINT#3;
   BenchUut6.processSequence[2] := USINT#5;
   BenchUut6.processSequence[3] := USINT#0;
   BenchUut6.processSequence[4] := USINT#0;
   BenchUut6.processSequence[5] := USINT#0;
   BenchUut6.processSequence[6] := USINT#0;
   BenchUut6.processSequence[7] := USINT#0;
   BenchUut6.processSequence[8] := USINT#0;
   TraceIn_processLength[147] := BenchUut6.processLength;
   TraceIn_sensor1[147] := BenchUut6.sensor1;
   TraceIn_sensor2[147] := BenchUut6.sensor2;
   TraceIn_sensor3[147] := BenchUut6.sensor3;
   TraceIn_sensor4[147] := BenchUut6.sensor4;
   TraceIn_sensor5[147] := BenchUut6.sensor5;
   TraceIn_station1Start[147] := BenchUut6.station1Start;
   TraceIn_station2Complete[147] := BenchUut6.station2Complete;
   TraceIn_station3Complete[147] := BenchUut6.station3Complete;
   TraceIn_station4Complete[147] := BenchUut6.station4Complete;
   TraceIn_processSequence_1[147] := BenchUut6.processSequence[1];
   TraceIn_processSequence_2[147] := BenchUut6.processSequence[2];
   TraceIn_processSequence_3[147] := BenchUut6.processSequence[3];
   TraceIn_processSequence_4[147] := BenchUut6.processSequence[4];
   TraceIn_processSequence_5[147] := BenchUut6.processSequence[5];
   TraceIn_processSequence_6[147] := BenchUut6.processSequence[6];
   TraceIn_processSequence_7[147] := BenchUut6.processSequence[7];
   TraceIn_processSequence_8[147] := BenchUut6.processSequence[8];
   BenchUut6();
   TraceOut_conveyorLeft[147] := BenchUut6.conveyorLeft;
   TraceOut_conveyorRight[147] := BenchUut6.conveyorRight;
   BenchCalls := BenchCalls + 1;
 148:
   BenchUut7.processLength := USINT#5;
   BenchUut7.sensor1 := FALSE;
   BenchUut7.sensor2 := FALSE;
   BenchUut7.sensor3 := FALSE;
   BenchUut7.sensor4 := FALSE;
   BenchUut7.sensor5 := FALSE;
   BenchUut7.station1Start := FALSE;
   BenchUut7.station2Complete := FALSE;
   BenchUut7.station3Complete := FALSE;
   BenchUut7.station4Complete := FALSE;
   BenchUut7.processSequence[1] := USINT#2;
   BenchUut7.processSequence[2] := USINT#2;
   BenchUut7.processSequence[3] := USINT#3;
   BenchUut7.processSequence[4] := USINT#3;
   BenchUut7.processSequence[5] := USINT#5;
   BenchUut7.processSequence[6] := USINT#0;
   BenchUut7.processSequence[7] := USINT#0;
   BenchUut7.processSequence[8] := USINT#0;
   TraceIn_processLength[148] := BenchUut7.processLength;
   TraceIn_sensor1[148] := BenchUut7.sensor1;
   TraceIn_sensor2[148] := BenchUut7.sensor2;
   TraceIn_sensor3[148] := BenchUut7.sensor3;
   TraceIn_sensor4[148] := BenchUut7.sensor4;
   TraceIn_sensor5[148] := BenchUut7.sensor5;
   TraceIn_station1Start[148] := BenchUut7.station1Start;
   TraceIn_station2Complete[148] := BenchUut7.station2Complete;
   TraceIn_station3Complete[148] := BenchUut7.station3Complete;
   TraceIn_station4Complete[148] := BenchUut7.station4Complete;
   TraceIn_processSequence_1[148] := BenchUut7.processSequence[1];
   TraceIn_processSequence_2[148] := BenchUut7.processSequence[2];
   TraceIn_processSequence_3[148] := BenchUut7.processSequence[3];
   TraceIn_processSequence_4[148] := BenchUut7.processSequence[4];
   TraceIn_processSequence_5[148] := BenchUut7.processSequence[5];
   TraceIn_processSequence_6[148] := BenchUut7.processSequence[6];
   TraceIn_processSequence_7[148] := BenchUut7.processSequence[7];
   TraceIn_processSequence_8[148] := BenchUut7.processSequence[8];
   BenchUut7();
   TraceOut_conveyorLeft[148] := BenchUut7.conveyorLeft;
   TraceOut_conveyorRight[148] := BenchUut7.conveyorRight;
   BenchCalls := BenchCalls + 1;
 149:
   BenchUut7.processLength := USINT#5;
   BenchUut7.sensor1 := TRUE;
   BenchUut7.sensor2 := FALSE;
   BenchUut7.sensor3 := FALSE;
   BenchUut7.sensor4 := FALSE;
   BenchUut7.sensor5 := FALSE;
   BenchUut7.station1Start := TRUE;
   BenchUut7.station2Complete := FALSE;
   BenchUut7.station3Complete := FALSE;
   BenchUut7.station4Complete := FALSE;
   BenchUut7.processSequence[1] := USINT#2;
   BenchUut7.processSequence[2] := USINT#2;
   BenchUut7.processSequence[3] := USINT#3;
   BenchUut7.processSequence[4] := USINT#3;
   BenchUut7.processSequence[5] := USINT#5;
   BenchUut7.processSequence[6] := USINT#0;
   BenchUut7.processSequence[7] := USINT#0;
   BenchUut7.processSequence[8] := USINT#0;
   TraceIn_processLength[149] := BenchUut7.processLength;
   TraceIn_sensor1[149] := BenchUut7.sensor1;
   TraceIn_sensor2[149] := BenchUut7.sensor2;
   TraceIn_sensor3[149] := BenchUut7.sensor3;
   TraceIn_sensor4[149] := BenchUut7.sensor4;
   TraceIn_sensor5[149] := BenchUut7.sensor5;
   TraceIn_station1Start[149] := BenchUut7.station1Start;
   TraceIn_station2Complete[149] := BenchUut7.station2Complete;
   TraceIn_station3Complete[149] := BenchUut7.station3Complete;
   TraceIn_station4Complete[149] := BenchUut7.station4Complete;
   TraceIn_processSequence_1[149] := BenchUut7.processSequence[1];
   TraceIn_processSequence_2[149] := BenchUut7.processSequence[2];
   TraceIn_processSequence_3[149] := BenchUut7.processSequence[3];
   TraceIn_processSequence_4[149] := BenchUut7.processSequence[4];
   TraceIn_processSequence_5[149] := BenchUut7.processSequence[5];
   TraceIn_processSequence_6[149] := BenchUut7.processSequence[6];
   TraceIn_processSequence_7[149] := BenchUut7.processSequence[7];
   TraceIn_processSequence_8[149] := BenchUut7.processSequence[8];
   BenchUut7();
   TraceOut_conveyorLeft[149] := BenchUut7.conveyorLeft;
   TraceOut_conveyorRight[149] := BenchUut7.conveyorRight;
   BenchCalls := BenchCalls + 1;
 150:
   BenchUut7.processLength := USINT#5;
   BenchUut7.sensor1 := FALSE;
   BenchUut7.sensor2 := TRUE;
   BenchUut7.sensor3 := FALSE;
   BenchUut7.sensor4 := FALSE;
   BenchUut7.sensor5 := FALSE;
   BenchUut7.station1Start := FALSE;
   BenchUut7.station2Complete := FALSE;
   BenchUut7.station3Complete := FALSE;
   BenchUut7.station4Complete := FALSE;
   BenchUut7.processSequence[1] := USINT#2;
   BenchUut7.processSequence[2] := USINT#2;
   BenchUut7.processSequence[3] := USINT#3;
   BenchUut7.processSequence[4] := USINT#3;
   BenchUut7.processSequence[5] := USINT#5;
   BenchUut7.processSequence[6] := USINT#0;
   BenchUut7.processSequence[7] := USINT#0;
   BenchUut7.processSequence[8] := USINT#0;
   TraceIn_processLength[150] := BenchUut7.processLength;
   TraceIn_sensor1[150] := BenchUut7.sensor1;
   TraceIn_sensor2[150] := BenchUut7.sensor2;
   TraceIn_sensor3[150] := BenchUut7.sensor3;
   TraceIn_sensor4[150] := BenchUut7.sensor4;
   TraceIn_sensor5[150] := BenchUut7.sensor5;
   TraceIn_station1Start[150] := BenchUut7.station1Start;
   TraceIn_station2Complete[150] := BenchUut7.station2Complete;
   TraceIn_station3Complete[150] := BenchUut7.station3Complete;
   TraceIn_station4Complete[150] := BenchUut7.station4Complete;
   TraceIn_processSequence_1[150] := BenchUut7.processSequence[1];
   TraceIn_processSequence_2[150] := BenchUut7.processSequence[2];
   TraceIn_processSequence_3[150] := BenchUut7.processSequence[3];
   TraceIn_processSequence_4[150] := BenchUut7.processSequence[4];
   TraceIn_processSequence_5[150] := BenchUut7.processSequence[5];
   TraceIn_processSequence_6[150] := BenchUut7.processSequence[6];
   TraceIn_processSequence_7[150] := BenchUut7.processSequence[7];
   TraceIn_processSequence_8[150] := BenchUut7.processSequence[8];
   BenchUut7();
   TraceOut_conveyorLeft[150] := BenchUut7.conveyorLeft;
   TraceOut_conveyorRight[150] := BenchUut7.conveyorRight;
   BenchCalls := BenchCalls + 1;
 151:
   BenchUut7.processLength := USINT#5;
   BenchUut7.sensor1 := FALSE;
   BenchUut7.sensor2 := TRUE;
   BenchUut7.sensor3 := FALSE;
   BenchUut7.sensor4 := FALSE;
   BenchUut7.sensor5 := FALSE;
   BenchUut7.station1Start := FALSE;
   BenchUut7.station2Complete := TRUE;
   BenchUut7.station3Complete := FALSE;
   BenchUut7.station4Complete := FALSE;
   BenchUut7.processSequence[1] := USINT#2;
   BenchUut7.processSequence[2] := USINT#2;
   BenchUut7.processSequence[3] := USINT#3;
   BenchUut7.processSequence[4] := USINT#3;
   BenchUut7.processSequence[5] := USINT#5;
   BenchUut7.processSequence[6] := USINT#0;
   BenchUut7.processSequence[7] := USINT#0;
   BenchUut7.processSequence[8] := USINT#0;
   TraceIn_processLength[151] := BenchUut7.processLength;
   TraceIn_sensor1[151] := BenchUut7.sensor1;
   TraceIn_sensor2[151] := BenchUut7.sensor2;
   TraceIn_sensor3[151] := BenchUut7.sensor3;
   TraceIn_sensor4[151] := BenchUut7.sensor4;
   TraceIn_sensor5[151] := BenchUut7.sensor5;
   TraceIn_station1Start[151] := BenchUut7.station1Start;
   TraceIn_station2Complete[151] := BenchUut7.station2Complete;
   TraceIn_station3Complete[151] := BenchUut7.station3Complete;
   TraceIn_station4Complete[151] := BenchUut7.station4Complete;
   TraceIn_processSequence_1[151] := BenchUut7.processSequence[1];
   TraceIn_processSequence_2[151] := BenchUut7.processSequence[2];
   TraceIn_processSequence_3[151] := BenchUut7.processSequence[3];
   TraceIn_processSequence_4[151] := BenchUut7.processSequence[4];
   TraceIn_processSequence_5[151] := BenchUut7.processSequence[5];
   TraceIn_processSequence_6[151] := BenchUut7.processSequence[6];
   TraceIn_processSequence_7[151] := BenchUut7.processSequence[7];
   TraceIn_processSequence_8[151] := BenchUut7.processSequence[8];
   BenchUut7();
   TraceOut_conveyorLeft[151] := BenchUut7.conveyorLeft;
   TraceOut_conveyorRight[151] := BenchUut7.conveyorRight;
   BenchCalls := BenchCalls + 1;
 152:
   BenchUut7.processLength := USINT#5;
   BenchUut7.sensor1 := FALSE;
   BenchUut7.sensor2 := TRUE;
   BenchUut7.sensor3 := FALSE;
   BenchUut7.sensor4 := FALSE;
   BenchUut7.sensor5 := FALSE;
   BenchUut7.station1Start := FALSE;
   BenchUut7.station2Complete := TRUE;
   BenchUut7.station3Complete := FALSE;
   BenchUut7.station4Complete := FALSE;
   BenchUut7.processSequence[1] := USINT#2;
   BenchUut7.processSequence[2] := USINT#2;
   BenchUut7.processSequence[3] := USINT#3;
   BenchUut7.processSequence[4] := USINT#3;
   BenchUut7.processSequence[5] := USINT#5;
   BenchUut7.processSequence[6] := USINT#0;
   BenchUut7.processSequence[7] := USINT#0;
   BenchUut7.processSequence[8] := USINT#0;
   TraceIn_processLength[152] := BenchUut7.processLength;
   TraceIn_sensor1[152] := BenchUut7.sensor1;
   TraceIn_sensor2[152] := BenchUut7.sensor2;
   TraceIn_sensor3[152] := BenchUut7.sensor3;
   TraceIn_sensor4[152] := BenchUut7.sensor4;
   TraceIn_sensor5[152] := BenchUut7.sensor5;
   TraceIn_station1Start[152] := BenchUut7.station1Start;
   TraceIn_station2Complete[152] := BenchUut7.station2Complete;
   TraceIn_station3Complete[152] := BenchUut7.station3Complete;
   TraceIn_station4Complete[152] := BenchUut7.station4Complete;
   TraceIn_processSequence_1[152] := BenchUut7.processSequence[1];
   TraceIn_processSequence_2[152] := BenchUut7.processSequence[2];
   TraceIn_processSequence_3[152] := BenchUut7.processSequence[3];
   TraceIn_processSequence_4[152] := BenchUut7.processSequence[4];
   TraceIn_processSequence_5[152] := BenchUut7.processSequence[5];
   TraceIn_processSequence_6[152] := BenchUut7.processSequence[6];
   TraceIn_processSequence_7[152] := BenchUut7.processSequence[7];
   TraceIn_processSequence_8[152] := BenchUut7.processSequence[8];
   BenchUut7();
   TraceOut_conveyorLeft[152] := BenchUut7.conveyorLeft;
   TraceOut_conveyorRight[152] := BenchUut7.conveyorRight;
   BenchCalls := BenchCalls + 1;
 153:
   BenchUut7.processLength := USINT#5;
   BenchUut7.sensor1 := FALSE;
   BenchUut7.sensor2 := TRUE;
   BenchUut7.sensor3 := FALSE;
   BenchUut7.sensor4 := FALSE;
   BenchUut7.sensor5 := FALSE;
   BenchUut7.station1Start := FALSE;
   BenchUut7.station2Complete := FALSE;
   BenchUut7.station3Complete := FALSE;
   BenchUut7.station4Complete := FALSE;
   BenchUut7.processSequence[1] := USINT#2;
   BenchUut7.processSequence[2] := USINT#2;
   BenchUut7.processSequence[3] := USINT#3;
   BenchUut7.processSequence[4] := USINT#3;
   BenchUut7.processSequence[5] := USINT#5;
   BenchUut7.processSequence[6] := USINT#0;
   BenchUut7.processSequence[7] := USINT#0;
   BenchUut7.processSequence[8] := USINT#0;
   TraceIn_processLength[153] := BenchUut7.processLength;
   TraceIn_sensor1[153] := BenchUut7.sensor1;
   TraceIn_sensor2[153] := BenchUut7.sensor2;
   TraceIn_sensor3[153] := BenchUut7.sensor3;
   TraceIn_sensor4[153] := BenchUut7.sensor4;
   TraceIn_sensor5[153] := BenchUut7.sensor5;
   TraceIn_station1Start[153] := BenchUut7.station1Start;
   TraceIn_station2Complete[153] := BenchUut7.station2Complete;
   TraceIn_station3Complete[153] := BenchUut7.station3Complete;
   TraceIn_station4Complete[153] := BenchUut7.station4Complete;
   TraceIn_processSequence_1[153] := BenchUut7.processSequence[1];
   TraceIn_processSequence_2[153] := BenchUut7.processSequence[2];
   TraceIn_processSequence_3[153] := BenchUut7.processSequence[3];
   TraceIn_processSequence_4[153] := BenchUut7.processSequence[4];
   TraceIn_processSequence_5[153] := BenchUut7.processSequence[5];
   TraceIn_processSequence_6[153] := BenchUut7.processSequence[6];
   TraceIn_processSequence_7[153] := BenchUut7.processSequence[7];
   TraceIn_processSequence_8[153] := BenchUut7.processSequence[8];
   BenchUut7();
   TraceOut_conveyorLeft[153] := BenchUut7.conveyorLeft;
   TraceOut_conveyorRight[153] := BenchUut7.conveyorRight;
   BenchCalls := BenchCalls + 1;
 154:
   BenchUut7.processLength := USINT#5;
   BenchUut7.sensor1 := FALSE;
   BenchUut7.sensor2 := TRUE;
   BenchUut7.sensor3 := FALSE;
   BenchUut7.sensor4 := FALSE;
   BenchUut7.sensor5 := FALSE;
   BenchUut7.station1Start := FALSE;
   BenchUut7.station2Complete := TRUE;
   BenchUut7.station3Complete := FALSE;
   BenchUut7.station4Complete := FALSE;
   BenchUut7.processSequence[1] := USINT#2;
   BenchUut7.processSequence[2] := USINT#2;
   BenchUut7.processSequence[3] := USINT#3;
   BenchUut7.processSequence[4] := USINT#3;
   BenchUut7.processSequence[5] := USINT#5;
   BenchUut7.processSequence[6] := USINT#0;
   BenchUut7.processSequence[7] := USINT#0;
   BenchUut7.processSequence[8] := USINT#0;
   TraceIn_processLength[154] := BenchUut7.processLength;
   TraceIn_sensor1[154] := BenchUut7.sensor1;
   TraceIn_sensor2[154] := BenchUut7.sensor2;
   TraceIn_sensor3[154] := BenchUut7.sensor3;
   TraceIn_sensor4[154] := BenchUut7.sensor4;
   TraceIn_sensor5[154] := BenchUut7.sensor5;
   TraceIn_station1Start[154] := BenchUut7.station1Start;
   TraceIn_station2Complete[154] := BenchUut7.station2Complete;
   TraceIn_station3Complete[154] := BenchUut7.station3Complete;
   TraceIn_station4Complete[154] := BenchUut7.station4Complete;
   TraceIn_processSequence_1[154] := BenchUut7.processSequence[1];
   TraceIn_processSequence_2[154] := BenchUut7.processSequence[2];
   TraceIn_processSequence_3[154] := BenchUut7.processSequence[3];
   TraceIn_processSequence_4[154] := BenchUut7.processSequence[4];
   TraceIn_processSequence_5[154] := BenchUut7.processSequence[5];
   TraceIn_processSequence_6[154] := BenchUut7.processSequence[6];
   TraceIn_processSequence_7[154] := BenchUut7.processSequence[7];
   TraceIn_processSequence_8[154] := BenchUut7.processSequence[8];
   BenchUut7();
   TraceOut_conveyorLeft[154] := BenchUut7.conveyorLeft;
   TraceOut_conveyorRight[154] := BenchUut7.conveyorRight;
   BenchCalls := BenchCalls + 1;
 155:
   BenchUut7.processLength := USINT#5;
   BenchUut7.sensor1 := FALSE;
   BenchUut7.sensor2 := FALSE;
   BenchUut7.sensor3 := TRUE;
   BenchUut7.sensor4 := FALSE;
   BenchUut7.sensor5 := FALSE;
   BenchUut7.station1Start := FALSE;
   BenchUut7.station2Complete := FALSE;
   BenchUut7.station3Complete := FALSE;
   BenchUut7.station4Complete := FALSE;
   BenchUut7.processSequence[1] := USINT#2;
   BenchUut7.processSequence[2] := USINT#2;
   BenchUut7.processSequence[3] := USINT#3;
   BenchUut7.processSequence[4] := USINT#3;
   BenchUut7.processSequence[5] := USINT#5;
   BenchUut7.processSequence[6] := USINT#0;
   BenchUut7.processSequence[7] := USINT#0;
   BenchUut7.processSequence[8] := USINT#0;
   TraceIn_processLength[155] := BenchUut7.processLength;
   TraceIn_sensor1[155] := BenchUut7.sensor1;
   TraceIn_sensor2[155] := BenchUut7.sensor2;
   TraceIn_sensor3[155] := BenchUut7.sensor3;
   TraceIn_sensor4[155] := BenchUut7.sensor4;
   TraceIn_sensor5[155] := BenchUut7.sensor5;
   TraceIn_station1Start[155] := BenchUut7.station1Start;
   TraceIn_station2Complete[155] := BenchUut7.station2Complete;
   TraceIn_station3Complete[155] := BenchUut7.station3Complete;
   TraceIn_station4Complete[155] := BenchUut7.station4Complete;
   TraceIn_processSequence_1[155] := BenchUut7.processSequence[1];
   TraceIn_processSequence_2[155] := BenchUut7.processSequence[2];
   TraceIn_processSequence_3[155] := BenchUut7.processSequence[3];
   TraceIn_processSequence_4[155] := BenchUut7.processSequence[4];
   TraceIn_processSequence_5[155] := BenchUut7.processSequence[5];
   TraceIn_processSequence_6[155] := BenchUut7.processSequence[6];
   TraceIn_processSequence_7[155] := BenchUut7.processSequence[7];
   TraceIn_processSequence_8[155] := BenchUut7.processSequence[8];
   BenchUut7();
   TraceOut_conveyorLeft[155] := BenchUut7.conveyorLeft;
   TraceOut_conveyorRight[155] := BenchUut7.conveyorRight;
   BenchCalls := BenchCalls + 1;
 156:
   BenchUut7.processLength := USINT#5;
   BenchUut7.sensor1 := FALSE;
   BenchUut7.sensor2 := FALSE;
   BenchUut7.sensor3 := TRUE;
   BenchUut7.sensor4 := FALSE;
   BenchUut7.sensor5 := FALSE;
   BenchUut7.station1Start := FALSE;
   BenchUut7.station2Complete := FALSE;
   BenchUut7.station3Complete := TRUE;
   BenchUut7.station4Complete := FALSE;
   BenchUut7.processSequence[1] := USINT#2;
   BenchUut7.processSequence[2] := USINT#2;
   BenchUut7.processSequence[3] := USINT#3;
   BenchUut7.processSequence[4] := USINT#3;
   BenchUut7.processSequence[5] := USINT#5;
   BenchUut7.processSequence[6] := USINT#0;
   BenchUut7.processSequence[7] := USINT#0;
   BenchUut7.processSequence[8] := USINT#0;
   TraceIn_processLength[156] := BenchUut7.processLength;
   TraceIn_sensor1[156] := BenchUut7.sensor1;
   TraceIn_sensor2[156] := BenchUut7.sensor2;
   TraceIn_sensor3[156] := BenchUut7.sensor3;
   TraceIn_sensor4[156] := BenchUut7.sensor4;
   TraceIn_sensor5[156] := BenchUut7.sensor5;
   TraceIn_station1Start[156] := BenchUut7.station1Start;
   TraceIn_station2Complete[156] := BenchUut7.station2Complete;
   TraceIn_station3Complete[156] := BenchUut7.station3Complete;
   TraceIn_station4Complete[156] := BenchUut7.station4Complete;
   TraceIn_processSequence_1[156] := BenchUut7.processSequence[1];
   TraceIn_processSequence_2[156] := BenchUut7.processSequence[2];
   TraceIn_processSequence_3[156] := BenchUut7.processSequence[3];
   TraceIn_processSequence_4[156] := BenchUut7.processSequence[4];
   TraceIn_processSequence_5[156] := BenchUut7.processSequence[5];
   TraceIn_processSequence_6[156] := BenchUut7.processSequence[6];
   TraceIn_processSequence_7[156] := BenchUut7.processSequence[7];
   TraceIn_processSequence_8[156] := BenchUut7.processSequence[8];
   BenchUut7();
   TraceOut_conveyorLeft[156] := BenchUut7.conveyorLeft;
   TraceOut_conveyorRight[156] := BenchUut7.conveyorRight;
   BenchCalls := BenchCalls + 1;
 157:
   BenchUut7.processLength := USINT#5;
   BenchUut7.sensor1 := FALSE;
   BenchUut7.sensor2 := FALSE;
   BenchUut7.sensor3 := TRUE;
   BenchUut7.sensor4 := FALSE;
   BenchUut7.sensor5 := FALSE;
   BenchUut7.station1Start := FALSE;
   BenchUut7.station2Complete := FALSE;
   BenchUut7.station3Complete := FALSE;
   BenchUut7.station4Complete := FALSE;
   BenchUut7.processSequence[1] := USINT#2;
   BenchUut7.processSequence[2] := USINT#2;
   BenchUut7.processSequence[3] := USINT#3;
   BenchUut7.processSequence[4] := USINT#3;
   BenchUut7.processSequence[5] := USINT#5;
   BenchUut7.processSequence[6] := USINT#0;
   BenchUut7.processSequence[7] := USINT#0;
   BenchUut7.processSequence[8] := USINT#0;
   TraceIn_processLength[157] := BenchUut7.processLength;
   TraceIn_sensor1[157] := BenchUut7.sensor1;
   TraceIn_sensor2[157] := BenchUut7.sensor2;
   TraceIn_sensor3[157] := BenchUut7.sensor3;
   TraceIn_sensor4[157] := BenchUut7.sensor4;
   TraceIn_sensor5[157] := BenchUut7.sensor5;
   TraceIn_station1Start[157] := BenchUut7.station1Start;
   TraceIn_station2Complete[157] := BenchUut7.station2Complete;
   TraceIn_station3Complete[157] := BenchUut7.station3Complete;
   TraceIn_station4Complete[157] := BenchUut7.station4Complete;
   TraceIn_processSequence_1[157] := BenchUut7.processSequence[1];
   TraceIn_processSequence_2[157] := BenchUut7.processSequence[2];
   TraceIn_processSequence_3[157] := BenchUut7.processSequence[3];
   TraceIn_processSequence_4[157] := BenchUut7.processSequence[4];
   TraceIn_processSequence_5[157] := BenchUut7.processSequence[5];
   TraceIn_processSequence_6[157] := BenchUut7.processSequence[6];
   TraceIn_processSequence_7[157] := BenchUut7.processSequence[7];
   TraceIn_processSequence_8[157] := BenchUut7.processSequence[8];
   BenchUut7();
   TraceOut_conveyorLeft[157] := BenchUut7.conveyorLeft;
   TraceOut_conveyorRight[157] := BenchUut7.conveyorRight;
   BenchCalls := BenchCalls + 1;
 158:
   BenchUut7.processLength := USINT#5;
   BenchUut7.sensor1 := FALSE;
   BenchUut7.sensor2 := FALSE;
   BenchUut7.sensor3 := TRUE;
   BenchUut7.sensor4 := FALSE;
   BenchUut7.sensor5 := FALSE;
   BenchUut7.station1Start := FALSE;
   BenchUut7.station2Complete := FALSE;
   BenchUut7.station3Complete := TRUE;
   BenchUut7.station4Complete := FALSE;
   BenchUut7.processSequence[1] := USINT#2;
   BenchUut7.processSequence[2] := USINT#2;
   BenchUut7.processSequence[3] := USINT#3;
   BenchUut7.processSequence[4] := USINT#3;
   BenchUut7.processSequence[5] := USINT#5;
   BenchUut7.processSequence[6] := USINT#0;
   BenchUut7.processSequence[7] := USINT#0;
   BenchUut7.processSequence[8] := USINT#0;
   TraceIn_processLength[158] := BenchUut7.processLength;
   TraceIn_sensor1[158] := BenchUut7.sensor1;
   TraceIn_sensor2[158] := BenchUut7.sensor2;
   TraceIn_sensor3[158] := BenchUut7.sensor3;
   TraceIn_sensor4[158] := BenchUut7.sensor4;
   TraceIn_sensor5[158] := BenchUut7.sensor5;
   TraceIn_station1Start[158] := BenchUut7.station1Start;
   TraceIn_station2Complete[158] := BenchUut7.station2Complete;
   TraceIn_station3Complete[158] := BenchUut7.station3Complete;
   TraceIn_station4Complete[158] := BenchUut7.station4Complete;
   TraceIn_processSequence_1[158] := BenchUut7.processSequence[1];
   TraceIn_processSequence_2[158] := BenchUut7.processSequence[2];
   TraceIn_processSequence_3[158] := BenchUut7.processSequence[3];
   TraceIn_processSequence_4[158] := BenchUut7.processSequence[4];
   TraceIn_processSequence_5[158] := BenchUut7.processSequence[5];
   TraceIn_processSequence_6[158] := BenchUut7.processSequence[6];
   TraceIn_processSequence_7[158] := BenchUut7.processSequence[7];
   TraceIn_processSequence_8[158] := BenchUut7.processSequence[8];
   BenchUut7();
   TraceOut_conveyorLeft[158] := BenchUut7.conveyorLeft;
   TraceOut_conveyorRight[158] := BenchUut7.conveyorRight;
   BenchCalls := BenchCalls + 1;
 159:
   BenchUut7.processLength := USINT#5;
   BenchUut7.sensor1 := FALSE;
   BenchUut7.sensor2 := FALSE;
   BenchUut7.sensor3 := FALSE;
   BenchUut7.sensor4 := FALSE;
   BenchUut7.sensor5 := TRUE;
   BenchUut7.station1Start := FALSE;
   BenchUut7.station2Complete := FALSE;
   BenchUut7.station3Complete := FALSE;
   BenchUut7.station4Complete := FALSE;
   BenchUut7.processSequence[1] := USINT#2;
   BenchUut7.processSequence[2] := USINT#2;
   BenchUut7.processSequence[3] := USINT#3;
   BenchUut7.processSequence[4] := USINT#3;
   BenchUut7.processSequence[5] := USINT#5;
   BenchUut7.processSequence[6] := USINT#0;
   BenchUut7.processSequence[7] := USINT#0;
   BenchUut7.processSequence[8] := USINT#0;
   TraceIn_processLength[159] := BenchUut7.processLength;
   TraceIn_sensor1[159] := BenchUut7.sensor1;
   TraceIn_sensor2[159] := BenchUut7.sensor2;
   TraceIn_sensor3[159] := BenchUut7.sensor3;
   TraceIn_sensor4[159] := BenchUut7.sensor4;
   TraceIn_sensor5[159] := BenchUut7.sensor5;
   TraceIn_station1Start[159] := BenchUut7.station1Start;
   TraceIn_station2Complete[159] := BenchUut7.station2Complete;
   TraceIn_station3Complete[159] := BenchUut7.station3Complete;
   TraceIn_station4Complete[159] := BenchUut7.station4Complete;
   TraceIn_processSequence_1[159] := BenchUut7.processSequence[1];
   TraceIn_processSequence_2[159] := BenchUut7.processSequence[2];
   TraceIn_processSequence_3[159] := BenchUut7.processSequence[3];
   TraceIn_processSequence_4[159] := BenchUut7.processSequence[4];
   TraceIn_processSequence_5[159] := BenchUut7.processSequence[5];
   TraceIn_processSequence_6[159] := BenchUut7.processSequence[6];
   TraceIn_processSequence_7[159] := BenchUut7.processSequence[7];
   TraceIn_processSequence_8[159] := BenchUut7.processSequence[8];
   BenchUut7();
   TraceOut_conveyorLeft[159] := BenchUut7.conveyorLeft;
   TraceOut_conveyorRight[159] := BenchUut7.conveyorRight;
   BenchCalls := BenchCalls + 1;
 END_CASE;
 BenchStep := BenchStep + 1;
 IF BenchStep >= 160 THEN BenchDone := TRUE; END_IF;
END_IF;
END_PROGRAM
